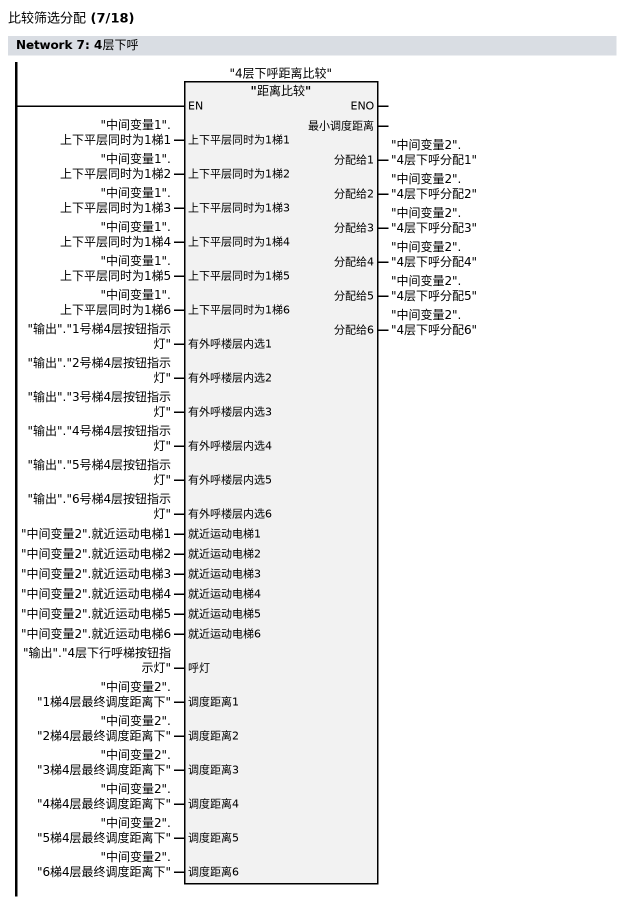
   RUNG wire#powerrail
      "4层下呼距离比较"(上下平层同时为1梯1 := "中间变量1".上下平层同时为1梯1, 上下平层同时为1梯2 := "中间变量1".上下平层同时为1梯2, 上下平层同时为1梯3 := "中间变量1".上下平层同时为1梯3, 上下平层同时为1梯4 := "中间变量1".上下平层同时为1梯4, 上下平层同时为1梯5 := "中间变量1".上下平层同时为1梯5, 上下平层同时为1梯6 := "中间变量1".上下平层同时为1梯6, 有外呼楼层内选1 := "输出"."1号梯4层按钮指示灯", 有外呼楼层内选2 := "输出"."2号梯4层按钮指示灯", 有外呼楼层内选3 := "输出"."3号梯4层按钮指示灯", 有外呼楼层内选4 := "输出"."4号梯4层按钮指示灯", 有外呼楼层内选5 := "输出"."5号梯4层按钮指示灯", 有外呼楼层内选6 := "输出"."6号梯4层按钮指示灯", 就近运动电梯1 := "中间变量2".就近运动电梯1, 就近运动电梯2 := "中间变量2".就近运动电梯2, 就近运动电梯3 := "中间变量2".就近运动电梯3, 就近运动电梯4 := "中间变量2".就近运动电梯4, 就近运动电梯5 := "中间变量2".就近运动电梯5, 就近运动电梯6 := "中间变量2".就近运动电梯6, 呼灯 := "输出"."4层下行呼梯按钮指示灯", 调度距离1 := "中间变量2"."1梯4层最终调度距离下", 调度距离2 := "中间变量2"."2梯4层最终调度距离下", 调度距离3 := "中间变量2"."3梯4层最终调度距离下", 调度距离4 := "中间变量2"."4梯4层最终调度距离下", 调度距离5 := "中间变量2"."5梯4层最终调度距离下", 调度距离6 := "中间变量2"."6梯4层最终调度距离下", 最小调度距离 =>, 分配给1 => "中间变量2"."4层下呼分配1", 分配给2 => "中间变量2"."4层下呼分配2", 分配给3 => "中间变量2"."4层下呼分配3", 分配给4 => "中间变量2"."4层下呼分配4", 分配给5 => "中间变量2"."4层下呼分配5", 分配给6 => "中间变量2"."4层下呼分配6")
   END_RUNG
   // the same network as SCL:
   "4层下呼距离比较"(上下平层同时为1梯1 := "中间变量1".上下平层同时为1梯1,   // "距离比较"
              上下平层同时为1梯2 := "中间变量1".上下平层同时为1梯2,
              上下平层同时为1梯3 := "中间变量1".上下平层同时为1梯3,
              上下平层同时为1梯4 := "中间变量1".上下平层同时为1梯4,
              上下平层同时为1梯5 := "中间变量1".上下平层同时为1梯5,
              上下平层同时为1梯6 := "中间变量1".上下平层同时为1梯6,
              有外呼楼层内选1 := "输出"."1号梯4层按钮指示灯",
              有外呼楼层内选2 := "输出"."2号梯4层按钮指示灯",
              有外呼楼层内选3 := "输出"."3号梯4层按钮指示灯",
              有外呼楼层内选4 := "输出"."4号梯4层按钮指示灯",
              有外呼楼层内选5 := "输出"."5号梯4层按钮指示灯",
              有外呼楼层内选6 := "输出"."6号梯4层按钮指示灯",
              就近运动电梯1 := "中间变量2".就近运动电梯1,
              就近运动电梯2 := "中间变量2".就近运动电梯2,
              就近运动电梯3 := "中间变量2".就近运动电梯3,
              就近运动电梯4 := "中间变量2".就近运动电梯4,
              就近运动电梯5 := "中间变量2".就近运动电梯5,
              就近运动电梯6 := "中间变量2".就近运动电梯6,
              呼灯 := "输出"."4层下行呼梯按钮指示灯",
              调度距离1 := "中间变量2"."1梯4层最终调度距离下",
              调度距离2 := "中间变量2"."2梯4层最终调度距离下",
              调度距离3 := "中间变量2"."3梯4层最终调度距离下",
              调度距离4 := "中间变量2"."4梯4层最终调度距离下",
              调度距离5 := "中间变量2"."5梯4层最终调度距离下",
              调度距离6 := "中间变量2"."6梯4层最终调度距离下",
              分配给1 => "中间变量2"."4层下呼分配1",
              分配给2 => "中间变量2"."4层下呼分配2",
              分配给3 => "中间变量2"."4层下呼分配3",
              分配给4 => "中间变量2"."4层下呼分配4",
              分配给5 => "中间变量2"."4层下呼分配5",
              分配给6 => "中间变量2"."4层下呼分配6");
END_REGION

REGION Network 8: 5层上呼
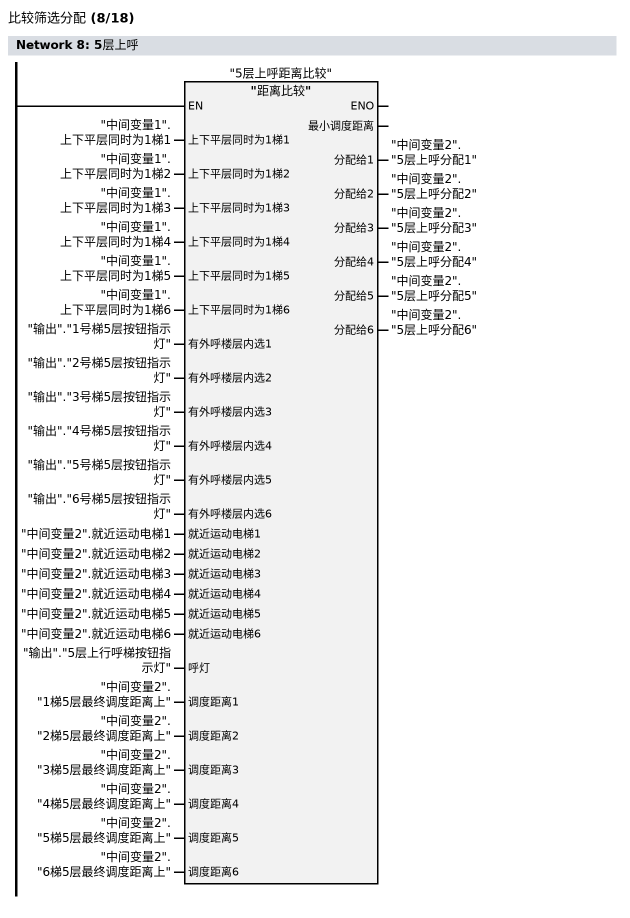
   RUNG wire#powerrail
      "5层上呼距离比较"(上下平层同时为1梯1 := "中间变量1".上下平层同时为1梯1, 上下平层同时为1梯2 := "中间变量1".上下平层同时为1梯2, 上下平层同时为1梯3 := "中间变量1".上下平层同时为1梯3, 上下平层同时为1梯4 := "中间变量1".上下平层同时为1梯4, 上下平层同时为1梯5 := "中间变量1".上下平层同时为1梯5, 上下平层同时为1梯6 := "中间变量1".上下平层同时为1梯6, 有外呼楼层内选1 := "输出"."1号梯5层按钮指示灯", 有外呼楼层内选2 := "输出"."2号梯5层按钮指示灯", 有外呼楼层内选3 := "输出"."3号梯5层按钮指示灯", 有外呼楼层内选4 := "输出"."4号梯5层按钮指示灯", 有外呼楼层内选5 := "输出"."5号梯5层按钮指示灯", 有外呼楼层内选6 := "输出"."6号梯5层按钮指示灯", 就近运动电梯1 := "中间变量2".就近运动电梯1, 就近运动电梯2 := "中间变量2".就近运动电梯2, 就近运动电梯3 := "中间变量2".就近运动电梯3, 就近运动电梯4 := "中间变量2".就近运动电梯4, 就近运动电梯5 := "中间变量2".就近运动电梯5, 就近运动电梯6 := "中间变量2".就近运动电梯6, 呼灯 := "输出"."5层上行呼梯按钮指示灯", 调度距离1 := "中间变量2"."1梯5层最终调度距离上", 调度距离2 := "中间变量2"."2梯5层最终调度距离上", 调度距离3 := "中间变量2"."3梯5层最终调度距离上", 调度距离4 := "中间变量2"."4梯5层最终调度距离上", 调度距离5 := "中间变量2"."5梯5层最终调度距离上", 调度距离6 := "中间变量2"."6梯5层最终调度距离上", 最小调度距离 =>, 分配给1 => "中间变量2"."5层上呼分配1", 分配给2 => "中间变量2"."5层上呼分配2", 分配给3 => "中间变量2"."5层上呼分配3", 分配给4 => "中间变量2"."5层上呼分配4", 分配给5 => "中间变量2"."5层上呼分配5", 分配给6 => "中间变量2"."5层上呼分配6")
   END_RUNG
   // the same network as SCL:
   "5层上呼距离比较"(上下平层同时为1梯1 := "中间变量1".上下平层同时为1梯1,   // "距离比较"
              上下平层同时为1梯2 := "中间变量1".上下平层同时为1梯2,
              上下平层同时为1梯3 := "中间变量1".上下平层同时为1梯3,
              上下平层同时为1梯4 := "中间变量1".上下平层同时为1梯4,
              上下平层同时为1梯5 := "中间变量1".上下平层同时为1梯5,
              上下平层同时为1梯6 := "中间变量1".上下平层同时为1梯6,
              有外呼楼层内选1 := "输出"."1号梯5层按钮指示灯",
              有外呼楼层内选2 := "输出"."2号梯5层按钮指示灯",
              有外呼楼层内选3 := "输出"."3号梯5层按钮指示灯",
              有外呼楼层内选4 := "输出"."4号梯5层按钮指示灯",
              有外呼楼层内选5 := "输出"."5号梯5层按钮指示灯",
              有外呼楼层内选6 := "输出"."6号梯5层按钮指示灯",
              就近运动电梯1 := "中间变量2".就近运动电梯1,
              就近运动电梯2 := "中间变量2".就近运动电梯2,
              就近运动电梯3 := "中间变量2".就近运动电梯3,
              就近运动电梯4 := "中间变量2".就近运动电梯4,
              就近运动电梯5 := "中间变量2".就近运动电梯5,
              就近运动电梯6 := "中间变量2".就近运动电梯6,
              呼灯 := "输出"."5层上行呼梯按钮指示灯",
              调度距离1 := "中间变量2"."1梯5层最终调度距离上",
              调度距离2 := "中间变量2"."2梯5层最终调度距离上",
              调度距离3 := "中间变量2"."3梯5层最终调度距离上",
              调度距离4 := "中间变量2"."4梯5层最终调度距离上",
              调度距离5 := "中间变量2"."5梯5层最终调度距离上",
              调度距离6 := "中间变量2"."6梯5层最终调度距离上",
              分配给1 => "中间变量2"."5层上呼分配1",
              分配给2 => "中间变量2"."5层上呼分配2",
              分配给3 => "中间变量2"."5层上呼分配3",
              分配给4 => "中间变量2"."5层上呼分配4",
              分配给5 => "中间变量2"."5层上呼分配5",
              分配给6 => "中间变量2"."5层上呼分配6");
END_REGION

REGION Network 9: 5层下呼
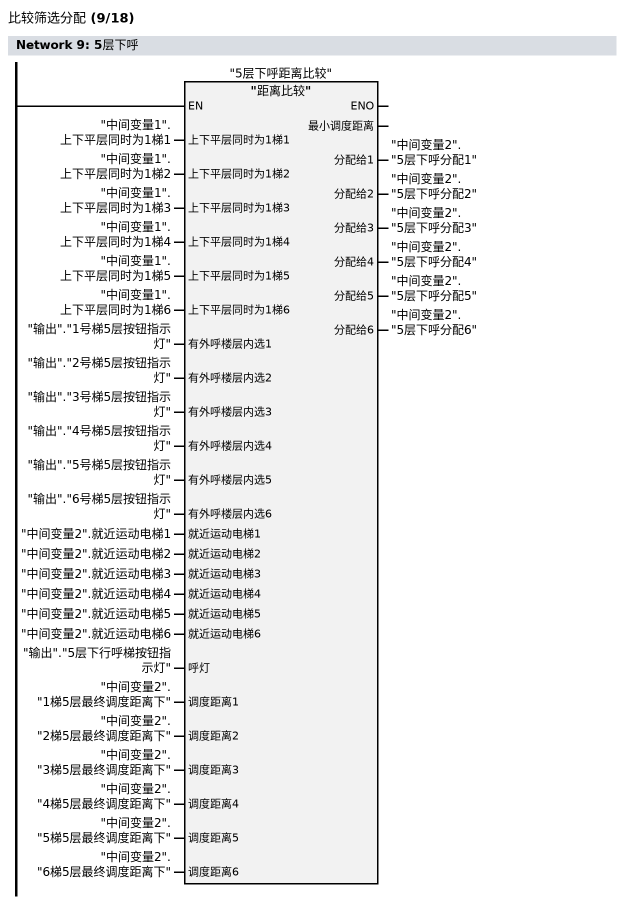
   RUNG wire#powerrail
      "5层下呼距离比较"(上下平层同时为1梯1 := "中间变量1".上下平层同时为1梯1, 上下平层同时为1梯2 := "中间变量1".上下平层同时为1梯2, 上下平层同时为1梯3 := "中间变量1".上下平层同时为1梯3, 上下平层同时为1梯4 := "中间变量1".上下平层同时为1梯4, 上下平层同时为1梯5 := "中间变量1".上下平层同时为1梯5, 上下平层同时为1梯6 := "中间变量1".上下平层同时为1梯6, 有外呼楼层内选1 := "输出"."1号梯5层按钮指示灯", 有外呼楼层内选2 := "输出"."2号梯5层按钮指示灯", 有外呼楼层内选3 := "输出"."3号梯5层按钮指示灯", 有外呼楼层内选4 := "输出"."4号梯5层按钮指示灯", 有外呼楼层内选5 := "输出"."5号梯5层按钮指示灯", 有外呼楼层内选6 := "输出"."6号梯5层按钮指示灯", 就近运动电梯1 := "中间变量2".就近运动电梯1, 就近运动电梯2 := "中间变量2".就近运动电梯2, 就近运动电梯3 := "中间变量2".就近运动电梯3, 就近运动电梯4 := "中间变量2".就近运动电梯4, 就近运动电梯5 := "中间变量2".就近运动电梯5, 就近运动电梯6 := "中间变量2".就近运动电梯6, 呼灯 := "输出"."5层下行呼梯按钮指示灯", 调度距离1 := "中间变量2"."1梯5层最终调度距离下", 调度距离2 := "中间变量2"."2梯5层最终调度距离下", 调度距离3 := "中间变量2"."3梯5层最终调度距离下", 调度距离4 := "中间变量2"."4梯5层最终调度距离下", 调度距离5 := "中间变量2"."5梯5层最终调度距离下", 调度距离6 := "中间变量2"."6梯5层最终调度距离下", 最小调度距离 =>, 分配给1 => "中间变量2"."5层下呼分配1", 分配给2 => "中间变量2"."5层下呼分配2", 分配给3 => "中间变量2"."5层下呼分配3", 分配给4 => "中间变量2"."5层下呼分配4", 分配给5 => "中间变量2"."5层下呼分配5", 分配给6 => "中间变量2"."5层下呼分配6")
   END_RUNG
   // the same network as SCL:
   "5层下呼距离比较"(上下平层同时为1梯1 := "中间变量1".上下平层同时为1梯1,   // "距离比较"
              上下平层同时为1梯2 := "中间变量1".上下平层同时为1梯2,
              上下平层同时为1梯3 := "中间变量1".上下平层同时为1梯3,
              上下平层同时为1梯4 := "中间变量1".上下平层同时为1梯4,
              上下平层同时为1梯5 := "中间变量1".上下平层同时为1梯5,
              上下平层同时为1梯6 := "中间变量1".上下平层同时为1梯6,
              有外呼楼层内选1 := "输出"."1号梯5层按钮指示灯",
              有外呼楼层内选2 := "输出"."2号梯5层按钮指示灯",
              有外呼楼层内选3 := "输出"."3号梯5层按钮指示灯",
              有外呼楼层内选4 := "输出"."4号梯5层按钮指示灯",
              有外呼楼层内选5 := "输出"."5号梯5层按钮指示灯",
              有外呼楼层内选6 := "输出"."6号梯5层按钮指示灯",
              就近运动电梯1 := "中间变量2".就近运动电梯1,
              就近运动电梯2 := "中间变量2".就近运动电梯2,
              就近运动电梯3 := "中间变量2".就近运动电梯3,
              就近运动电梯4 := "中间变量2".就近运动电梯4,
              就近运动电梯5 := "中间变量2".就近运动电梯5,
              就近运动电梯6 := "中间变量2".就近运动电梯6,
              呼灯 := "输出"."5层下行呼梯按钮指示灯",
              调度距离1 := "中间变量2"."1梯5层最终调度距离下",
              调度距离2 := "中间变量2"."2梯5层最终调度距离下",
              调度距离3 := "中间变量2"."3梯5层最终调度距离下",
              调度距离4 := "中间变量2"."4梯5层最终调度距离下",
              调度距离5 := "中间变量2"."5梯5层最终调度距离下",
              调度距离6 := "中间变量2"."6梯5层最终调度距离下",
              分配给1 => "中间变量2"."5层下呼分配1",
              分配给2 => "中间变量2"."5层下呼分配2",
              分配给3 => "中间变量2"."5层下呼分配3",
              分配给4 => "中间变量2"."5层下呼分配4",
              分配给5 => "中间变量2"."5层下呼分配5",
              分配给6 => "中间变量2"."5层下呼分配6");
END_REGION

REGION Network 10: 6层上呼
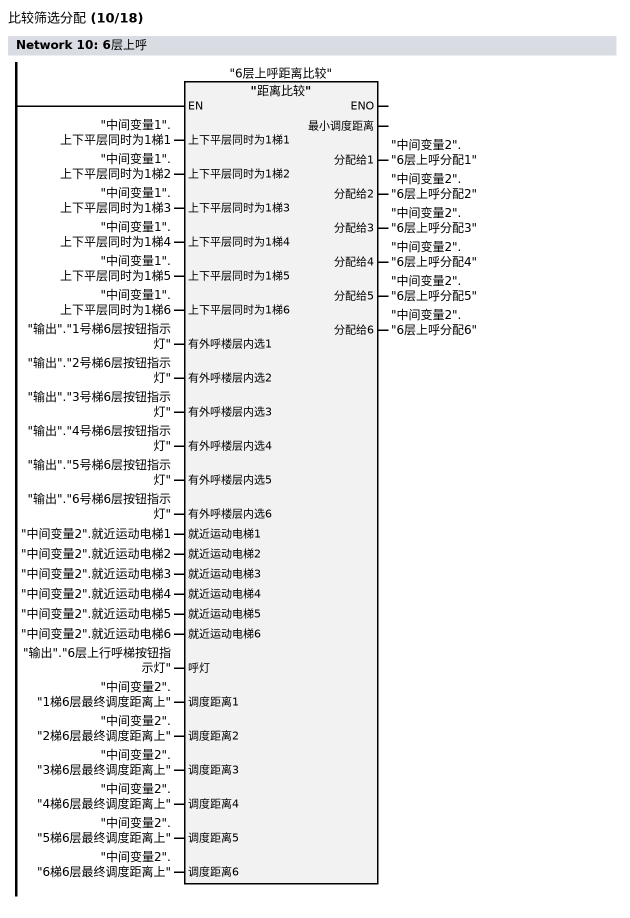
   RUNG wire#powerrail
      "6层上呼距离比较"(上下平层同时为1梯1 := "中间变量1".上下平层同时为1梯1, 上下平层同时为1梯2 := "中间变量1".上下平层同时为1梯2, 上下平层同时为1梯3 := "中间变量1".上下平层同时为1梯3, 上下平层同时为1梯4 := "中间变量1".上下平层同时为1梯4, 上下平层同时为1梯5 := "中间变量1".上下平层同时为1梯5, 上下平层同时为1梯6 := "中间变量1".上下平层同时为1梯6, 有外呼楼层内选1 := "输出"."1号梯6层按钮指示灯", 有外呼楼层内选2 := "输出"."2号梯6层按钮指示灯", 有外呼楼层内选3 := "输出"."3号梯6层按钮指示灯", 有外呼楼层内选4 := "输出"."4号梯6层按钮指示灯", 有外呼楼层内选5 := "输出"."5号梯6层按钮指示灯", 有外呼楼层内选6 := "输出"."6号梯6层按钮指示灯", 就近运动电梯1 := "中间变量2".就近运动电梯1, 就近运动电梯2 := "中间变量2".就近运动电梯2, 就近运动电梯3 := "中间变量2".就近运动电梯3, 就近运动电梯4 := "中间变量2".就近运动电梯4, 就近运动电梯5 := "中间变量2".就近运动电梯5, 就近运动电梯6 := "中间变量2".就近运动电梯6, 呼灯 := "输出"."6层上行呼梯按钮指示灯", 调度距离1 := "中间变量2"."1梯6层最终调度距离上", 调度距离2 := "中间变量2"."2梯6层最终调度距离上", 调度距离3 := "中间变量2"."3梯6层最终调度距离上", 调度距离4 := "中间变量2"."4梯6层最终调度距离上", 调度距离5 := "中间变量2"."5梯6层最终调度距离上", 调度距离6 := "中间变量2"."6梯6层最终调度距离上", 最小调度距离 =>, 分配给1 => "中间变量2"."6层上呼分配1", 分配给2 => "中间变量2"."6层上呼分配2", 分配给3 => "中间变量2"."6层上呼分配3", 分配给4 => "中间变量2"."6层上呼分配4", 分配给5 => "中间变量2"."6层上呼分配5", 分配给6 => "中间变量2"."6层上呼分配6")
   END_RUNG
   // the same network as SCL:
   "6层上呼距离比较"(上下平层同时为1梯1 := "中间变量1".上下平层同时为1梯1,   // "距离比较"
              上下平层同时为1梯2 := "中间变量1".上下平层同时为1梯2,
              上下平层同时为1梯3 := "中间变量1".上下平层同时为1梯3,
              上下平层同时为1梯4 := "中间变量1".上下平层同时为1梯4,
              上下平层同时为1梯5 := "中间变量1".上下平层同时为1梯5,
              上下平层同时为1梯6 := "中间变量1".上下平层同时为1梯6,
              有外呼楼层内选1 := "输出"."1号梯6层按钮指示灯",
              有外呼楼层内选2 := "输出"."2号梯6层按钮指示灯",
              有外呼楼层内选3 := "输出"."3号梯6层按钮指示灯",
              有外呼楼层内选4 := "输出"."4号梯6层按钮指示灯",
              有外呼楼层内选5 := "输出"."5号梯6层按钮指示灯",
              有外呼楼层内选6 := "输出"."6号梯6层按钮指示灯",
              就近运动电梯1 := "中间变量2".就近运动电梯1,
              就近运动电梯2 := "中间变量2".就近运动电梯2,
              就近运动电梯3 := "中间变量2".就近运动电梯3,
              就近运动电梯4 := "中间变量2".就近运动电梯4,
              就近运动电梯5 := "中间变量2".就近运动电梯5,
              就近运动电梯6 := "中间变量2".就近运动电梯6,
              呼灯 := "输出"."6层上行呼梯按钮指示灯",
              调度距离1 := "中间变量2"."1梯6层最终调度距离上",
              调度距离2 := "中间变量2"."2梯6层最终调度距离上",
              调度距离3 := "中间变量2"."3梯6层最终调度距离上",
              调度距离4 := "中间变量2"."4梯6层最终调度距离上",
              调度距离5 := "中间变量2"."5梯6层最终调度距离上",
              调度距离6 := "中间变量2"."6梯6层最终调度距离上",
              分配给1 => "中间变量2"."6层上呼分配1",
              分配给2 => "中间变量2"."6层上呼分配2",
              分配给3 => "中间变量2"."6层上呼分配3",
              分配给4 => "中间变量2"."6层上呼分配4",
              分配给5 => "中间变量2"."6层上呼分配5",
              分配给6 => "中间变量2"."6层上呼分配6");
END_REGION

REGION Network 11: 6层下呼
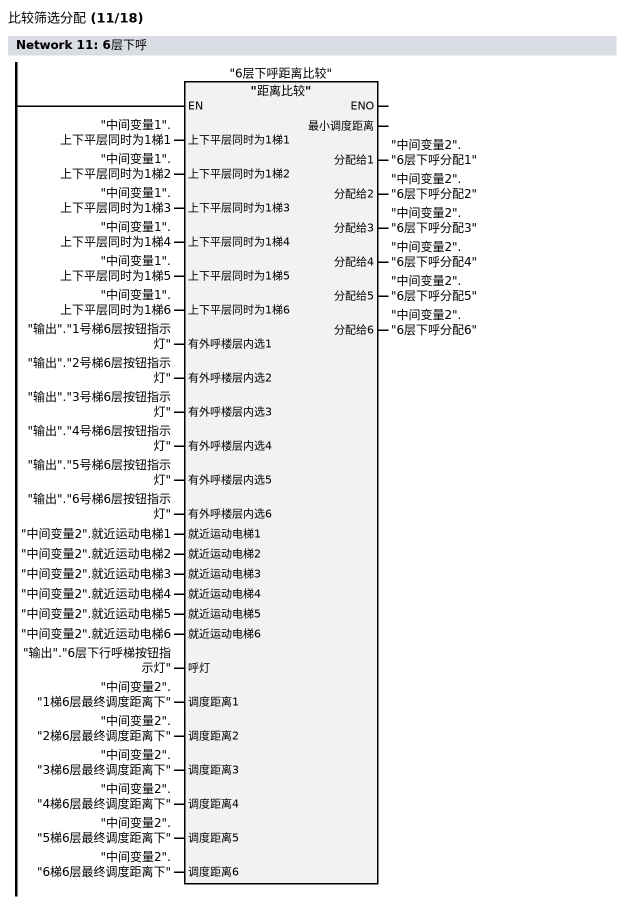
   RUNG wire#powerrail
      "6层下呼距离比较"(上下平层同时为1梯1 := "中间变量1".上下平层同时为1梯1, 上下平层同时为1梯2 := "中间变量1".上下平层同时为1梯2, 上下平层同时为1梯3 := "中间变量1".上下平层同时为1梯3, 上下平层同时为1梯4 := "中间变量1".上下平层同时为1梯4, 上下平层同时为1梯5 := "中间变量1".上下平层同时为1梯5, 上下平层同时为1梯6 := "中间变量1".上下平层同时为1梯6, 有外呼楼层内选1 := "输出"."1号梯6层按钮指示灯", 有外呼楼层内选2 := "输出"."2号梯6层按钮指示灯", 有外呼楼层内选3 := "输出"."3号梯6层按钮指示灯", 有外呼楼层内选4 := "输出"."4号梯6层按钮指示灯", 有外呼楼层内选5 := "输出"."5号梯6层按钮指示灯", 有外呼楼层内选6 := "输出"."6号梯6层按钮指示灯", 就近运动电梯1 := "中间变量2".就近运动电梯1, 就近运动电梯2 := "中间变量2".就近运动电梯2, 就近运动电梯3 := "中间变量2".就近运动电梯3, 就近运动电梯4 := "中间变量2".就近运动电梯4, 就近运动电梯5 := "中间变量2".就近运动电梯5, 就近运动电梯6 := "中间变量2".就近运动电梯6, 呼灯 := "输出"."6层下行呼梯按钮指示灯", 调度距离1 := "中间变量2"."1梯6层最终调度距离下", 调度距离2 := "中间变量2"."2梯6层最终调度距离下", 调度距离3 := "中间变量2"."3梯6层最终调度距离下", 调度距离4 := "中间变量2"."4梯6层最终调度距离下", 调度距离5 := "中间变量2"."5梯6层最终调度距离下", 调度距离6 := "中间变量2"."6梯6层最终调度距离下", 最小调度距离 =>, 分配给1 => "中间变量2"."6层下呼分配1", 分配给2 => "中间变量2"."6层下呼分配2", 分配给3 => "中间变量2"."6层下呼分配3", 分配给4 => "中间变量2"."6层下呼分配4", 分配给5 => "中间变量2"."6层下呼分配5", 分配给6 => "中间变量2"."6层下呼分配6")
   END_RUNG
   // the same network as SCL:
   "6层下呼距离比较"(上下平层同时为1梯1 := "中间变量1".上下平层同时为1梯1,   // "距离比较"
              上下平层同时为1梯2 := "中间变量1".上下平层同时为1梯2,
              上下平层同时为1梯3 := "中间变量1".上下平层同时为1梯3,
              上下平层同时为1梯4 := "中间变量1".上下平层同时为1梯4,
              上下平层同时为1梯5 := "中间变量1".上下平层同时为1梯5,
              上下平层同时为1梯6 := "中间变量1".上下平层同时为1梯6,
              有外呼楼层内选1 := "输出"."1号梯6层按钮指示灯",
              有外呼楼层内选2 := "输出"."2号梯6层按钮指示灯",
              有外呼楼层内选3 := "输出"."3号梯6层按钮指示灯",
              有外呼楼层内选4 := "输出"."4号梯6层按钮指示灯",
              有外呼楼层内选5 := "输出"."5号梯6层按钮指示灯",
              有外呼楼层内选6 := "输出"."6号梯6层按钮指示灯",
              就近运动电梯1 := "中间变量2".就近运动电梯1,
              就近运动电梯2 := "中间变量2".就近运动电梯2,
              就近运动电梯3 := "中间变量2".就近运动电梯3,
              就近运动电梯4 := "中间变量2".就近运动电梯4,
              就近运动电梯5 := "中间变量2".就近运动电梯5,
              就近运动电梯6 := "中间变量2".就近运动电梯6,
              呼灯 := "输出"."6层下行呼梯按钮指示灯",
              调度距离1 := "中间变量2"."1梯6层最终调度距离下",
              调度距离2 := "中间变量2"."2梯6层最终调度距离下",
              调度距离3 := "中间变量2"."3梯6层最终调度距离下",
              调度距离4 := "中间变量2"."4梯6层最终调度距离下",
              调度距离5 := "中间变量2"."5梯6层最终调度距离下",
              调度距离6 := "中间变量2"."6梯6层最终调度距离下",
              分配给1 => "中间变量2"."6层下呼分配1",
              分配给2 => "中间变量2"."6层下呼分配2",
              分配给3 => "中间变量2"."6层下呼分配3",
              分配给4 => "中间变量2"."6层下呼分配4",
              分配给5 => "中间变量2"."6层下呼分配5",
              分配给6 => "中间变量2"."6层下呼分配6");
END_REGION

REGION Network 12: 7层上呼
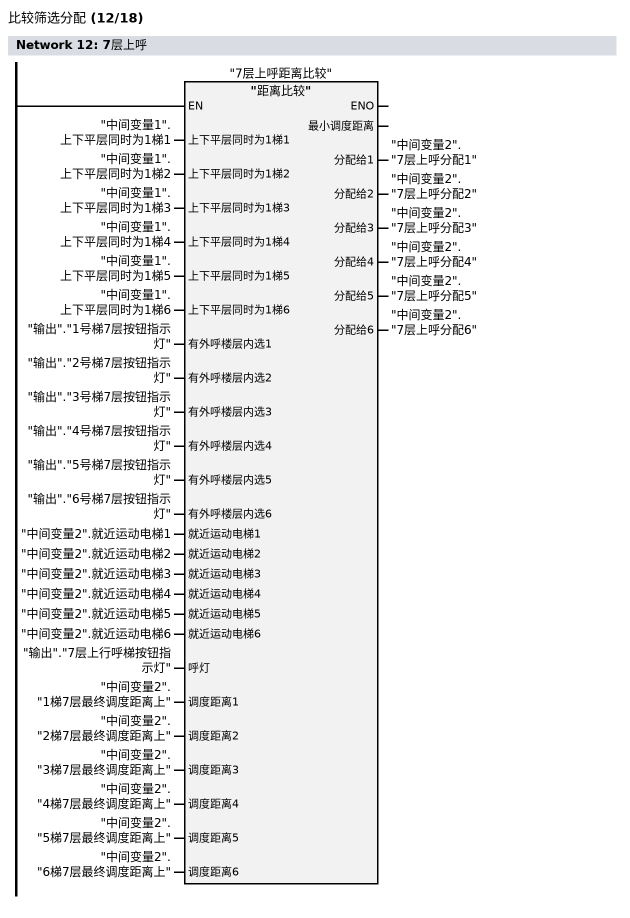
   RUNG wire#powerrail
      "7层上呼距离比较"(上下平层同时为1梯1 := "中间变量1".上下平层同时为1梯1, 上下平层同时为1梯2 := "中间变量1".上下平层同时为1梯2, 上下平层同时为1梯3 := "中间变量1".上下平层同时为1梯3, 上下平层同时为1梯4 := "中间变量1".上下平层同时为1梯4, 上下平层同时为1梯5 := "中间变量1".上下平层同时为1梯5, 上下平层同时为1梯6 := "中间变量1".上下平层同时为1梯6, 有外呼楼层内选1 := "输出"."1号梯7层按钮指示灯", 有外呼楼层内选2 := "输出"."2号梯7层按钮指示灯", 有外呼楼层内选3 := "输出"."3号梯7层按钮指示灯", 有外呼楼层内选4 := "输出"."4号梯7层按钮指示灯", 有外呼楼层内选5 := "输出"."5号梯7层按钮指示灯", 有外呼楼层内选6 := "输出"."6号梯7层按钮指示灯", 就近运动电梯1 := "中间变量2".就近运动电梯1, 就近运动电梯2 := "中间变量2".就近运动电梯2, 就近运动电梯3 := "中间变量2".就近运动电梯3, 就近运动电梯4 := "中间变量2".就近运动电梯4, 就近运动电梯5 := "中间变量2".就近运动电梯5, 就近运动电梯6 := "中间变量2".就近运动电梯6, 呼灯 := "输出"."7层上行呼梯按钮指示灯", 调度距离1 := "中间变量2"."1梯7层最终调度距离上", 调度距离2 := "中间变量2"."2梯7层最终调度距离上", 调度距离3 := "中间变量2"."3梯7层最终调度距离上", 调度距离4 := "中间变量2"."4梯7层最终调度距离上", 调度距离5 := "中间变量2"."5梯7层最终调度距离上", 调度距离6 := "中间变量2"."6梯7层最终调度距离上", 最小调度距离 =>, 分配给1 => "中间变量2"."7层上呼分配1", 分配给2 => "中间变量2"."7层上呼分配2", 分配给3 => "中间变量2"."7层上呼分配3", 分配给4 => "中间变量2"."7层上呼分配4", 分配给5 => "中间变量2"."7层上呼分配5", 分配给6 => "中间变量2"."7层上呼分配6")
   END_RUNG
   // the same network as SCL:
   "7层上呼距离比较"(上下平层同时为1梯1 := "中间变量1".上下平层同时为1梯1,   // "距离比较"
              上下平层同时为1梯2 := "中间变量1".上下平层同时为1梯2,
              上下平层同时为1梯3 := "中间变量1".上下平层同时为1梯3,
              上下平层同时为1梯4 := "中间变量1".上下平层同时为1梯4,
              上下平层同时为1梯5 := "中间变量1".上下平层同时为1梯5,
              上下平层同时为1梯6 := "中间变量1".上下平层同时为1梯6,
              有外呼楼层内选1 := "输出"."1号梯7层按钮指示灯",
              有外呼楼层内选2 := "输出"."2号梯7层按钮指示灯",
              有外呼楼层内选3 := "输出"."3号梯7层按钮指示灯",
              有外呼楼层内选4 := "输出"."4号梯7层按钮指示灯",
              有外呼楼层内选5 := "输出"."5号梯7层按钮指示灯",
              有外呼楼层内选6 := "输出"."6号梯7层按钮指示灯",
              就近运动电梯1 := "中间变量2".就近运动电梯1,
              就近运动电梯2 := "中间变量2".就近运动电梯2,
              就近运动电梯3 := "中间变量2".就近运动电梯3,
              就近运动电梯4 := "中间变量2".就近运动电梯4,
              就近运动电梯5 := "中间变量2".就近运动电梯5,
              就近运动电梯6 := "中间变量2".就近运动电梯6,
              呼灯 := "输出"."7层上行呼梯按钮指示灯",
              调度距离1 := "中间变量2"."1梯7层最终调度距离上",
              调度距离2 := "中间变量2"."2梯7层最终调度距离上",
              调度距离3 := "中间变量2"."3梯7层最终调度距离上",
              调度距离4 := "中间变量2"."4梯7层最终调度距离上",
              调度距离5 := "中间变量2"."5梯7层最终调度距离上",
              调度距离6 := "中间变量2"."6梯7层最终调度距离上",
              分配给1 => "中间变量2"."7层上呼分配1",
              分配给2 => "中间变量2"."7层上呼分配2",
              分配给3 => "中间变量2"."7层上呼分配3",
              分配给4 => "中间变量2"."7层上呼分配4",
              分配给5 => "中间变量2"."7层上呼分配5",
              分配给6 => "中间变量2"."7层上呼分配6");
END_REGION

REGION Network 13: 7层下呼
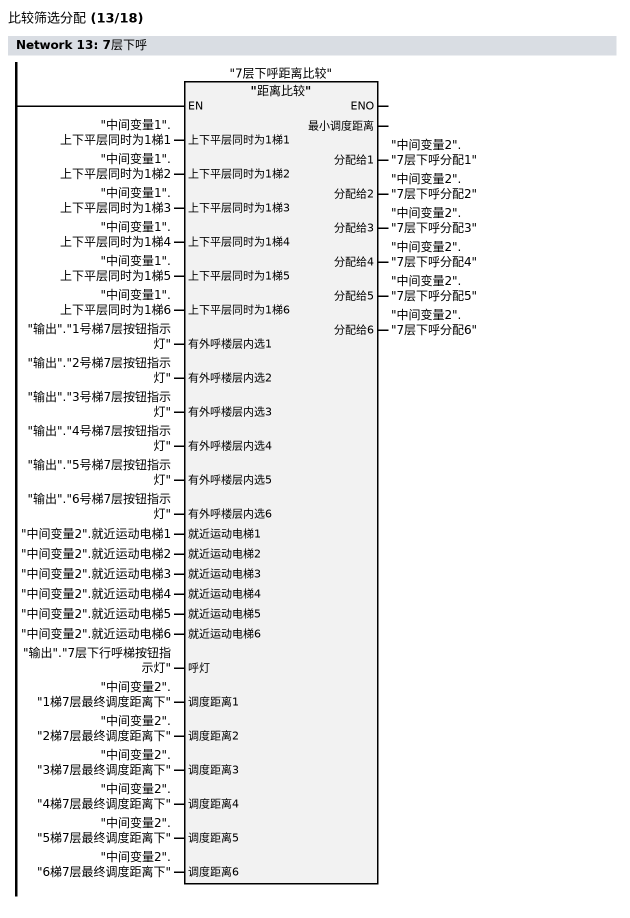
   RUNG wire#powerrail
      "7层下呼距离比较"(上下平层同时为1梯1 := "中间变量1".上下平层同时为1梯1, 上下平层同时为1梯2 := "中间变量1".上下平层同时为1梯2, 上下平层同时为1梯3 := "中间变量1".上下平层同时为1梯3, 上下平层同时为1梯4 := "中间变量1".上下平层同时为1梯4, 上下平层同时为1梯5 := "中间变量1".上下平层同时为1梯5, 上下平层同时为1梯6 := "中间变量1".上下平层同时为1梯6, 有外呼楼层内选1 := "输出"."1号梯7层按钮指示灯", 有外呼楼层内选2 := "输出"."2号梯7层按钮指示灯", 有外呼楼层内选3 := "输出"."3号梯7层按钮指示灯", 有外呼楼层内选4 := "输出"."4号梯7层按钮指示灯", 有外呼楼层内选5 := "输出"."5号梯7层按钮指示灯", 有外呼楼层内选6 := "输出"."6号梯7层按钮指示灯", 就近运动电梯1 := "中间变量2".就近运动电梯1, 就近运动电梯2 := "中间变量2".就近运动电梯2, 就近运动电梯3 := "中间变量2".就近运动电梯3, 就近运动电梯4 := "中间变量2".就近运动电梯4, 就近运动电梯5 := "中间变量2".就近运动电梯5, 就近运动电梯6 := "中间变量2".就近运动电梯6, 呼灯 := "输出"."7层下行呼梯按钮指示灯", 调度距离1 := "中间变量2"."1梯7层最终调度距离下", 调度距离2 := "中间变量2"."2梯7层最终调度距离下", 调度距离3 := "中间变量2"."3梯7层最终调度距离下", 调度距离4 := "中间变量2"."4梯7层最终调度距离下", 调度距离5 := "中间变量2"."5梯7层最终调度距离下", 调度距离6 := "中间变量2"."6梯7层最终调度距离下", 最小调度距离 =>, 分配给1 => "中间变量2"."7层下呼分配1", 分配给2 => "中间变量2"."7层下呼分配2", 分配给3 => "中间变量2"."7层下呼分配3", 分配给4 => "中间变量2"."7层下呼分配4", 分配给5 => "中间变量2"."7层下呼分配5", 分配给6 => "中间变量2"."7层下呼分配6")
   END_RUNG
   // the same network as SCL:
   "7层下呼距离比较"(上下平层同时为1梯1 := "中间变量1".上下平层同时为1梯1,   // "距离比较"
              上下平层同时为1梯2 := "中间变量1".上下平层同时为1梯2,
              上下平层同时为1梯3 := "中间变量1".上下平层同时为1梯3,
              上下平层同时为1梯4 := "中间变量1".上下平层同时为1梯4,
              上下平层同时为1梯5 := "中间变量1".上下平层同时为1梯5,
              上下平层同时为1梯6 := "中间变量1".上下平层同时为1梯6,
              有外呼楼层内选1 := "输出"."1号梯7层按钮指示灯",
              有外呼楼层内选2 := "输出"."2号梯7层按钮指示灯",
              有外呼楼层内选3 := "输出"."3号梯7层按钮指示灯",
              有外呼楼层内选4 := "输出"."4号梯7层按钮指示灯",
              有外呼楼层内选5 := "输出"."5号梯7层按钮指示灯",
              有外呼楼层内选6 := "输出"."6号梯7层按钮指示灯",
              就近运动电梯1 := "中间变量2".就近运动电梯1,
              就近运动电梯2 := "中间变量2".就近运动电梯2,
              就近运动电梯3 := "中间变量2".就近运动电梯3,
              就近运动电梯4 := "中间变量2".就近运动电梯4,
              就近运动电梯5 := "中间变量2".就近运动电梯5,
              就近运动电梯6 := "中间变量2".就近运动电梯6,
              呼灯 := "输出"."7层下行呼梯按钮指示灯",
              调度距离1 := "中间变量2"."1梯7层最终调度距离下",
              调度距离2 := "中间变量2"."2梯7层最终调度距离下",
              调度距离3 := "中间变量2"."3梯7层最终调度距离下",
              调度距离4 := "中间变量2"."4梯7层最终调度距离下",
              调度距离5 := "中间变量2"."5梯7层最终调度距离下",
              调度距离6 := "中间变量2"."6梯7层最终调度距离下",
              分配给1 => "中间变量2"."7层下呼分配1",
              分配给2 => "中间变量2"."7层下呼分配2",
              分配给3 => "中间变量2"."7层下呼分配3",
              分配给4 => "中间变量2"."7层下呼分配4",
              分配给5 => "中间变量2"."7层下呼分配5",
              分配给6 => "中间变量2"."7层下呼分配6");
END_REGION

REGION Network 14: 8层上呼
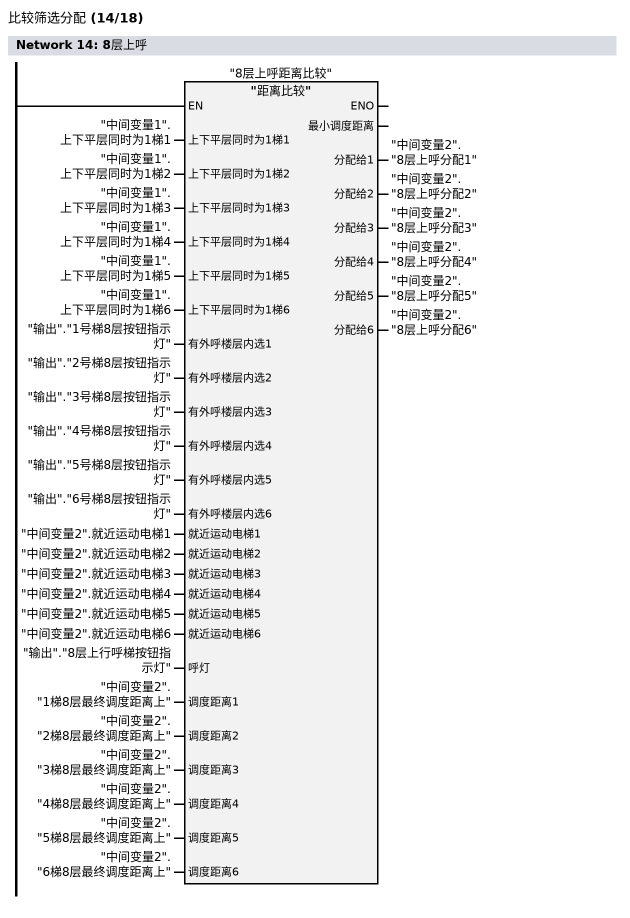
   RUNG wire#powerrail
      "8层上呼距离比较"(上下平层同时为1梯1 := "中间变量1".上下平层同时为1梯1, 上下平层同时为1梯2 := "中间变量1".上下平层同时为1梯2, 上下平层同时为1梯3 := "中间变量1".上下平层同时为1梯3, 上下平层同时为1梯4 := "中间变量1".上下平层同时为1梯4, 上下平层同时为1梯5 := "中间变量1".上下平层同时为1梯5, 上下平层同时为1梯6 := "中间变量1".上下平层同时为1梯6, 有外呼楼层内选1 := "输出"."1号梯8层按钮指示灯", 有外呼楼层内选2 := "输出"."2号梯8层按钮指示灯", 有外呼楼层内选3 := "输出"."3号梯8层按钮指示灯", 有外呼楼层内选4 := "输出"."4号梯8层按钮指示灯", 有外呼楼层内选5 := "输出"."5号梯8层按钮指示灯", 有外呼楼层内选6 := "输出"."6号梯8层按钮指示灯", 就近运动电梯1 := "中间变量2".就近运动电梯1, 就近运动电梯2 := "中间变量2".就近运动电梯2, 就近运动电梯3 := "中间变量2".就近运动电梯3, 就近运动电梯4 := "中间变量2".就近运动电梯4, 就近运动电梯5 := "中间变量2".就近运动电梯5, 就近运动电梯6 := "中间变量2".就近运动电梯6, 呼灯 := "输出"."8层上行呼梯按钮指示灯", 调度距离1 := "中间变量2"."1梯8层最终调度距离上", 调度距离2 := "中间变量2"."2梯8层最终调度距离上", 调度距离3 := "中间变量2"."3梯8层最终调度距离上", 调度距离4 := "中间变量2"."4梯8层最终调度距离上", 调度距离5 := "中间变量2"."5梯8层最终调度距离上", 调度距离6 := "中间变量2"."6梯8层最终调度距离上", 最小调度距离 =>, 分配给1 => "中间变量2"."8层上呼分配1", 分配给2 => "中间变量2"."8层上呼分配2", 分配给3 => "中间变量2"."8层上呼分配3", 分配给4 => "中间变量2"."8层上呼分配4", 分配给5 => "中间变量2"."8层上呼分配5", 分配给6 => "中间变量2"."8层上呼分配6")
   END_RUNG
   // the same network as SCL:
   "8层上呼距离比较"(上下平层同时为1梯1 := "中间变量1".上下平层同时为1梯1,   // "距离比较"
              上下平层同时为1梯2 := "中间变量1".上下平层同时为1梯2,
              上下平层同时为1梯3 := "中间变量1".上下平层同时为1梯3,
              上下平层同时为1梯4 := "中间变量1".上下平层同时为1梯4,
              上下平层同时为1梯5 := "中间变量1".上下平层同时为1梯5,
              上下平层同时为1梯6 := "中间变量1".上下平层同时为1梯6,
              有外呼楼层内选1 := "输出"."1号梯8层按钮指示灯",
              有外呼楼层内选2 := "输出"."2号梯8层按钮指示灯",
              有外呼楼层内选3 := "输出"."3号梯8层按钮指示灯",
              有外呼楼层内选4 := "输出"."4号梯8层按钮指示灯",
              有外呼楼层内选5 := "输出"."5号梯8层按钮指示灯",
              有外呼楼层内选6 := "输出"."6号梯8层按钮指示灯",
              就近运动电梯1 := "中间变量2".就近运动电梯1,
              就近运动电梯2 := "中间变量2".就近运动电梯2,
              就近运动电梯3 := "中间变量2".就近运动电梯3,
              就近运动电梯4 := "中间变量2".就近运动电梯4,
              就近运动电梯5 := "中间变量2".就近运动电梯5,
              就近运动电梯6 := "中间变量2".就近运动电梯6,
              呼灯 := "输出"."8层上行呼梯按钮指示灯",
              调度距离1 := "中间变量2"."1梯8层最终调度距离上",
              调度距离2 := "中间变量2"."2梯8层最终调度距离上",
              调度距离3 := "中间变量2"."3梯8层最终调度距离上",
              调度距离4 := "中间变量2"."4梯8层最终调度距离上",
              调度距离5 := "中间变量2"."5梯8层最终调度距离上",
              调度距离6 := "中间变量2"."6梯8层最终调度距离上",
              分配给1 => "中间变量2"."8层上呼分配1",
              分配给2 => "中间变量2"."8层上呼分配2",
              分配给3 => "中间变量2"."8层上呼分配3",
              分配给4 => "中间变量2"."8层上呼分配4",
              分配给5 => "中间变量2"."8层上呼分配5",
              分配给6 => "中间变量2"."8层上呼分配6");
END_REGION

REGION Network 15: 8层下呼
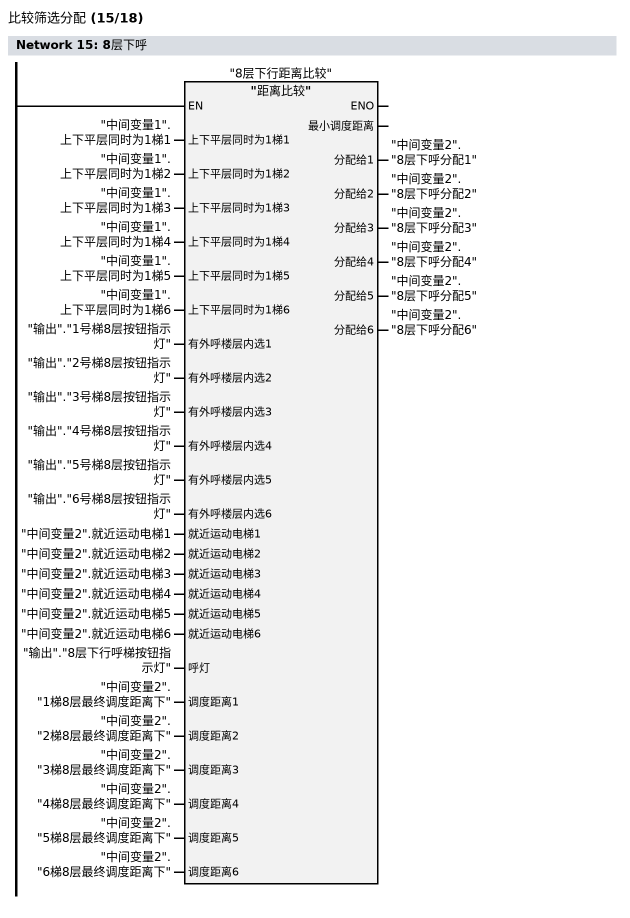
   RUNG wire#powerrail
      "8层下行距离比较"(上下平层同时为1梯1 := "中间变量1".上下平层同时为1梯1, 上下平层同时为1梯2 := "中间变量1".上下平层同时为1梯2, 上下平层同时为1梯3 := "中间变量1".上下平层同时为1梯3, 上下平层同时为1梯4 := "中间变量1".上下平层同时为1梯4, 上下平层同时为1梯5 := "中间变量1".上下平层同时为1梯5, 上下平层同时为1梯6 := "中间变量1".上下平层同时为1梯6, 有外呼楼层内选1 := "输出"."1号梯8层按钮指示灯", 有外呼楼层内选2 := "输出"."2号梯8层按钮指示灯", 有外呼楼层内选3 := "输出"."3号梯8层按钮指示灯", 有外呼楼层内选4 := "输出"."4号梯8层按钮指示灯", 有外呼楼层内选5 := "输出"."5号梯8层按钮指示灯", 有外呼楼层内选6 := "输出"."6号梯8层按钮指示灯", 就近运动电梯1 := "中间变量2".就近运动电梯1, 就近运动电梯2 := "中间变量2".就近运动电梯2, 就近运动电梯3 := "中间变量2".就近运动电梯3, 就近运动电梯4 := "中间变量2".就近运动电梯4, 就近运动电梯5 := "中间变量2".就近运动电梯5, 就近运动电梯6 := "中间变量2".就近运动电梯6, 呼灯 := "输出"."8层下行呼梯按钮指示灯", 调度距离1 := "中间变量2"."1梯8层最终调度距离下", 调度距离2 := "中间变量2"."2梯8层最终调度距离下", 调度距离3 := "中间变量2"."3梯8层最终调度距离下", 调度距离4 := "中间变量2"."4梯8层最终调度距离下", 调度距离5 := "中间变量2"."5梯8层最终调度距离下", 调度距离6 := "中间变量2"."6梯8层最终调度距离下", 最小调度距离 =>, 分配给1 => "中间变量2"."8层下呼分配1", 分配给2 => "中间变量2"."8层下呼分配2", 分配给3 => "中间变量2"."8层下呼分配3", 分配给4 => "中间变量2"."8层下呼分配4", 分配给5 => "中间变量2"."8层下呼分配5", 分配给6 => "中间变量2"."8层下呼分配6")
   END_RUNG
   // the same network as SCL:
   "8层下行距离比较"(上下平层同时为1梯1 := "中间变量1".上下平层同时为1梯1,   // "距离比较"
              上下平层同时为1梯2 := "中间变量1".上下平层同时为1梯2,
              上下平层同时为1梯3 := "中间变量1".上下平层同时为1梯3,
              上下平层同时为1梯4 := "中间变量1".上下平层同时为1梯4,
              上下平层同时为1梯5 := "中间变量1".上下平层同时为1梯5,
              上下平层同时为1梯6 := "中间变量1".上下平层同时为1梯6,
              有外呼楼层内选1 := "输出"."1号梯8层按钮指示灯",
              有外呼楼层内选2 := "输出"."2号梯8层按钮指示灯",
              有外呼楼层内选3 := "输出"."3号梯8层按钮指示灯",
              有外呼楼层内选4 := "输出"."4号梯8层按钮指示灯",
              有外呼楼层内选5 := "输出"."5号梯8层按钮指示灯",
              有外呼楼层内选6 := "输出"."6号梯8层按钮指示灯",
              就近运动电梯1 := "中间变量2".就近运动电梯1,
              就近运动电梯2 := "中间变量2".就近运动电梯2,
              就近运动电梯3 := "中间变量2".就近运动电梯3,
              就近运动电梯4 := "中间变量2".就近运动电梯4,
              就近运动电梯5 := "中间变量2".就近运动电梯5,
              就近运动电梯6 := "中间变量2".就近运动电梯6,
              呼灯 := "输出"."8层下行呼梯按钮指示灯",
              调度距离1 := "中间变量2"."1梯8层最终调度距离下",
              调度距离2 := "中间变量2"."2梯8层最终调度距离下",
              调度距离3 := "中间变量2"."3梯8层最终调度距离下",
              调度距离4 := "中间变量2"."4梯8层最终调度距离下",
              调度距离5 := "中间变量2"."5梯8层最终调度距离下",
              调度距离6 := "中间变量2"."6梯8层最终调度距离下",
              分配给1 => "中间变量2"."8层下呼分配1",
              分配给2 => "中间变量2"."8层下呼分配2",
              分配给3 => "中间变量2"."8层下呼分配3",
              分配给4 => "中间变量2"."8层下呼分配4",
              分配给5 => "中间变量2"."8层下呼分配5",
              分配给6 => "中间变量2"."8层下呼分配6");
END_REGION

REGION Network 16: 9层上呼
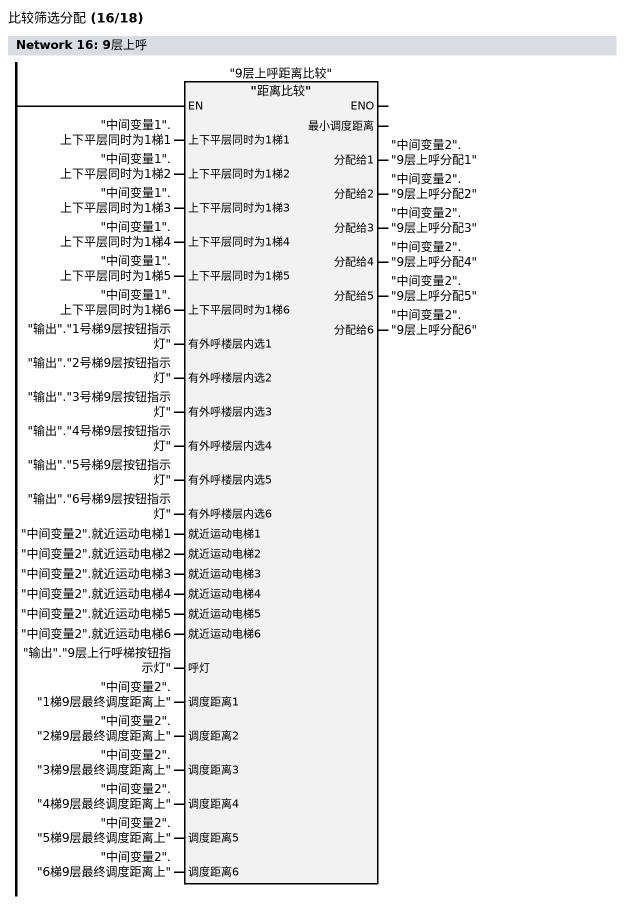
   RUNG wire#powerrail
      "9层上呼距离比较"(上下平层同时为1梯1 := "中间变量1".上下平层同时为1梯1, 上下平层同时为1梯2 := "中间变量1".上下平层同时为1梯2, 上下平层同时为1梯3 := "中间变量1".上下平层同时为1梯3, 上下平层同时为1梯4 := "中间变量1".上下平层同时为1梯4, 上下平层同时为1梯5 := "中间变量1".上下平层同时为1梯5, 上下平层同时为1梯6 := "中间变量1".上下平层同时为1梯6, 有外呼楼层内选1 := "输出"."1号梯9层按钮指示灯", 有外呼楼层内选2 := "输出"."2号梯9层按钮指示灯", 有外呼楼层内选3 := "输出"."3号梯9层按钮指示灯", 有外呼楼层内选4 := "输出"."4号梯9层按钮指示灯", 有外呼楼层内选5 := "输出"."5号梯9层按钮指示灯", 有外呼楼层内选6 := "输出"."6号梯9层按钮指示灯", 就近运动电梯1 := "中间变量2".就近运动电梯1, 就近运动电梯2 := "中间变量2".就近运动电梯2, 就近运动电梯3 := "中间变量2".就近运动电梯3, 就近运动电梯4 := "中间变量2".就近运动电梯4, 就近运动电梯5 := "中间变量2".就近运动电梯5, 就近运动电梯6 := "中间变量2".就近运动电梯6, 呼灯 := "输出"."9层上行呼梯按钮指示灯", 调度距离1 := "中间变量2"."1梯9层最终调度距离上", 调度距离2 := "中间变量2"."2梯9层最终调度距离上", 调度距离3 := "中间变量2"."3梯9层最终调度距离上", 调度距离4 := "中间变量2"."4梯9层最终调度距离上", 调度距离5 := "中间变量2"."5梯9层最终调度距离上", 调度距离6 := "中间变量2"."6梯9层最终调度距离上", 最小调度距离 =>, 分配给1 => "中间变量2"."9层上呼分配1", 分配给2 => "中间变量2"."9层上呼分配2", 分配给3 => "中间变量2"."9层上呼分配3", 分配给4 => "中间变量2"."9层上呼分配4", 分配给5 => "中间变量2"."9层上呼分配5", 分配给6 => "中间变量2"."9层上呼分配6")
   END_RUNG
   // the same network as SCL:
   "9层上呼距离比较"(上下平层同时为1梯1 := "中间变量1".上下平层同时为1梯1,   // "距离比较"
              上下平层同时为1梯2 := "中间变量1".上下平层同时为1梯2,
              上下平层同时为1梯3 := "中间变量1".上下平层同时为1梯3,
              上下平层同时为1梯4 := "中间变量1".上下平层同时为1梯4,
              上下平层同时为1梯5 := "中间变量1".上下平层同时为1梯5,
              上下平层同时为1梯6 := "中间变量1".上下平层同时为1梯6,
              有外呼楼层内选1 := "输出"."1号梯9层按钮指示灯",
              有外呼楼层内选2 := "输出"."2号梯9层按钮指示灯",
              有外呼楼层内选3 := "输出"."3号梯9层按钮指示灯",
              有外呼楼层内选4 := "输出"."4号梯9层按钮指示灯",
              有外呼楼层内选5 := "输出"."5号梯9层按钮指示灯",
              有外呼楼层内选6 := "输出"."6号梯9层按钮指示灯",
              就近运动电梯1 := "中间变量2".就近运动电梯1,
              就近运动电梯2 := "中间变量2".就近运动电梯2,
              就近运动电梯3 := "中间变量2".就近运动电梯3,
              就近运动电梯4 := "中间变量2".就近运动电梯4,
              就近运动电梯5 := "中间变量2".就近运动电梯5,
              就近运动电梯6 := "中间变量2".就近运动电梯6,
              呼灯 := "输出"."9层上行呼梯按钮指示灯",
              调度距离1 := "中间变量2"."1梯9层最终调度距离上",
              调度距离2 := "中间变量2"."2梯9层最终调度距离上",
              调度距离3 := "中间变量2"."3梯9层最终调度距离上",
              调度距离4 := "中间变量2"."4梯9层最终调度距离上",
              调度距离5 := "中间变量2"."5梯9层最终调度距离上",
              调度距离6 := "中间变量2"."6梯9层最终调度距离上",
              分配给1 => "中间变量2"."9层上呼分配1",
              分配给2 => "中间变量2"."9层上呼分配2",
              分配给3 => "中间变量2"."9层上呼分配3",
              分配给4 => "中间变量2"."9层上呼分配4",
              分配给5 => "中间变量2"."9层上呼分配5",
              分配给6 => "中间变量2"."9层上呼分配6");
END_REGION

REGION Network 17: 9层下呼
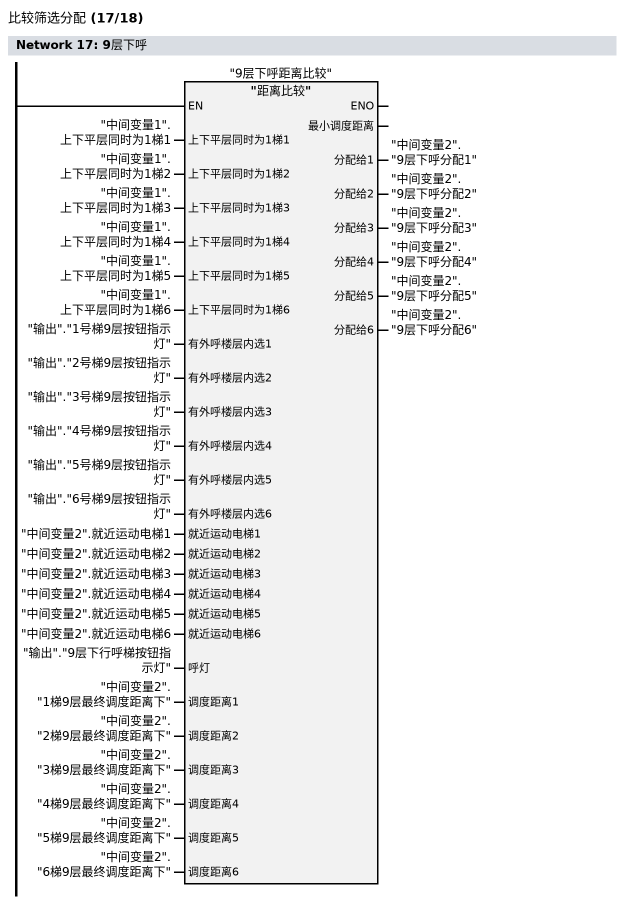
   RUNG wire#powerrail
      "9层下呼距离比较"(上下平层同时为1梯1 := "中间变量1".上下平层同时为1梯1, 上下平层同时为1梯2 := "中间变量1".上下平层同时为1梯2, 上下平层同时为1梯3 := "中间变量1".上下平层同时为1梯3, 上下平层同时为1梯4 := "中间变量1".上下平层同时为1梯4, 上下平层同时为1梯5 := "中间变量1".上下平层同时为1梯5, 上下平层同时为1梯6 := "中间变量1".上下平层同时为1梯6, 有外呼楼层内选1 := "输出"."1号梯9层按钮指示灯", 有外呼楼层内选2 := "输出"."2号梯9层按钮指示灯", 有外呼楼层内选3 := "输出"."3号梯9层按钮指示灯", 有外呼楼层内选4 := "输出"."4号梯9层按钮指示灯", 有外呼楼层内选5 := "输出"."5号梯9层按钮指示灯", 有外呼楼层内选6 := "输出"."6号梯9层按钮指示灯", 就近运动电梯1 := "中间变量2".就近运动电梯1, 就近运动电梯2 := "中间变量2".就近运动电梯2, 就近运动电梯3 := "中间变量2".就近运动电梯3, 就近运动电梯4 := "中间变量2".就近运动电梯4, 就近运动电梯5 := "中间变量2".就近运动电梯5, 就近运动电梯6 := "中间变量2".就近运动电梯6, 呼灯 := "输出"."9层下行呼梯按钮指示灯", 调度距离1 := "中间变量2"."1梯9层最终调度距离下", 调度距离2 := "中间变量2"."2梯9层最终调度距离下", 调度距离3 := "中间变量2"."3梯9层最终调度距离下", 调度距离4 := "中间变量2"."4梯9层最终调度距离下", 调度距离5 := "中间变量2"."5梯9层最终调度距离下", 调度距离6 := "中间变量2"."6梯9层最终调度距离下", 最小调度距离 =>, 分配给1 => "中间变量2"."9层下呼分配1", 分配给2 => "中间变量2"."9层下呼分配2", 分配给3 => "中间变量2"."9层下呼分配3", 分配给4 => "中间变量2"."9层下呼分配4", 分配给5 => "中间变量2"."9层下呼分配5", 分配给6 => "中间变量2"."9层下呼分配6")
   END_RUNG
   // the same network as SCL:
   "9层下呼距离比较"(上下平层同时为1梯1 := "中间变量1".上下平层同时为1梯1,   // "距离比较"
              上下平层同时为1梯2 := "中间变量1".上下平层同时为1梯2,
              上下平层同时为1梯3 := "中间变量1".上下平层同时为1梯3,
              上下平层同时为1梯4 := "中间变量1".上下平层同时为1梯4,
              上下平层同时为1梯5 := "中间变量1".上下平层同时为1梯5,
              上下平层同时为1梯6 := "中间变量1".上下平层同时为1梯6,
              有外呼楼层内选1 := "输出"."1号梯9层按钮指示灯",
              有外呼楼层内选2 := "输出"."2号梯9层按钮指示灯",
              有外呼楼层内选3 := "输出"."3号梯9层按钮指示灯",
              有外呼楼层内选4 := "输出"."4号梯9层按钮指示灯",
              有外呼楼层内选5 := "输出"."5号梯9层按钮指示灯",
              有外呼楼层内选6 := "输出"."6号梯9层按钮指示灯",
              就近运动电梯1 := "中间变量2".就近运动电梯1,
              就近运动电梯2 := "中间变量2".就近运动电梯2,
              就近运动电梯3 := "中间变量2".就近运动电梯3,
              就近运动电梯4 := "中间变量2".就近运动电梯4,
              就近运动电梯5 := "中间变量2".就近运动电梯5,
              就近运动电梯6 := "中间变量2".就近运动电梯6,
              呼灯 := "输出"."9层下行呼梯按钮指示灯",
              调度距离1 := "中间变量2"."1梯9层最终调度距离下",
              调度距离2 := "中间变量2"."2梯9层最终调度距离下",
              调度距离3 := "中间变量2"."3梯9层最终调度距离下",
              调度距离4 := "中间变量2"."4梯9层最终调度距离下",
              调度距离5 := "中间变量2"."5梯9层最终调度距离下",
              调度距离6 := "中间变量2"."6梯9层最终调度距离下",
              分配给1 => "中间变量2"."9层下呼分配1",
              分配给2 => "中间变量2"."9层下呼分配2",
              分配给3 => "中间变量2"."9层下呼分配3",
              分配给4 => "中间变量2"."9层下呼分配4",
              分配给5 => "中间变量2"."9层下呼分配5",
              分配给6 => "中间变量2"."9层下呼分配6");
END_REGION

REGION Network 18: 10层下呼
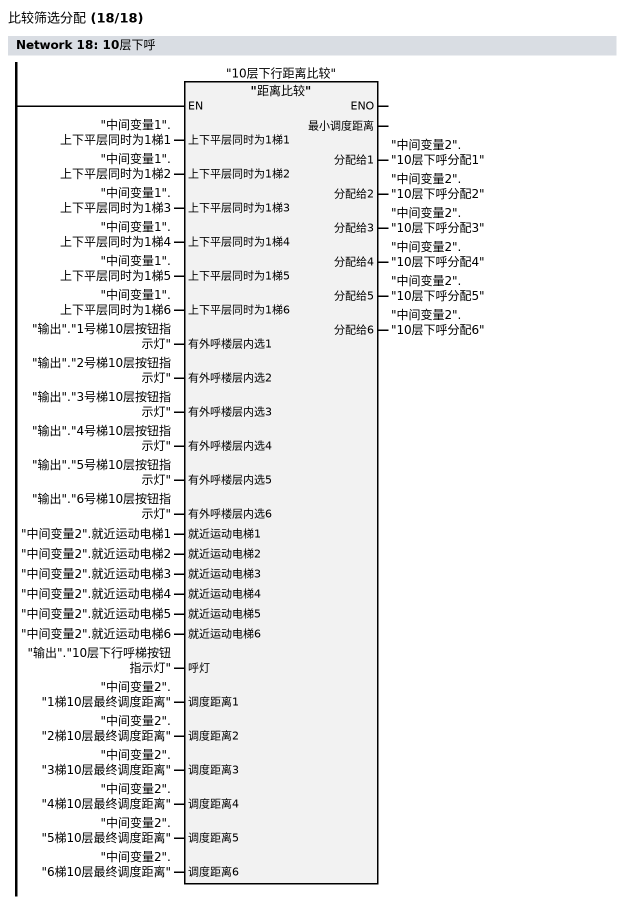
   RUNG wire#powerrail
      "10层下行距离比较"(上下平层同时为1梯1 := "中间变量1".上下平层同时为1梯1, 上下平层同时为1梯2 := "中间变量1".上下平层同时为1梯2, 上下平层同时为1梯3 := "中间变量1".上下平层同时为1梯3, 上下平层同时为1梯4 := "中间变量1".上下平层同时为1梯4, 上下平层同时为1梯5 := "中间变量1".上下平层同时为1梯5, 上下平层同时为1梯6 := "中间变量1".上下平层同时为1梯6, 有外呼楼层内选1 := "输出"."1号梯10层按钮指示灯", 有外呼楼层内选2 := "输出"."2号梯10层按钮指示灯", 有外呼楼层内选3 := "输出"."3号梯10层按钮指示灯", 有外呼楼层内选4 := "输出"."4号梯10层按钮指示灯", 有外呼楼层内选5 := "输出"."5号梯10层按钮指示灯", 有外呼楼层内选6 := "输出"."6号梯10层按钮指示灯", 就近运动电梯1 := "中间变量2".就近运动电梯1, 就近运动电梯2 := "中间变量2".就近运动电梯2, 就近运动电梯3 := "中间变量2".就近运动电梯3, 就近运动电梯4 := "中间变量2".就近运动电梯4, 就近运动电梯5 := "中间变量2".就近运动电梯5, 就近运动电梯6 := "中间变量2".就近运动电梯6, 呼灯 := "输出"."10层下行呼梯按钮指示灯", 调度距离1 := "中间变量2"."1梯10层最终调度距离", 调度距离2 := "中间变量2"."2梯10层最终调度距离", 调度距离3 := "中间变量2"."3梯10层最终调度距离", 调度距离4 := "中间变量2"."4梯10层最终调度距离", 调度距离5 := "中间变量2"."5梯10层最终调度距离", 调度距离6 := "中间变量2"."6梯10层最终调度距离", 最小调度距离 =>, 分配给1 => "中间变量2"."10层下呼分配1", 分配给2 => "中间变量2"."10层下呼分配2", 分配给3 => "中间变量2"."10层下呼分配3", 分配给4 => "中间变量2"."10层下呼分配4", 分配给5 => "中间变量2"."10层下呼分配5", 分配给6 => "中间变量2"."10层下呼分配6")
   END_RUNG
   // the same network as SCL:
   "10层下行距离比较"(上下平层同时为1梯1 := "中间变量1".上下平层同时为1梯1,   // "距离比较"
               上下平层同时为1梯2 := "中间变量1".上下平层同时为1梯2,
               上下平层同时为1梯3 := "中间变量1".上下平层同时为1梯3,
               上下平层同时为1梯4 := "中间变量1".上下平层同时为1梯4,
               上下平层同时为1梯5 := "中间变量1".上下平层同时为1梯5,
               上下平层同时为1梯6 := "中间变量1".上下平层同时为1梯6,
               有外呼楼层内选1 := "输出"."1号梯10层按钮指示灯",
               有外呼楼层内选2 := "输出"."2号梯10层按钮指示灯",
               有外呼楼层内选3 := "输出"."3号梯10层按钮指示灯",
               有外呼楼层内选4 := "输出"."4号梯10层按钮指示灯",
               有外呼楼层内选5 := "输出"."5号梯10层按钮指示灯",
               有外呼楼层内选6 := "输出"."6号梯10层按钮指示灯",
               就近运动电梯1 := "中间变量2".就近运动电梯1,
               就近运动电梯2 := "中间变量2".就近运动电梯2,
               就近运动电梯3 := "中间变量2".就近运动电梯3,
               就近运动电梯4 := "中间变量2".就近运动电梯4,
               就近运动电梯5 := "中间变量2".就近运动电梯5,
               就近运动电梯6 := "中间变量2".就近运动电梯6,
               呼灯 := "输出"."10层下行呼梯按钮指示灯",
               调度距离1 := "中间变量2"."1梯10层最终调度距离",
               调度距离2 := "中间变量2"."2梯10层最终调度距离",
               调度距离3 := "中间变量2"."3梯10层最终调度距离",
               调度距离4 := "中间变量2"."4梯10层最终调度距离",
               调度距离5 := "中间变量2"."5梯10层最终调度距离",
               调度距离6 := "中间变量2"."6梯10层最终调度距离",
               分配给1 => "中间变量2"."10层下呼分配1",
               分配给2 => "中间变量2"."10层下呼分配2",
               分配给3 => "中间变量2"."10层下呼分配3",
               分配给4 => "中间变量2"."10层下呼分配4",
               分配给5 => "中间变量2"."10层下呼分配5",
               分配给6 => "中间变量2"."10层下呼分配6");
END_REGION
END_FUNCTION

FUNCTION "电梯初始化" : Void   // FC2, LAD
{ S7_Optimized_Access := 'TRUE' }
VERSION : 0.1
BEGIN

REGION Network 1: 1号梯初始化
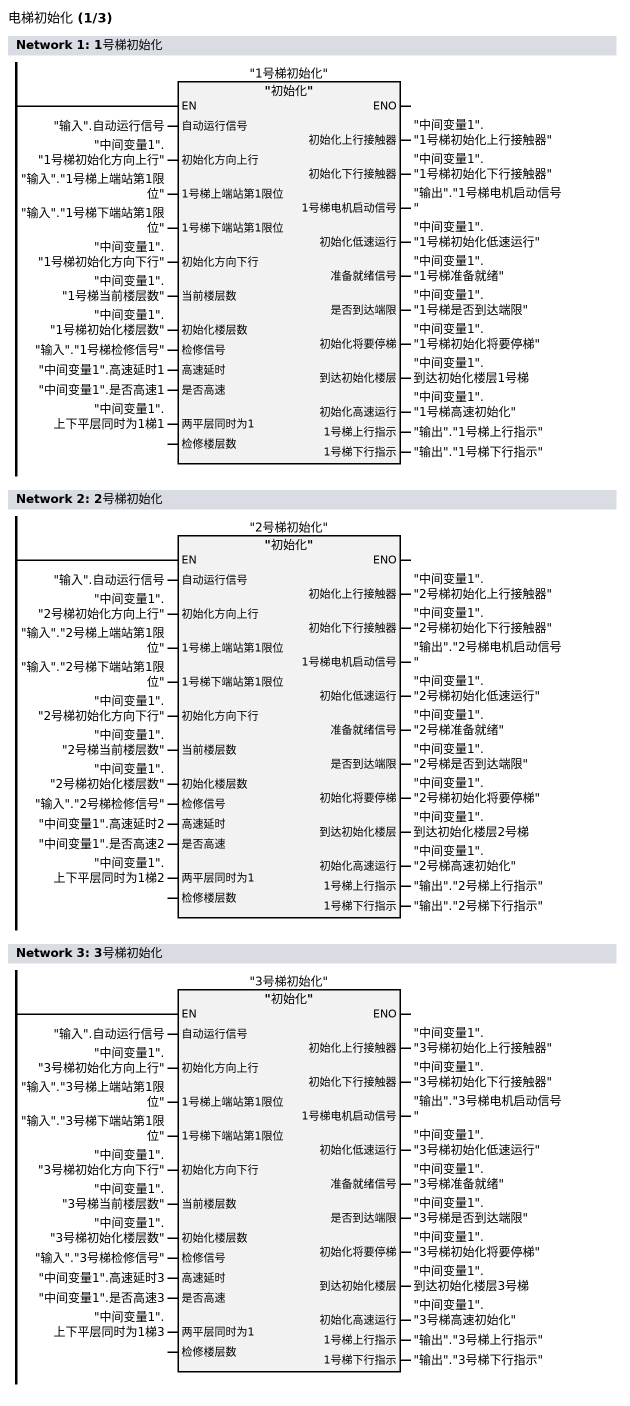
   RUNG wire#powerrail
      "1号梯初始化"(自动运行信号 := "输入".自动运行信号, 初始化方向上行 := "中间变量1"."1号梯初始化方向上行", "1号梯上端站第1限位" := "输入"."1号梯上端站第1限位", "1号梯下端站第1限位" := "输入"."1号梯下端站第1限位", 初始化方向下行 := "中间变量1"."1号梯初始化方向下行", 当前楼层数 := "中间变量1"."1号梯当前楼层数", 初始化楼层数 := "中间变量1"."1号梯初始化楼层数", 检修信号 := "输入"."1号梯检修信号", 高速延时 := "中间变量1".高速延时1, 是否高速 := "中间变量1".是否高速1, 两平层同时为1 := "中间变量1".上下平层同时为1梯1, 检修楼层数 :=, 初始化上行接触器 => "中间变量1"."1号梯初始化上行接触器", 初始化下行接触器 => "中间变量1"."1号梯初始化下行接触器", "1号梯电机启动信号" => "输出"."1号梯电机启动信号", 初始化低速运行 => "中间变量1"."1号梯初始化低速运行", 准备就绪信号 => "中间变量1"."1号梯准备就绪", 是否到达端限 => "中间变量1"."1号梯是否到达端限", 初始化将要停梯 => "中间变量1"."1号梯初始化将要停梯", 到达初始化楼层 => "中间变量1".到达初始化楼层1号梯, 初始化高速运行 => "中间变量1"."1号梯高速初始化", "1号梯上行指示" => "输出"."1号梯上行指示", "1号梯下行指示" => "输出"."1号梯下行指示")
   END_RUNG
   // the same network as SCL:
   "1号梯初始化"(自动运行信号 := "输入".自动运行信号,   // "初始化"
            初始化方向上行 := "中间变量1"."1号梯初始化方向上行",
            "1号梯上端站第1限位" := "输入"."1号梯上端站第1限位",
            "1号梯下端站第1限位" := "输入"."1号梯下端站第1限位",
            初始化方向下行 := "中间变量1"."1号梯初始化方向下行",
            当前楼层数 := "中间变量1"."1号梯当前楼层数",
            初始化楼层数 := "中间变量1"."1号梯初始化楼层数",
            检修信号 := "输入"."1号梯检修信号",
            高速延时 := "中间变量1".高速延时1,
            是否高速 := "中间变量1".是否高速1,
            两平层同时为1 := "中间变量1".上下平层同时为1梯1,
            初始化上行接触器 => "中间变量1"."1号梯初始化上行接触器",
            初始化下行接触器 => "中间变量1"."1号梯初始化下行接触器",
            "1号梯电机启动信号" => "输出"."1号梯电机启动信号",
            初始化低速运行 => "中间变量1"."1号梯初始化低速运行",
            准备就绪信号 => "中间变量1"."1号梯准备就绪",
            是否到达端限 => "中间变量1"."1号梯是否到达端限",
            初始化将要停梯 => "中间变量1"."1号梯初始化将要停梯",
            到达初始化楼层 => "中间变量1".到达初始化楼层1号梯,
            初始化高速运行 => "中间变量1"."1号梯高速初始化",
            "1号梯上行指示" => "输出"."1号梯上行指示",
            "1号梯下行指示" => "输出"."1号梯下行指示");
END_REGION

REGION Network 2: 2号梯初始化
   RUNG wire#powerrail
      "2号梯初始化"(自动运行信号 := "输入".自动运行信号, 初始化方向上行 := "中间变量1"."2号梯初始化方向上行", "1号梯上端站第1限位" := "输入"."2号梯上端站第1限位", "1号梯下端站第1限位" := "输入"."2号梯下端站第1限位", 初始化方向下行 := "中间变量1"."2号梯初始化方向下行", 当前楼层数 := "中间变量1"."2号梯当前楼层数", 初始化楼层数 := "中间变量1"."2号梯初始化楼层数", 检修信号 := "输入"."2号梯检修信号", 高速延时 := "中间变量1".高速延时2, 是否高速 := "中间变量1".是否高速2, 两平层同时为1 := "中间变量1".上下平层同时为1梯2, 检修楼层数 :=, 初始化上行接触器 => "中间变量1"."2号梯初始化上行接触器", 初始化下行接触器 => "中间变量1"."2号梯初始化下行接触器", "1号梯电机启动信号" => "输出"."2号梯电机启动信号", 初始化低速运行 => "中间变量1"."2号梯初始化低速运行", 准备就绪信号 => "中间变量1"."2号梯准备就绪", 是否到达端限 => "中间变量1"."2号梯是否到达端限", 初始化将要停梯 => "中间变量1"."2号梯初始化将要停梯", 到达初始化楼层 => "中间变量1".到达初始化楼层2号梯, 初始化高速运行 => "中间变量1"."2号梯高速初始化", "1号梯上行指示" => "输出"."2号梯上行指示", "1号梯下行指示" => "输出"."2号梯下行指示")
   END_RUNG
   // the same network as SCL:
   "2号梯初始化"(自动运行信号 := "输入".自动运行信号,   // "初始化"
            初始化方向上行 := "中间变量1"."2号梯初始化方向上行",
            "1号梯上端站第1限位" := "输入"."2号梯上端站第1限位",
            "1号梯下端站第1限位" := "输入"."2号梯下端站第1限位",
            初始化方向下行 := "中间变量1"."2号梯初始化方向下行",
            当前楼层数 := "中间变量1"."2号梯当前楼层数",
            初始化楼层数 := "中间变量1"."2号梯初始化楼层数",
            检修信号 := "输入"."2号梯检修信号",
            高速延时 := "中间变量1".高速延时2,
            是否高速 := "中间变量1".是否高速2,
            两平层同时为1 := "中间变量1".上下平层同时为1梯2,
            初始化上行接触器 => "中间变量1"."2号梯初始化上行接触器",
            初始化下行接触器 => "中间变量1"."2号梯初始化下行接触器",
            "1号梯电机启动信号" => "输出"."2号梯电机启动信号",
            初始化低速运行 => "中间变量1"."2号梯初始化低速运行",
            准备就绪信号 => "中间变量1"."2号梯准备就绪",
            是否到达端限 => "中间变量1"."2号梯是否到达端限",
            初始化将要停梯 => "中间变量1"."2号梯初始化将要停梯",
            到达初始化楼层 => "中间变量1".到达初始化楼层2号梯,
            初始化高速运行 => "中间变量1"."2号梯高速初始化",
            "1号梯上行指示" => "输出"."2号梯上行指示",
            "1号梯下行指示" => "输出"."2号梯下行指示");
END_REGION

REGION Network 3: 3号梯初始化
   RUNG wire#powerrail
      "3号梯初始化"(自动运行信号 := "输入".自动运行信号, 初始化方向上行 := "中间变量1"."3号梯初始化方向上行", "1号梯上端站第1限位" := "输入"."3号梯上端站第1限位", "1号梯下端站第1限位" := "输入"."3号梯下端站第1限位", 初始化方向下行 := "中间变量1"."3号梯初始化方向下行", 当前楼层数 := "中间变量1"."3号梯当前楼层数", 初始化楼层数 := "中间变量1"."3号梯初始化楼层数", 检修信号 := "输入"."3号梯检修信号", 高速延时 := "中间变量1".高速延时3, 是否高速 := "中间变量1".是否高速3, 两平层同时为1 := "中间变量1".上下平层同时为1梯3, 检修楼层数 :=, 初始化上行接触器 => "中间变量1"."3号梯初始化上行接触器", 初始化下行接触器 => "中间变量1"."3号梯初始化下行接触器", "1号梯电机启动信号" => "输出"."3号梯电机启动信号", 初始化低速运行 => "中间变量1"."3号梯初始化低速运行", 准备就绪信号 => "中间变量1"."3号梯准备就绪", 是否到达端限 => "中间变量1"."3号梯是否到达端限", 初始化将要停梯 => "中间变量1"."3号梯初始化将要停梯", 到达初始化楼层 => "中间变量1".到达初始化楼层3号梯, 初始化高速运行 => "中间变量1"."3号梯高速初始化", "1号梯上行指示" => "输出"."3号梯上行指示", "1号梯下行指示" => "输出"."3号梯下行指示")
   END_RUNG
   // the same network as SCL:
   "3号梯初始化"(自动运行信号 := "输入".自动运行信号,   // "初始化"
            初始化方向上行 := "中间变量1"."3号梯初始化方向上行",
            "1号梯上端站第1限位" := "输入"."3号梯上端站第1限位",
            "1号梯下端站第1限位" := "输入"."3号梯下端站第1限位",
            初始化方向下行 := "中间变量1"."3号梯初始化方向下行",
            当前楼层数 := "中间变量1"."3号梯当前楼层数",
            初始化楼层数 := "中间变量1"."3号梯初始化楼层数",
            检修信号 := "输入"."3号梯检修信号",
            高速延时 := "中间变量1".高速延时3,
            是否高速 := "中间变量1".是否高速3,
            两平层同时为1 := "中间变量1".上下平层同时为1梯3,
            初始化上行接触器 => "中间变量1"."3号梯初始化上行接触器",
            初始化下行接触器 => "中间变量1"."3号梯初始化下行接触器",
            "1号梯电机启动信号" => "输出"."3号梯电机启动信号",
            初始化低速运行 => "中间变量1"."3号梯初始化低速运行",
            准备就绪信号 => "中间变量1"."3号梯准备就绪",
            是否到达端限 => "中间变量1"."3号梯是否到达端限",
            初始化将要停梯 => "中间变量1"."3号梯初始化将要停梯",
            到达初始化楼层 => "中间变量1".到达初始化楼层3号梯,
            初始化高速运行 => "中间变量1"."3号梯高速初始化",
            "1号梯上行指示" => "输出"."3号梯上行指示",
            "1号梯下行指示" => "输出"."3号梯下行指示");
END_REGION

REGION Network 4: 4号梯初始化
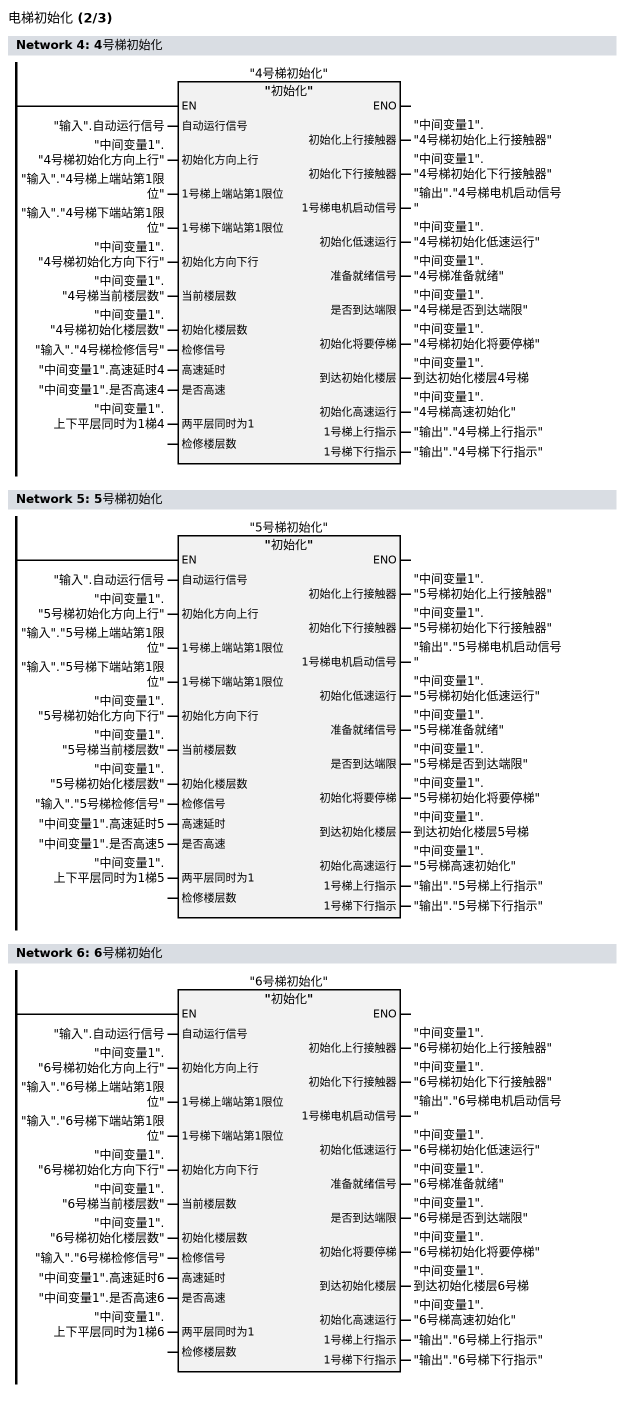
   RUNG wire#powerrail
      "4号梯初始化"(自动运行信号 := "输入".自动运行信号, 初始化方向上行 := "中间变量1"."4号梯初始化方向上行", "1号梯上端站第1限位" := "输入"."4号梯上端站第1限位", "1号梯下端站第1限位" := "输入"."4号梯下端站第1限位", 初始化方向下行 := "中间变量1"."4号梯初始化方向下行", 当前楼层数 := "中间变量1"."4号梯当前楼层数", 初始化楼层数 := "中间变量1"."4号梯初始化楼层数", 检修信号 := "输入"."4号梯检修信号", 高速延时 := "中间变量1".高速延时4, 是否高速 := "中间变量1".是否高速4, 两平层同时为1 := "中间变量1".上下平层同时为1梯4, 检修楼层数 :=, 初始化上行接触器 => "中间变量1"."4号梯初始化上行接触器", 初始化下行接触器 => "中间变量1"."4号梯初始化下行接触器", "1号梯电机启动信号" => "输出"."4号梯电机启动信号", 初始化低速运行 => "中间变量1"."4号梯初始化低速运行", 准备就绪信号 => "中间变量1"."4号梯准备就绪", 是否到达端限 => "中间变量1"."4号梯是否到达端限", 初始化将要停梯 => "中间变量1"."4号梯初始化将要停梯", 到达初始化楼层 => "中间变量1".到达初始化楼层4号梯, 初始化高速运行 => "中间变量1"."4号梯高速初始化", "1号梯上行指示" => "输出"."4号梯上行指示", "1号梯下行指示" => "输出"."4号梯下行指示")
   END_RUNG
   // the same network as SCL:
   "4号梯初始化"(自动运行信号 := "输入".自动运行信号,   // "初始化"
            初始化方向上行 := "中间变量1"."4号梯初始化方向上行",
            "1号梯上端站第1限位" := "输入"."4号梯上端站第1限位",
            "1号梯下端站第1限位" := "输入"."4号梯下端站第1限位",
            初始化方向下行 := "中间变量1"."4号梯初始化方向下行",
            当前楼层数 := "中间变量1"."4号梯当前楼层数",
            初始化楼层数 := "中间变量1"."4号梯初始化楼层数",
            检修信号 := "输入"."4号梯检修信号",
            高速延时 := "中间变量1".高速延时4,
            是否高速 := "中间变量1".是否高速4,
            两平层同时为1 := "中间变量1".上下平层同时为1梯4,
            初始化上行接触器 => "中间变量1"."4号梯初始化上行接触器",
            初始化下行接触器 => "中间变量1"."4号梯初始化下行接触器",
            "1号梯电机启动信号" => "输出"."4号梯电机启动信号",
            初始化低速运行 => "中间变量1"."4号梯初始化低速运行",
            准备就绪信号 => "中间变量1"."4号梯准备就绪",
            是否到达端限 => "中间变量1"."4号梯是否到达端限",
            初始化将要停梯 => "中间变量1"."4号梯初始化将要停梯",
            到达初始化楼层 => "中间变量1".到达初始化楼层4号梯,
            初始化高速运行 => "中间变量1"."4号梯高速初始化",
            "1号梯上行指示" => "输出"."4号梯上行指示",
            "1号梯下行指示" => "输出"."4号梯下行指示");
END_REGION

REGION Network 5: 5号梯初始化
   RUNG wire#powerrail
      "5号梯初始化"(自动运行信号 := "输入".自动运行信号, 初始化方向上行 := "中间变量1"."5号梯初始化方向上行", "1号梯上端站第1限位" := "输入"."5号梯上端站第1限位", "1号梯下端站第1限位" := "输入"."5号梯下端站第1限位", 初始化方向下行 := "中间变量1"."5号梯初始化方向下行", 当前楼层数 := "中间变量1"."5号梯当前楼层数", 初始化楼层数 := "中间变量1"."5号梯初始化楼层数", 检修信号 := "输入"."5号梯检修信号", 高速延时 := "中间变量1".高速延时5, 是否高速 := "中间变量1".是否高速5, 两平层同时为1 := "中间变量1".上下平层同时为1梯5, 检修楼层数 :=, 初始化上行接触器 => "中间变量1"."5号梯初始化上行接触器", 初始化下行接触器 => "中间变量1"."5号梯初始化下行接触器", "1号梯电机启动信号" => "输出"."5号梯电机启动信号", 初始化低速运行 => "中间变量1"."5号梯初始化低速运行", 准备就绪信号 => "中间变量1"."5号梯准备就绪", 是否到达端限 => "中间变量1"."5号梯是否到达端限", 初始化将要停梯 => "中间变量1"."5号梯初始化将要停梯", 到达初始化楼层 => "中间变量1".到达初始化楼层5号梯, 初始化高速运行 => "中间变量1"."5号梯高速初始化", "1号梯上行指示" => "输出"."5号梯上行指示", "1号梯下行指示" => "输出"."5号梯下行指示")
   END_RUNG
   // the same network as SCL:
   "5号梯初始化"(自动运行信号 := "输入".自动运行信号,   // "初始化"
            初始化方向上行 := "中间变量1"."5号梯初始化方向上行",
            "1号梯上端站第1限位" := "输入"."5号梯上端站第1限位",
            "1号梯下端站第1限位" := "输入"."5号梯下端站第1限位",
            初始化方向下行 := "中间变量1"."5号梯初始化方向下行",
            当前楼层数 := "中间变量1"."5号梯当前楼层数",
            初始化楼层数 := "中间变量1"."5号梯初始化楼层数",
            检修信号 := "输入"."5号梯检修信号",
            高速延时 := "中间变量1".高速延时5,
            是否高速 := "中间变量1".是否高速5,
            两平层同时为1 := "中间变量1".上下平层同时为1梯5,
            初始化上行接触器 => "中间变量1"."5号梯初始化上行接触器",
            初始化下行接触器 => "中间变量1"."5号梯初始化下行接触器",
            "1号梯电机启动信号" => "输出"."5号梯电机启动信号",
            初始化低速运行 => "中间变量1"."5号梯初始化低速运行",
            准备就绪信号 => "中间变量1"."5号梯准备就绪",
            是否到达端限 => "中间变量1"."5号梯是否到达端限",
            初始化将要停梯 => "中间变量1"."5号梯初始化将要停梯",
            到达初始化楼层 => "中间变量1".到达初始化楼层5号梯,
            初始化高速运行 => "中间变量1"."5号梯高速初始化",
            "1号梯上行指示" => "输出"."5号梯上行指示",
            "1号梯下行指示" => "输出"."5号梯下行指示");
END_REGION

REGION Network 6: 6号梯初始化
   RUNG wire#powerrail
      "6号梯初始化"(自动运行信号 := "输入".自动运行信号, 初始化方向上行 := "中间变量1"."6号梯初始化方向上行", "1号梯上端站第1限位" := "输入"."6号梯上端站第1限位", "1号梯下端站第1限位" := "输入"."6号梯下端站第1限位", 初始化方向下行 := "中间变量1"."6号梯初始化方向下行", 当前楼层数 := "中间变量1"."6号梯当前楼层数", 初始化楼层数 := "中间变量1"."6号梯初始化楼层数", 检修信号 := "输入"."6号梯检修信号", 高速延时 := "中间变量1".高速延时6, 是否高速 := "中间变量1".是否高速6, 两平层同时为1 := "中间变量1".上下平层同时为1梯6, 检修楼层数 :=, 初始化上行接触器 => "中间变量1"."6号梯初始化上行接触器", 初始化下行接触器 => "中间变量1"."6号梯初始化下行接触器", "1号梯电机启动信号" => "输出"."6号梯电机启动信号", 初始化低速运行 => "中间变量1"."6号梯初始化低速运行", 准备就绪信号 => "中间变量1"."6号梯准备就绪", 是否到达端限 => "中间变量1"."6号梯是否到达端限", 初始化将要停梯 => "中间变量1"."6号梯初始化将要停梯", 到达初始化楼层 => "中间变量1".到达初始化楼层6号梯, 初始化高速运行 => "中间变量1"."6号梯高速初始化", "1号梯上行指示" => "输出"."6号梯上行指示", "1号梯下行指示" => "输出"."6号梯下行指示")
   END_RUNG
   // the same network as SCL:
   "6号梯初始化"(自动运行信号 := "输入".自动运行信号,   // "初始化"
            初始化方向上行 := "中间变量1"."6号梯初始化方向上行",
            "1号梯上端站第1限位" := "输入"."6号梯上端站第1限位",
            "1号梯下端站第1限位" := "输入"."6号梯下端站第1限位",
            初始化方向下行 := "中间变量1"."6号梯初始化方向下行",
            当前楼层数 := "中间变量1"."6号梯当前楼层数",
            初始化楼层数 := "中间变量1"."6号梯初始化楼层数",
            检修信号 := "输入"."6号梯检修信号",
            高速延时 := "中间变量1".高速延时6,
            是否高速 := "中间变量1".是否高速6,
            两平层同时为1 := "中间变量1".上下平层同时为1梯6,
            初始化上行接触器 => "中间变量1"."6号梯初始化上行接触器",
            初始化下行接触器 => "中间变量1"."6号梯初始化下行接触器",
            "1号梯电机启动信号" => "输出"."6号梯电机启动信号",
            初始化低速运行 => "中间变量1"."6号梯初始化低速运行",
            准备就绪信号 => "中间变量1"."6号梯准备就绪",
            是否到达端限 => "中间变量1"."6号梯是否到达端限",
            初始化将要停梯 => "中间变量1"."6号梯初始化将要停梯",
            到达初始化楼层 => "中间变量1".到达初始化楼层6号梯,
            初始化高速运行 => "中间变量1"."6号梯高速初始化",
            "1号梯上行指示" => "输出"."6号梯上行指示",
            "1号梯下行指示" => "输出"."6号梯下行指示");
END_REGION

REGION Network 7: 准备就绪输出
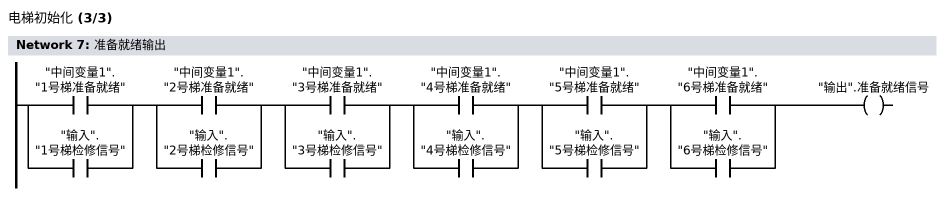
   RUNG wire#powerrail
      Contact( "中间变量1"."1号梯准备就绪" )
      wire#w1
      Contact( "中间变量1"."2号梯准备就绪" )
      wire#w2
      Contact( "中间变量1"."3号梯准备就绪" )
      wire#w3
      Contact( "中间变量1"."4号梯准备就绪" )
      wire#w4
      Contact( "中间变量1"."5号梯准备就绪" )
      wire#w5
      Contact( "中间变量1"."6号梯准备就绪" )
      wire#w6
      Coil( "输出".准备就绪信号 )
   END_RUNG
   RUNG wire#powerrail
      Contact( "输入"."1号梯检修信号" )
   END_RUNG wire#w1
   RUNG wire#w1
      Contact( "输入"."2号梯检修信号" )
   END_RUNG wire#w2
   RUNG wire#w2
      Contact( "输入"."3号梯检修信号" )
   END_RUNG wire#w3
   RUNG wire#w3
      Contact( "输入"."4号梯检修信号" )
   END_RUNG wire#w4
   RUNG wire#w4
      Contact( "输入"."5号梯检修信号" )
   END_RUNG wire#w5
   RUNG wire#w5
      Contact( "输入"."6号梯检修信号" )
   END_RUNG wire#w6
   // the same network as SCL:
   "输出".准备就绪信号 := ("中间变量1"."1号梯准备就绪" OR "输入"."1号梯检修信号") AND ("中间变量1"."2号梯准备就绪" OR "输入"."2号梯检修信号") AND ("中间变量1"."3号梯准备就绪" OR "输入"."3号梯检修信号") AND ("中间变量1"."4号梯准备就绪" OR "输入"."4号梯检修信号") AND ("中间变量1"."5号梯准备就绪" OR "输入"."5号梯检修信号") AND ("中间变量1"."6号梯准备就绪" OR "输入"."6号梯检修信号");
END_REGION
END_FUNCTION

FUNCTION "电梯高低速转换" : Void   // FC3, LAD
{ S7_Optimized_Access := 'TRUE' }
VERSION : 0.1
BEGIN

REGION Network 1: 1号梯
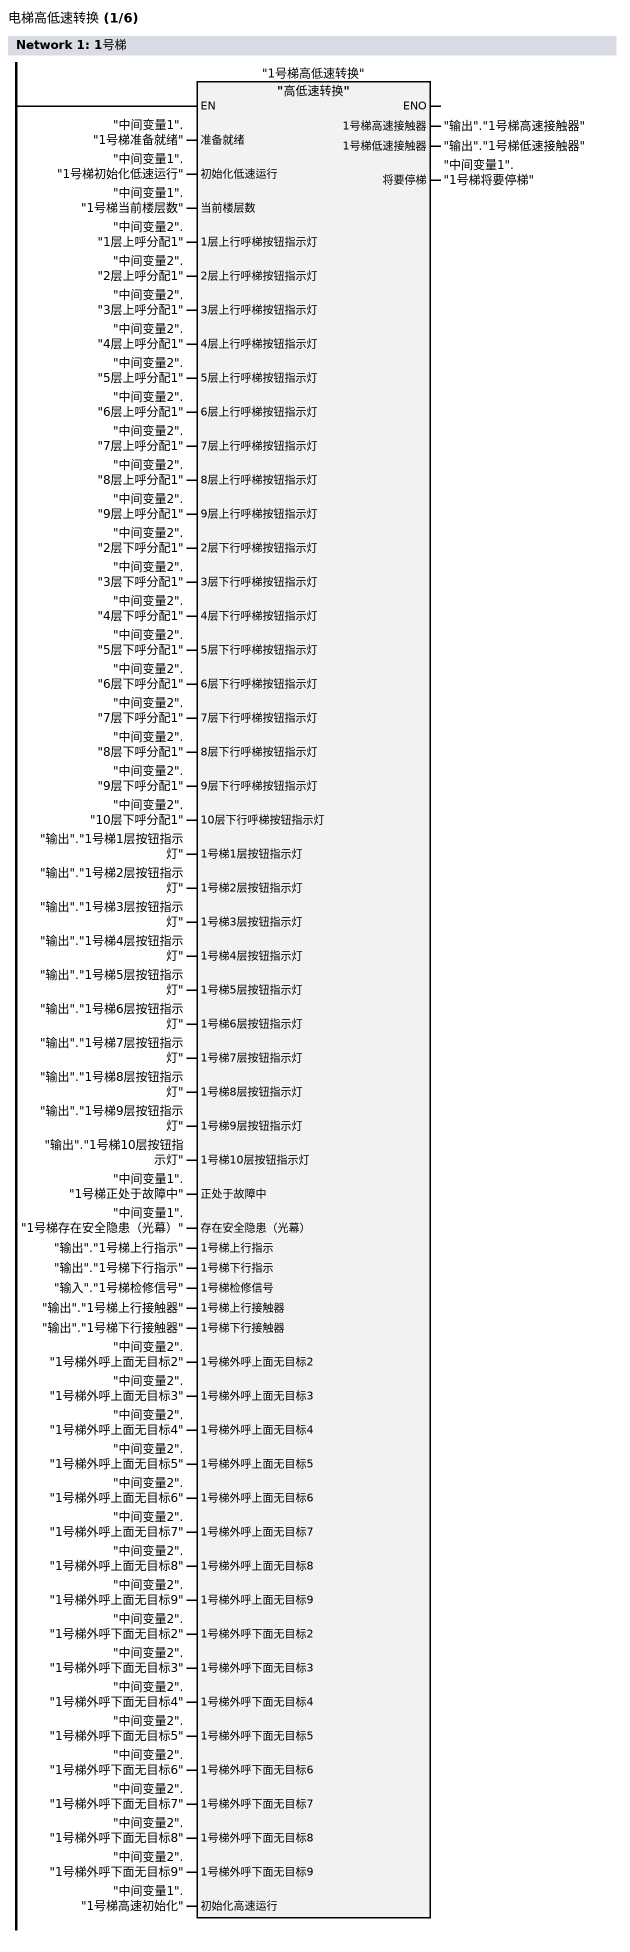
   RUNG wire#powerrail
      "1号梯高低速转换"(准备就绪 := "中间变量1"."1号梯准备就绪", 初始化低速运行 := "中间变量1"."1号梯初始化低速运行", 当前楼层数 := "中间变量1"."1号梯当前楼层数", "1层上行呼梯按钮指示灯" := "中间变量2"."1层上呼分配1", "2层上行呼梯按钮指示灯" := "中间变量2"."2层上呼分配1", "3层上行呼梯按钮指示灯" := "中间变量2"."3层上呼分配1", "4层上行呼梯按钮指示灯" := "中间变量2"."4层上呼分配1", "5层上行呼梯按钮指示灯" := "中间变量2"."5层上呼分配1", "6层上行呼梯按钮指示灯" := "中间变量2"."6层上呼分配1", "7层上行呼梯按钮指示灯" := "中间变量2"."7层上呼分配1", "8层上行呼梯按钮指示灯" := "中间变量2"."8层上呼分配1", "9层上行呼梯按钮指示灯" := "中间变量2"."9层上呼分配1", "2层下行呼梯按钮指示灯" := "中间变量2"."2层下呼分配1", "3层下行呼梯按钮指示灯" := "中间变量2"."3层下呼分配1", "4层下行呼梯按钮指示灯" := "中间变量2"."4层下呼分配1", "5层下行呼梯按钮指示灯" := "中间变量2"."5层下呼分配1", "6层下行呼梯按钮指示灯" := "中间变量2"."6层下呼分配1", "7层下行呼梯按钮指示灯" := "中间变量2"."7层下呼分配1", "8层下行呼梯按钮指示灯" := "中间变量2"."8层下呼分配1", "9层下行呼梯按钮指示灯" := "中间变量2"."9层下呼分配1", "10层下行呼梯按钮指示灯" := "中间变量2"."10层下呼分配1", "1号梯1层按钮指示灯" := "输出"."1号梯1层按钮指示灯", "1号梯2层按钮指示灯" := "输出"."1号梯2层按钮指示灯", "1号梯3层按钮指示灯" := "输出"."1号梯3层按钮指示灯", "1号梯4层按钮指示灯" := "输出"."1号梯4层按钮指示灯", "1号梯5层按钮指示灯" := "输出"."1号梯5层按钮指示灯", "1号梯6层按钮指示灯" := "输出"."1号梯6层按钮指示灯", "1号梯7层按钮指示灯" := "输出"."1号梯7层按钮指示灯", "1号梯8层按钮指示灯" := "输出"."1号梯8层按钮指示灯", "1号梯9层按钮指示灯" := "输出"."1号梯9层按钮指示灯", "1号梯10层按钮指示灯" := "输出"."1号梯10层按钮指示灯", 正处于故障中 := "中间变量1"."1号梯正处于故障中", "存在安全隐患（光幕）" := "中间变量1"."1号梯存在安全隐患（光幕）", "1号梯上行指示" := "输出"."1号梯上行指示", "1号梯下行指示" := "输出"."1号梯下行指示", "1号梯检修信号" := "输入"."1号梯检修信号", "1号梯上行接触器" := "输出"."1号梯上行接触器", "1号梯下行接触器" := "输出"."1号梯下行接触器", "1号梯外呼上面无目标2" := "中间变量2"."1号梯外呼上面无目标2", "1号梯外呼上面无目标3" := "中间变量2"."1号梯外呼上面无目标3", "1号梯外呼上面无目标4" := "中间变量2"."1号梯外呼上面无目标4", "1号梯外呼上面无目标5" := "中间变量2"."1号梯外呼上面无目标5", "1号梯外呼上面无目标6" := "中间变量2"."1号梯外呼上面无目标6", "1号梯外呼上面无目标7" := "中间变量2"."1号梯外呼上面无目标7", "1号梯外呼上面无目标8" := "中间变量2"."1号梯外呼上面无目标8", "1号梯外呼上面无目标9" := "中间变量2"."1号梯外呼上面无目标9", "1号梯外呼下面无目标2" := "中间变量2"."1号梯外呼下面无目标2", "1号梯外呼下面无目标3" := "中间变量2"."1号梯外呼下面无目标3", "1号梯外呼下面无目标4" := "中间变量2"."1号梯外呼下面无目标4", "1号梯外呼下面无目标5" := "中间变量2"."1号梯外呼下面无目标5", "1号梯外呼下面无目标6" := "中间变量2"."1号梯外呼下面无目标6", "1号梯外呼下面无目标7" := "中间变量2"."1号梯外呼下面无目标7", "1号梯外呼下面无目标8" := "中间变量2"."1号梯外呼下面无目标8", "1号梯外呼下面无目标9" := "中间变量2"."1号梯外呼下面无目标9", 初始化高速运行 := "中间变量1"."1号梯高速初始化", "1号梯高速接触器" => "输出"."1号梯高速接触器", "1号梯低速接触器" => "输出"."1号梯低速接触器", 将要停梯 => "中间变量1"."1号梯将要停梯")
   END_RUNG
   // the same network as SCL:
   "1号梯高低速转换"(准备就绪 := "中间变量1"."1号梯准备就绪",   // "高低速转换"
              初始化低速运行 := "中间变量1"."1号梯初始化低速运行",
              当前楼层数 := "中间变量1"."1号梯当前楼层数",
              "1层上行呼梯按钮指示灯" := "中间变量2"."1层上呼分配1",
              "2层上行呼梯按钮指示灯" := "中间变量2"."2层上呼分配1",
              "3层上行呼梯按钮指示灯" := "中间变量2"."3层上呼分配1",
              "4层上行呼梯按钮指示灯" := "中间变量2"."4层上呼分配1",
              "5层上行呼梯按钮指示灯" := "中间变量2"."5层上呼分配1",
              "6层上行呼梯按钮指示灯" := "中间变量2"."6层上呼分配1",
              "7层上行呼梯按钮指示灯" := "中间变量2"."7层上呼分配1",
              "8层上行呼梯按钮指示灯" := "中间变量2"."8层上呼分配1",
              "9层上行呼梯按钮指示灯" := "中间变量2"."9层上呼分配1",
              "2层下行呼梯按钮指示灯" := "中间变量2"."2层下呼分配1",
              "3层下行呼梯按钮指示灯" := "中间变量2"."3层下呼分配1",
              "4层下行呼梯按钮指示灯" := "中间变量2"."4层下呼分配1",
              "5层下行呼梯按钮指示灯" := "中间变量2"."5层下呼分配1",
              "6层下行呼梯按钮指示灯" := "中间变量2"."6层下呼分配1",
              "7层下行呼梯按钮指示灯" := "中间变量2"."7层下呼分配1",
              "8层下行呼梯按钮指示灯" := "中间变量2"."8层下呼分配1",
              "9层下行呼梯按钮指示灯" := "中间变量2"."9层下呼分配1",
              "10层下行呼梯按钮指示灯" := "中间变量2"."10层下呼分配1",
              "1号梯1层按钮指示灯" := "输出"."1号梯1层按钮指示灯",
              "1号梯2层按钮指示灯" := "输出"."1号梯2层按钮指示灯",
              "1号梯3层按钮指示灯" := "输出"."1号梯3层按钮指示灯",
              "1号梯4层按钮指示灯" := "输出"."1号梯4层按钮指示灯",
              "1号梯5层按钮指示灯" := "输出"."1号梯5层按钮指示灯",
              "1号梯6层按钮指示灯" := "输出"."1号梯6层按钮指示灯",
              "1号梯7层按钮指示灯" := "输出"."1号梯7层按钮指示灯",
              "1号梯8层按钮指示灯" := "输出"."1号梯8层按钮指示灯",
              "1号梯9层按钮指示灯" := "输出"."1号梯9层按钮指示灯",
              "1号梯10层按钮指示灯" := "输出"."1号梯10层按钮指示灯",
              正处于故障中 := "中间变量1"."1号梯正处于故障中",
              "存在安全隐患（光幕）" := "中间变量1"."1号梯存在安全隐患（光幕）",
              "1号梯上行指示" := "输出"."1号梯上行指示",
              "1号梯下行指示" := "输出"."1号梯下行指示",
              "1号梯检修信号" := "输入"."1号梯检修信号",
              "1号梯上行接触器" := "输出"."1号梯上行接触器",
              "1号梯下行接触器" := "输出"."1号梯下行接触器",
              "1号梯外呼上面无目标2" := "中间变量2"."1号梯外呼上面无目标2",
              "1号梯外呼上面无目标3" := "中间变量2"."1号梯外呼上面无目标3",
              "1号梯外呼上面无目标4" := "中间变量2"."1号梯外呼上面无目标4",
              "1号梯外呼上面无目标5" := "中间变量2"."1号梯外呼上面无目标5",
              "1号梯外呼上面无目标6" := "中间变量2"."1号梯外呼上面无目标6",
              "1号梯外呼上面无目标7" := "中间变量2"."1号梯外呼上面无目标7",
              "1号梯外呼上面无目标8" := "中间变量2"."1号梯外呼上面无目标8",
              "1号梯外呼上面无目标9" := "中间变量2"."1号梯外呼上面无目标9",
              "1号梯外呼下面无目标2" := "中间变量2"."1号梯外呼下面无目标2",
              "1号梯外呼下面无目标3" := "中间变量2"."1号梯外呼下面无目标3",
              "1号梯外呼下面无目标4" := "中间变量2"."1号梯外呼下面无目标4",
              "1号梯外呼下面无目标5" := "中间变量2"."1号梯外呼下面无目标5",
              "1号梯外呼下面无目标6" := "中间变量2"."1号梯外呼下面无目标6",
              "1号梯外呼下面无目标7" := "中间变量2"."1号梯外呼下面无目标7",
              "1号梯外呼下面无目标8" := "中间变量2"."1号梯外呼下面无目标8",
              "1号梯外呼下面无目标9" := "中间变量2"."1号梯外呼下面无目标9",
              初始化高速运行 := "中间变量1"."1号梯高速初始化",
              "1号梯高速接触器" => "输出"."1号梯高速接触器",
              "1号梯低速接触器" => "输出"."1号梯低速接触器",
              将要停梯 => "中间变量1"."1号梯将要停梯");
END_REGION

REGION Network 2: 2号梯
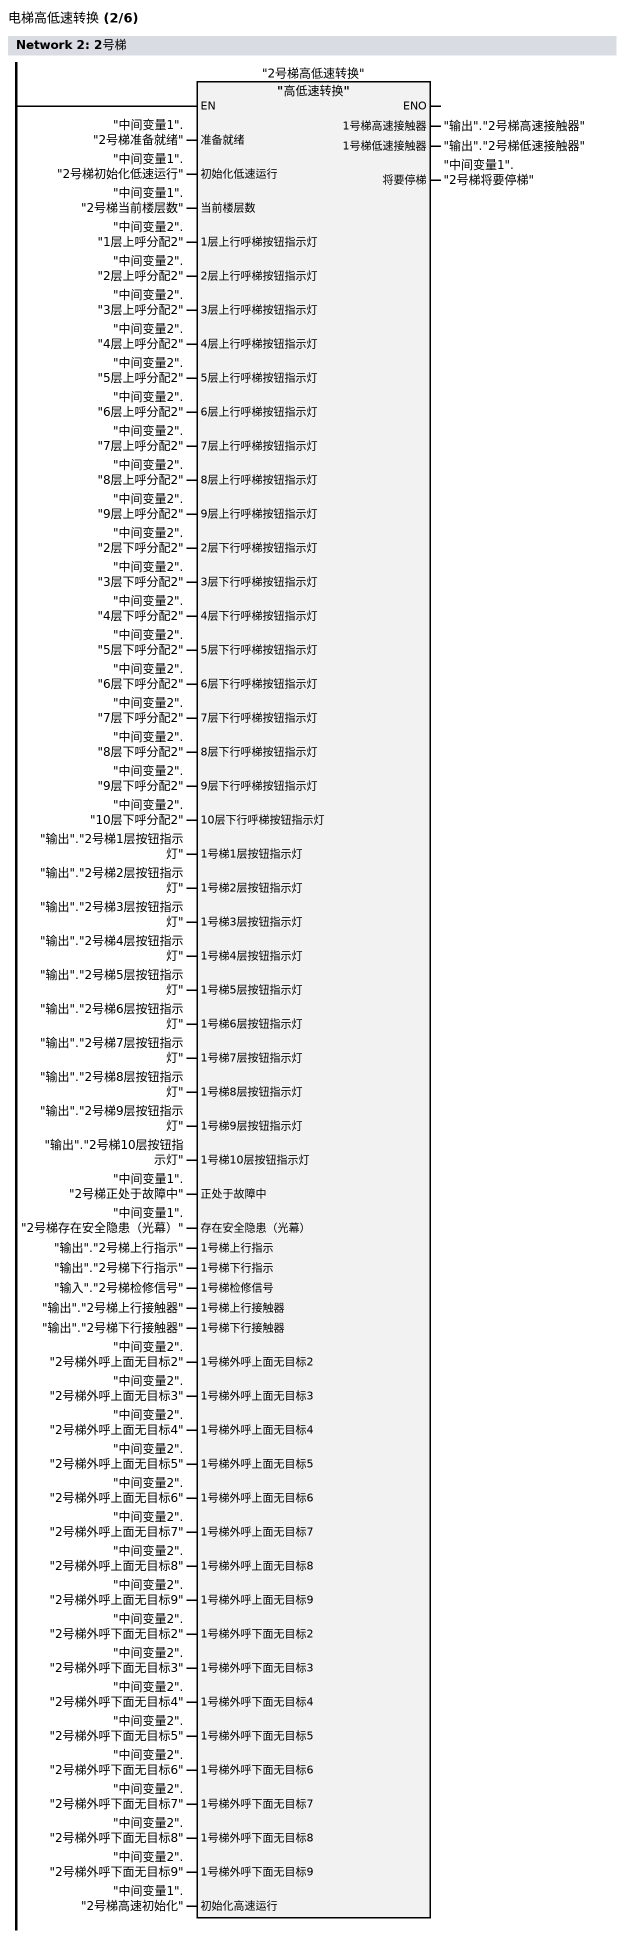
   RUNG wire#powerrail
      "2号梯高低速转换"(准备就绪 := "中间变量1"."2号梯准备就绪", 初始化低速运行 := "中间变量1"."2号梯初始化低速运行", 当前楼层数 := "中间变量1"."2号梯当前楼层数", "1层上行呼梯按钮指示灯" := "中间变量2"."1层上呼分配2", "2层上行呼梯按钮指示灯" := "中间变量2"."2层上呼分配2", "3层上行呼梯按钮指示灯" := "中间变量2"."3层上呼分配2", "4层上行呼梯按钮指示灯" := "中间变量2"."4层上呼分配2", "5层上行呼梯按钮指示灯" := "中间变量2"."5层上呼分配2", "6层上行呼梯按钮指示灯" := "中间变量2"."6层上呼分配2", "7层上行呼梯按钮指示灯" := "中间变量2"."7层上呼分配2", "8层上行呼梯按钮指示灯" := "中间变量2"."8层上呼分配2", "9层上行呼梯按钮指示灯" := "中间变量2"."9层上呼分配2", "2层下行呼梯按钮指示灯" := "中间变量2"."2层下呼分配2", "3层下行呼梯按钮指示灯" := "中间变量2"."3层下呼分配2", "4层下行呼梯按钮指示灯" := "中间变量2"."4层下呼分配2", "5层下行呼梯按钮指示灯" := "中间变量2"."5层下呼分配2", "6层下行呼梯按钮指示灯" := "中间变量2"."6层下呼分配2", "7层下行呼梯按钮指示灯" := "中间变量2"."7层下呼分配2", "8层下行呼梯按钮指示灯" := "中间变量2"."8层下呼分配2", "9层下行呼梯按钮指示灯" := "中间变量2"."9层下呼分配2", "10层下行呼梯按钮指示灯" := "中间变量2"."10层下呼分配2", "1号梯1层按钮指示灯" := "输出"."2号梯1层按钮指示灯", "1号梯2层按钮指示灯" := "输出"."2号梯2层按钮指示灯", "1号梯3层按钮指示灯" := "输出"."2号梯3层按钮指示灯", "1号梯4层按钮指示灯" := "输出"."2号梯4层按钮指示灯", "1号梯5层按钮指示灯" := "输出"."2号梯5层按钮指示灯", "1号梯6层按钮指示灯" := "输出"."2号梯6层按钮指示灯", "1号梯7层按钮指示灯" := "输出"."2号梯7层按钮指示灯", "1号梯8层按钮指示灯" := "输出"."2号梯8层按钮指示灯", "1号梯9层按钮指示灯" := "输出"."2号梯9层按钮指示灯", "1号梯10层按钮指示灯" := "输出"."2号梯10层按钮指示灯", 正处于故障中 := "中间变量1"."2号梯正处于故障中", "存在安全隐患（光幕）" := "中间变量1"."2号梯存在安全隐患（光幕）", "1号梯上行指示" := "输出"."2号梯上行指示", "1号梯下行指示" := "输出"."2号梯下行指示", "1号梯检修信号" := "输入"."2号梯检修信号", "1号梯上行接触器" := "输出"."2号梯上行接触器", "1号梯下行接触器" := "输出"."2号梯下行接触器", "1号梯外呼上面无目标2" := "中间变量2"."2号梯外呼上面无目标2", "1号梯外呼上面无目标3" := "中间变量2"."2号梯外呼上面无目标3", "1号梯外呼上面无目标4" := "中间变量2"."2号梯外呼上面无目标4", "1号梯外呼上面无目标5" := "中间变量2"."2号梯外呼上面无目标5", "1号梯外呼上面无目标6" := "中间变量2"."2号梯外呼上面无目标6", "1号梯外呼上面无目标7" := "中间变量2"."2号梯外呼上面无目标7", "1号梯外呼上面无目标8" := "中间变量2"."2号梯外呼上面无目标8", "1号梯外呼上面无目标9" := "中间变量2"."2号梯外呼上面无目标9", "1号梯外呼下面无目标2" := "中间变量2"."2号梯外呼下面无目标2", "1号梯外呼下面无目标3" := "中间变量2"."2号梯外呼下面无目标3", "1号梯外呼下面无目标4" := "中间变量2"."2号梯外呼下面无目标4", "1号梯外呼下面无目标5" := "中间变量2"."2号梯外呼下面无目标5", "1号梯外呼下面无目标6" := "中间变量2"."2号梯外呼下面无目标6", "1号梯外呼下面无目标7" := "中间变量2"."2号梯外呼下面无目标7", "1号梯外呼下面无目标8" := "中间变量2"."2号梯外呼下面无目标8", "1号梯外呼下面无目标9" := "中间变量2"."2号梯外呼下面无目标9", 初始化高速运行 := "中间变量1"."2号梯高速初始化", "1号梯高速接触器" => "输出"."2号梯高速接触器", "1号梯低速接触器" => "输出"."2号梯低速接触器", 将要停梯 => "中间变量1"."2号梯将要停梯")
   END_RUNG
   // the same network as SCL:
   "2号梯高低速转换"(准备就绪 := "中间变量1"."2号梯准备就绪",   // "高低速转换"
              初始化低速运行 := "中间变量1"."2号梯初始化低速运行",
              当前楼层数 := "中间变量1"."2号梯当前楼层数",
              "1层上行呼梯按钮指示灯" := "中间变量2"."1层上呼分配2",
              "2层上行呼梯按钮指示灯" := "中间变量2"."2层上呼分配2",
              "3层上行呼梯按钮指示灯" := "中间变量2"."3层上呼分配2",
              "4层上行呼梯按钮指示灯" := "中间变量2"."4层上呼分配2",
              "5层上行呼梯按钮指示灯" := "中间变量2"."5层上呼分配2",
              "6层上行呼梯按钮指示灯" := "中间变量2"."6层上呼分配2",
              "7层上行呼梯按钮指示灯" := "中间变量2"."7层上呼分配2",
              "8层上行呼梯按钮指示灯" := "中间变量2"."8层上呼分配2",
              "9层上行呼梯按钮指示灯" := "中间变量2"."9层上呼分配2",
              "2层下行呼梯按钮指示灯" := "中间变量2"."2层下呼分配2",
              "3层下行呼梯按钮指示灯" := "中间变量2"."3层下呼分配2",
              "4层下行呼梯按钮指示灯" := "中间变量2"."4层下呼分配2",
              "5层下行呼梯按钮指示灯" := "中间变量2"."5层下呼分配2",
              "6层下行呼梯按钮指示灯" := "中间变量2"."6层下呼分配2",
              "7层下行呼梯按钮指示灯" := "中间变量2"."7层下呼分配2",
              "8层下行呼梯按钮指示灯" := "中间变量2"."8层下呼分配2",
              "9层下行呼梯按钮指示灯" := "中间变量2"."9层下呼分配2",
              "10层下行呼梯按钮指示灯" := "中间变量2"."10层下呼分配2",
              "1号梯1层按钮指示灯" := "输出"."2号梯1层按钮指示灯",
              "1号梯2层按钮指示灯" := "输出"."2号梯2层按钮指示灯",
              "1号梯3层按钮指示灯" := "输出"."2号梯3层按钮指示灯",
              "1号梯4层按钮指示灯" := "输出"."2号梯4层按钮指示灯",
              "1号梯5层按钮指示灯" := "输出"."2号梯5层按钮指示灯",
              "1号梯6层按钮指示灯" := "输出"."2号梯6层按钮指示灯",
              "1号梯7层按钮指示灯" := "输出"."2号梯7层按钮指示灯",
              "1号梯8层按钮指示灯" := "输出"."2号梯8层按钮指示灯",
              "1号梯9层按钮指示灯" := "输出"."2号梯9层按钮指示灯",
              "1号梯10层按钮指示灯" := "输出"."2号梯10层按钮指示灯",
              正处于故障中 := "中间变量1"."2号梯正处于故障中",
              "存在安全隐患（光幕）" := "中间变量1"."2号梯存在安全隐患（光幕）",
              "1号梯上行指示" := "输出"."2号梯上行指示",
              "1号梯下行指示" := "输出"."2号梯下行指示",
              "1号梯检修信号" := "输入"."2号梯检修信号",
              "1号梯上行接触器" := "输出"."2号梯上行接触器",
              "1号梯下行接触器" := "输出"."2号梯下行接触器",
              "1号梯外呼上面无目标2" := "中间变量2"."2号梯外呼上面无目标2",
              "1号梯外呼上面无目标3" := "中间变量2"."2号梯外呼上面无目标3",
              "1号梯外呼上面无目标4" := "中间变量2"."2号梯外呼上面无目标4",
              "1号梯外呼上面无目标5" := "中间变量2"."2号梯外呼上面无目标5",
              "1号梯外呼上面无目标6" := "中间变量2"."2号梯外呼上面无目标6",
              "1号梯外呼上面无目标7" := "中间变量2"."2号梯外呼上面无目标7",
              "1号梯外呼上面无目标8" := "中间变量2"."2号梯外呼上面无目标8",
              "1号梯外呼上面无目标9" := "中间变量2"."2号梯外呼上面无目标9",
              "1号梯外呼下面无目标2" := "中间变量2"."2号梯外呼下面无目标2",
              "1号梯外呼下面无目标3" := "中间变量2"."2号梯外呼下面无目标3",
              "1号梯外呼下面无目标4" := "中间变量2"."2号梯外呼下面无目标4",
              "1号梯外呼下面无目标5" := "中间变量2"."2号梯外呼下面无目标5",
              "1号梯外呼下面无目标6" := "中间变量2"."2号梯外呼下面无目标6",
              "1号梯外呼下面无目标7" := "中间变量2"."2号梯外呼下面无目标7",
              "1号梯外呼下面无目标8" := "中间变量2"."2号梯外呼下面无目标8",
              "1号梯外呼下面无目标9" := "中间变量2"."2号梯外呼下面无目标9",
              初始化高速运行 := "中间变量1"."2号梯高速初始化",
              "1号梯高速接触器" => "输出"."2号梯高速接触器",
              "1号梯低速接触器" => "输出"."2号梯低速接触器",
              将要停梯 => "中间变量1"."2号梯将要停梯");
END_REGION

REGION Network 3: 3号梯
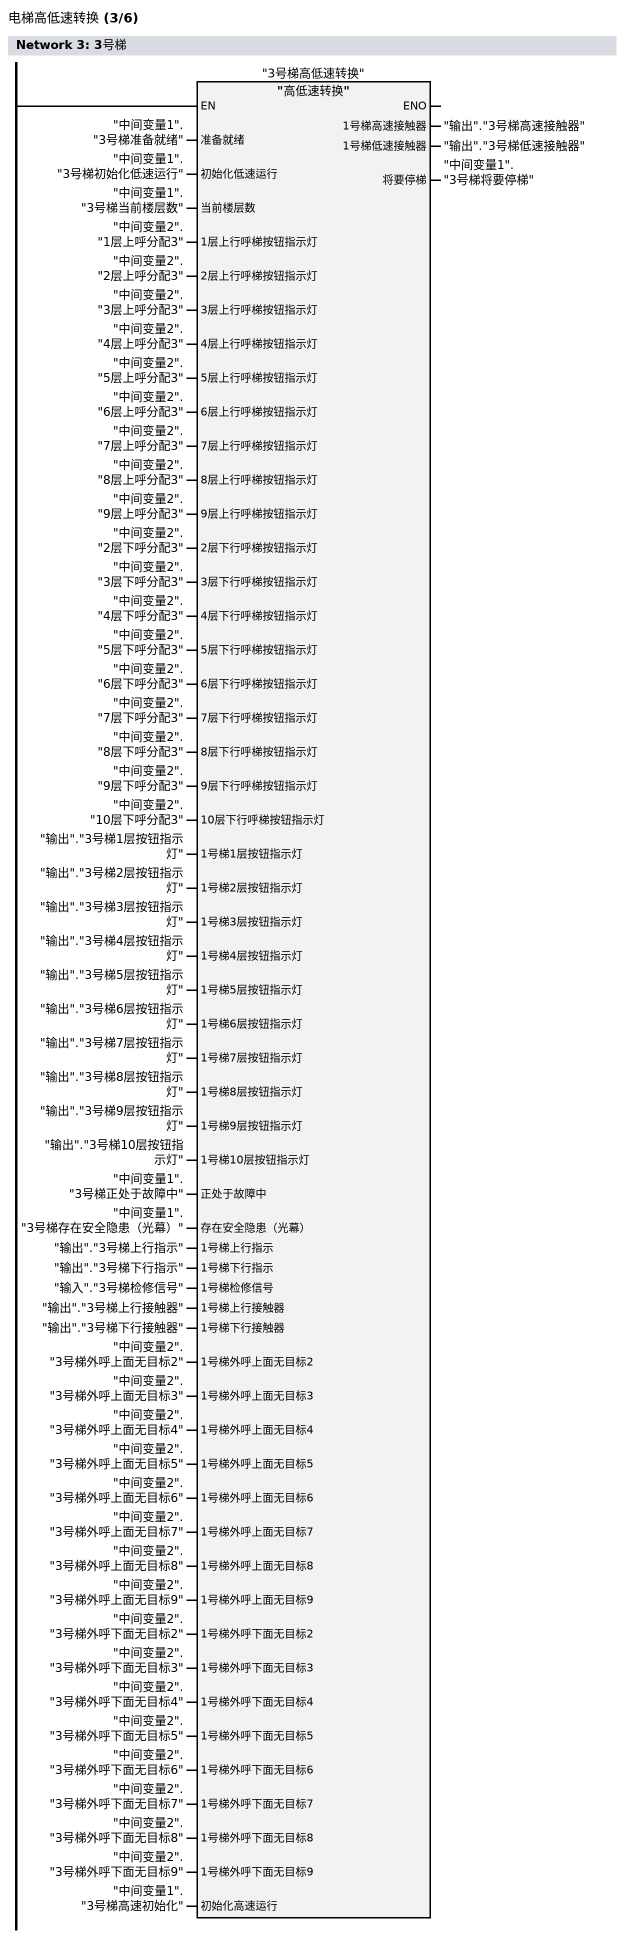
   RUNG wire#powerrail
      "3号梯高低速转换"(准备就绪 := "中间变量1"."3号梯准备就绪", 初始化低速运行 := "中间变量1"."3号梯初始化低速运行", 当前楼层数 := "中间变量1"."3号梯当前楼层数", "1层上行呼梯按钮指示灯" := "中间变量2"."1层上呼分配3", "2层上行呼梯按钮指示灯" := "中间变量2"."2层上呼分配3", "3层上行呼梯按钮指示灯" := "中间变量2"."3层上呼分配3", "4层上行呼梯按钮指示灯" := "中间变量2"."4层上呼分配3", "5层上行呼梯按钮指示灯" := "中间变量2"."5层上呼分配3", "6层上行呼梯按钮指示灯" := "中间变量2"."6层上呼分配3", "7层上行呼梯按钮指示灯" := "中间变量2"."7层上呼分配3", "8层上行呼梯按钮指示灯" := "中间变量2"."8层上呼分配3", "9层上行呼梯按钮指示灯" := "中间变量2"."9层上呼分配3", "2层下行呼梯按钮指示灯" := "中间变量2"."2层下呼分配3", "3层下行呼梯按钮指示灯" := "中间变量2"."3层下呼分配3", "4层下行呼梯按钮指示灯" := "中间变量2"."4层下呼分配3", "5层下行呼梯按钮指示灯" := "中间变量2"."5层下呼分配3", "6层下行呼梯按钮指示灯" := "中间变量2"."6层下呼分配3", "7层下行呼梯按钮指示灯" := "中间变量2"."7层下呼分配3", "8层下行呼梯按钮指示灯" := "中间变量2"."8层下呼分配3", "9层下行呼梯按钮指示灯" := "中间变量2"."9层下呼分配3", "10层下行呼梯按钮指示灯" := "中间变量2"."10层下呼分配3", "1号梯1层按钮指示灯" := "输出"."3号梯1层按钮指示灯", "1号梯2层按钮指示灯" := "输出"."3号梯2层按钮指示灯", "1号梯3层按钮指示灯" := "输出"."3号梯3层按钮指示灯", "1号梯4层按钮指示灯" := "输出"."3号梯4层按钮指示灯", "1号梯5层按钮指示灯" := "输出"."3号梯5层按钮指示灯", "1号梯6层按钮指示灯" := "输出"."3号梯6层按钮指示灯", "1号梯7层按钮指示灯" := "输出"."3号梯7层按钮指示灯", "1号梯8层按钮指示灯" := "输出"."3号梯8层按钮指示灯", "1号梯9层按钮指示灯" := "输出"."3号梯9层按钮指示灯", "1号梯10层按钮指示灯" := "输出"."3号梯10层按钮指示灯", 正处于故障中 := "中间变量1"."3号梯正处于故障中", "存在安全隐患（光幕）" := "中间变量1"."3号梯存在安全隐患（光幕）", "1号梯上行指示" := "输出"."3号梯上行指示", "1号梯下行指示" := "输出"."3号梯下行指示", "1号梯检修信号" := "输入"."3号梯检修信号", "1号梯上行接触器" := "输出"."3号梯上行接触器", "1号梯下行接触器" := "输出"."3号梯下行接触器", "1号梯外呼上面无目标2" := "中间变量2"."3号梯外呼上面无目标2", "1号梯外呼上面无目标3" := "中间变量2"."3号梯外呼上面无目标3", "1号梯外呼上面无目标4" := "中间变量2"."3号梯外呼上面无目标4", "1号梯外呼上面无目标5" := "中间变量2"."3号梯外呼上面无目标5", "1号梯外呼上面无目标6" := "中间变量2"."3号梯外呼上面无目标6", "1号梯外呼上面无目标7" := "中间变量2"."3号梯外呼上面无目标7", "1号梯外呼上面无目标8" := "中间变量2"."3号梯外呼上面无目标8", "1号梯外呼上面无目标9" := "中间变量2"."3号梯外呼上面无目标9", "1号梯外呼下面无目标2" := "中间变量2"."3号梯外呼下面无目标2", "1号梯外呼下面无目标3" := "中间变量2"."3号梯外呼下面无目标3", "1号梯外呼下面无目标4" := "中间变量2"."3号梯外呼下面无目标4", "1号梯外呼下面无目标5" := "中间变量2"."3号梯外呼下面无目标5", "1号梯外呼下面无目标6" := "中间变量2"."3号梯外呼下面无目标6", "1号梯外呼下面无目标7" := "中间变量2"."3号梯外呼下面无目标7", "1号梯外呼下面无目标8" := "中间变量2"."3号梯外呼下面无目标8", "1号梯外呼下面无目标9" := "中间变量2"."3号梯外呼下面无目标9", 初始化高速运行 := "中间变量1"."3号梯高速初始化", "1号梯高速接触器" => "输出"."3号梯高速接触器", "1号梯低速接触器" => "输出"."3号梯低速接触器", 将要停梯 => "中间变量1"."3号梯将要停梯")
   END_RUNG
   // the same network as SCL:
   "3号梯高低速转换"(准备就绪 := "中间变量1"."3号梯准备就绪",   // "高低速转换"
              初始化低速运行 := "中间变量1"."3号梯初始化低速运行",
              当前楼层数 := "中间变量1"."3号梯当前楼层数",
              "1层上行呼梯按钮指示灯" := "中间变量2"."1层上呼分配3",
              "2层上行呼梯按钮指示灯" := "中间变量2"."2层上呼分配3",
              "3层上行呼梯按钮指示灯" := "中间变量2"."3层上呼分配3",
              "4层上行呼梯按钮指示灯" := "中间变量2"."4层上呼分配3",
              "5层上行呼梯按钮指示灯" := "中间变量2"."5层上呼分配3",
              "6层上行呼梯按钮指示灯" := "中间变量2"."6层上呼分配3",
              "7层上行呼梯按钮指示灯" := "中间变量2"."7层上呼分配3",
              "8层上行呼梯按钮指示灯" := "中间变量2"."8层上呼分配3",
              "9层上行呼梯按钮指示灯" := "中间变量2"."9层上呼分配3",
              "2层下行呼梯按钮指示灯" := "中间变量2"."2层下呼分配3",
              "3层下行呼梯按钮指示灯" := "中间变量2"."3层下呼分配3",
              "4层下行呼梯按钮指示灯" := "中间变量2"."4层下呼分配3",
              "5层下行呼梯按钮指示灯" := "中间变量2"."5层下呼分配3",
              "6层下行呼梯按钮指示灯" := "中间变量2"."6层下呼分配3",
              "7层下行呼梯按钮指示灯" := "中间变量2"."7层下呼分配3",
              "8层下行呼梯按钮指示灯" := "中间变量2"."8层下呼分配3",
              "9层下行呼梯按钮指示灯" := "中间变量2"."9层下呼分配3",
              "10层下行呼梯按钮指示灯" := "中间变量2"."10层下呼分配3",
              "1号梯1层按钮指示灯" := "输出"."3号梯1层按钮指示灯",
              "1号梯2层按钮指示灯" := "输出"."3号梯2层按钮指示灯",
              "1号梯3层按钮指示灯" := "输出"."3号梯3层按钮指示灯",
              "1号梯4层按钮指示灯" := "输出"."3号梯4层按钮指示灯",
              "1号梯5层按钮指示灯" := "输出"."3号梯5层按钮指示灯",
              "1号梯6层按钮指示灯" := "输出"."3号梯6层按钮指示灯",
              "1号梯7层按钮指示灯" := "输出"."3号梯7层按钮指示灯",
              "1号梯8层按钮指示灯" := "输出"."3号梯8层按钮指示灯",
              "1号梯9层按钮指示灯" := "输出"."3号梯9层按钮指示灯",
              "1号梯10层按钮指示灯" := "输出"."3号梯10层按钮指示灯",
              正处于故障中 := "中间变量1"."3号梯正处于故障中",
              "存在安全隐患（光幕）" := "中间变量1"."3号梯存在安全隐患（光幕）",
              "1号梯上行指示" := "输出"."3号梯上行指示",
              "1号梯下行指示" := "输出"."3号梯下行指示",
              "1号梯检修信号" := "输入"."3号梯检修信号",
              "1号梯上行接触器" := "输出"."3号梯上行接触器",
              "1号梯下行接触器" := "输出"."3号梯下行接触器",
              "1号梯外呼上面无目标2" := "中间变量2"."3号梯外呼上面无目标2",
              "1号梯外呼上面无目标3" := "中间变量2"."3号梯外呼上面无目标3",
              "1号梯外呼上面无目标4" := "中间变量2"."3号梯外呼上面无目标4",
              "1号梯外呼上面无目标5" := "中间变量2"."3号梯外呼上面无目标5",
              "1号梯外呼上面无目标6" := "中间变量2"."3号梯外呼上面无目标6",
              "1号梯外呼上面无目标7" := "中间变量2"."3号梯外呼上面无目标7",
              "1号梯外呼上面无目标8" := "中间变量2"."3号梯外呼上面无目标8",
              "1号梯外呼上面无目标9" := "中间变量2"."3号梯外呼上面无目标9",
              "1号梯外呼下面无目标2" := "中间变量2"."3号梯外呼下面无目标2",
              "1号梯外呼下面无目标3" := "中间变量2"."3号梯外呼下面无目标3",
              "1号梯外呼下面无目标4" := "中间变量2"."3号梯外呼下面无目标4",
              "1号梯外呼下面无目标5" := "中间变量2"."3号梯外呼下面无目标5",
              "1号梯外呼下面无目标6" := "中间变量2"."3号梯外呼下面无目标6",
              "1号梯外呼下面无目标7" := "中间变量2"."3号梯外呼下面无目标7",
              "1号梯外呼下面无目标8" := "中间变量2"."3号梯外呼下面无目标8",
              "1号梯外呼下面无目标9" := "中间变量2"."3号梯外呼下面无目标9",
              初始化高速运行 := "中间变量1"."3号梯高速初始化",
              "1号梯高速接触器" => "输出"."3号梯高速接触器",
              "1号梯低速接触器" => "输出"."3号梯低速接触器",
              将要停梯 => "中间变量1"."3号梯将要停梯");
END_REGION

REGION Network 4: 4号梯
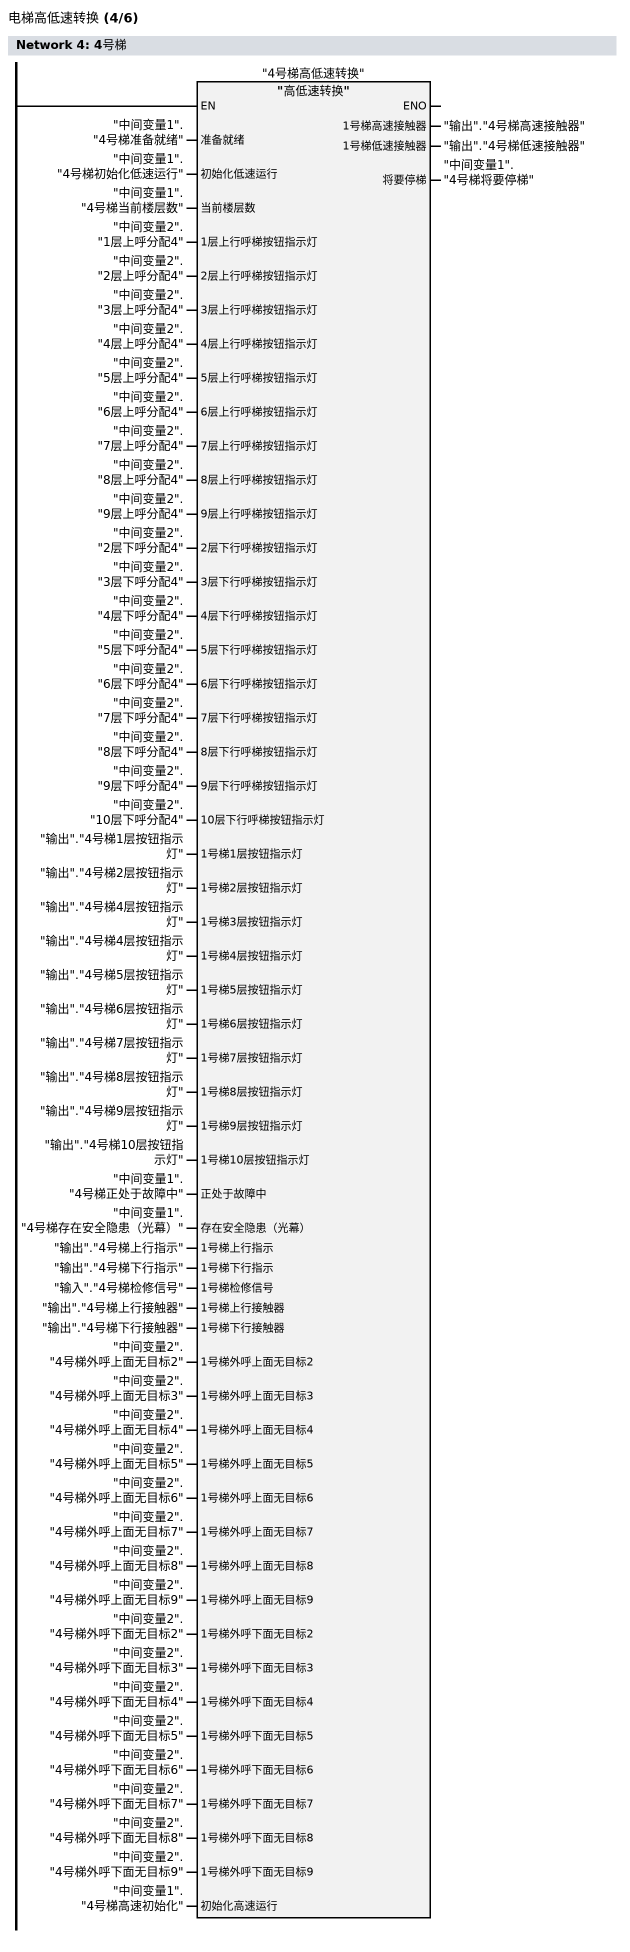
   RUNG wire#powerrail
      "4号梯高低速转换"(准备就绪 := "中间变量1"."4号梯准备就绪", 初始化低速运行 := "中间变量1"."4号梯初始化低速运行", 当前楼层数 := "中间变量1"."4号梯当前楼层数", "1层上行呼梯按钮指示灯" := "中间变量2"."1层上呼分配4", "2层上行呼梯按钮指示灯" := "中间变量2"."2层上呼分配4", "3层上行呼梯按钮指示灯" := "中间变量2"."3层上呼分配4", "4层上行呼梯按钮指示灯" := "中间变量2"."4层上呼分配4", "5层上行呼梯按钮指示灯" := "中间变量2"."5层上呼分配4", "6层上行呼梯按钮指示灯" := "中间变量2"."6层上呼分配4", "7层上行呼梯按钮指示灯" := "中间变量2"."7层上呼分配4", "8层上行呼梯按钮指示灯" := "中间变量2"."8层上呼分配4", "9层上行呼梯按钮指示灯" := "中间变量2"."9层上呼分配4", "2层下行呼梯按钮指示灯" := "中间变量2"."2层下呼分配4", "3层下行呼梯按钮指示灯" := "中间变量2"."3层下呼分配4", "4层下行呼梯按钮指示灯" := "中间变量2"."4层下呼分配4", "5层下行呼梯按钮指示灯" := "中间变量2"."5层下呼分配4", "6层下行呼梯按钮指示灯" := "中间变量2"."6层下呼分配4", "7层下行呼梯按钮指示灯" := "中间变量2"."7层下呼分配4", "8层下行呼梯按钮指示灯" := "中间变量2"."8层下呼分配4", "9层下行呼梯按钮指示灯" := "中间变量2"."9层下呼分配4", "10层下行呼梯按钮指示灯" := "中间变量2"."10层下呼分配4", "1号梯1层按钮指示灯" := "输出"."4号梯1层按钮指示灯", "1号梯2层按钮指示灯" := "输出"."4号梯2层按钮指示灯", "1号梯3层按钮指示灯" := "输出"."4号梯4层按钮指示灯", "1号梯4层按钮指示灯" := "输出"."4号梯4层按钮指示灯", "1号梯5层按钮指示灯" := "输出"."4号梯5层按钮指示灯", "1号梯6层按钮指示灯" := "输出"."4号梯6层按钮指示灯", "1号梯7层按钮指示灯" := "输出"."4号梯7层按钮指示灯", "1号梯8层按钮指示灯" := "输出"."4号梯8层按钮指示灯", "1号梯9层按钮指示灯" := "输出"."4号梯9层按钮指示灯", "1号梯10层按钮指示灯" := "输出"."4号梯10层按钮指示灯", 正处于故障中 := "中间变量1"."4号梯正处于故障中", "存在安全隐患（光幕）" := "中间变量1"."4号梯存在安全隐患（光幕）", "1号梯上行指示" := "输出"."4号梯上行指示", "1号梯下行指示" := "输出"."4号梯下行指示", "1号梯检修信号" := "输入"."4号梯检修信号", "1号梯上行接触器" := "输出"."4号梯上行接触器", "1号梯下行接触器" := "输出"."4号梯下行接触器", "1号梯外呼上面无目标2" := "中间变量2"."4号梯外呼上面无目标2", "1号梯外呼上面无目标3" := "中间变量2"."4号梯外呼上面无目标3", "1号梯外呼上面无目标4" := "中间变量2"."4号梯外呼上面无目标4", "1号梯外呼上面无目标5" := "中间变量2"."4号梯外呼上面无目标5", "1号梯外呼上面无目标6" := "中间变量2"."4号梯外呼上面无目标6", "1号梯外呼上面无目标7" := "中间变量2"."4号梯外呼上面无目标7", "1号梯外呼上面无目标8" := "中间变量2"."4号梯外呼上面无目标8", "1号梯外呼上面无目标9" := "中间变量2"."4号梯外呼上面无目标9", "1号梯外呼下面无目标2" := "中间变量2"."4号梯外呼下面无目标2", "1号梯外呼下面无目标3" := "中间变量2"."4号梯外呼下面无目标3", "1号梯外呼下面无目标4" := "中间变量2"."4号梯外呼下面无目标4", "1号梯外呼下面无目标5" := "中间变量2"."4号梯外呼下面无目标5", "1号梯外呼下面无目标6" := "中间变量2"."4号梯外呼下面无目标6", "1号梯外呼下面无目标7" := "中间变量2"."4号梯外呼下面无目标7", "1号梯外呼下面无目标8" := "中间变量2"."4号梯外呼下面无目标8", "1号梯外呼下面无目标9" := "中间变量2"."4号梯外呼下面无目标9", 初始化高速运行 := "中间变量1"."4号梯高速初始化", "1号梯高速接触器" => "输出"."4号梯高速接触器", "1号梯低速接触器" => "输出"."4号梯低速接触器", 将要停梯 => "中间变量1"."4号梯将要停梯")
   END_RUNG
   // the same network as SCL:
   "4号梯高低速转换"(准备就绪 := "中间变量1"."4号梯准备就绪",   // "高低速转换"
              初始化低速运行 := "中间变量1"."4号梯初始化低速运行",
              当前楼层数 := "中间变量1"."4号梯当前楼层数",
              "1层上行呼梯按钮指示灯" := "中间变量2"."1层上呼分配4",
              "2层上行呼梯按钮指示灯" := "中间变量2"."2层上呼分配4",
              "3层上行呼梯按钮指示灯" := "中间变量2"."3层上呼分配4",
              "4层上行呼梯按钮指示灯" := "中间变量2"."4层上呼分配4",
              "5层上行呼梯按钮指示灯" := "中间变量2"."5层上呼分配4",
              "6层上行呼梯按钮指示灯" := "中间变量2"."6层上呼分配4",
              "7层上行呼梯按钮指示灯" := "中间变量2"."7层上呼分配4",
              "8层上行呼梯按钮指示灯" := "中间变量2"."8层上呼分配4",
              "9层上行呼梯按钮指示灯" := "中间变量2"."9层上呼分配4",
              "2层下行呼梯按钮指示灯" := "中间变量2"."2层下呼分配4",
              "3层下行呼梯按钮指示灯" := "中间变量2"."3层下呼分配4",
              "4层下行呼梯按钮指示灯" := "中间变量2"."4层下呼分配4",
              "5层下行呼梯按钮指示灯" := "中间变量2"."5层下呼分配4",
              "6层下行呼梯按钮指示灯" := "中间变量2"."6层下呼分配4",
              "7层下行呼梯按钮指示灯" := "中间变量2"."7层下呼分配4",
              "8层下行呼梯按钮指示灯" := "中间变量2"."8层下呼分配4",
              "9层下行呼梯按钮指示灯" := "中间变量2"."9层下呼分配4",
              "10层下行呼梯按钮指示灯" := "中间变量2"."10层下呼分配4",
              "1号梯1层按钮指示灯" := "输出"."4号梯1层按钮指示灯",
              "1号梯2层按钮指示灯" := "输出"."4号梯2层按钮指示灯",
              "1号梯3层按钮指示灯" := "输出"."4号梯4层按钮指示灯",
              "1号梯4层按钮指示灯" := "输出"."4号梯4层按钮指示灯",
              "1号梯5层按钮指示灯" := "输出"."4号梯5层按钮指示灯",
              "1号梯6层按钮指示灯" := "输出"."4号梯6层按钮指示灯",
              "1号梯7层按钮指示灯" := "输出"."4号梯7层按钮指示灯",
              "1号梯8层按钮指示灯" := "输出"."4号梯8层按钮指示灯",
              "1号梯9层按钮指示灯" := "输出"."4号梯9层按钮指示灯",
              "1号梯10层按钮指示灯" := "输出"."4号梯10层按钮指示灯",
              正处于故障中 := "中间变量1"."4号梯正处于故障中",
              "存在安全隐患（光幕）" := "中间变量1"."4号梯存在安全隐患（光幕）",
              "1号梯上行指示" := "输出"."4号梯上行指示",
              "1号梯下行指示" := "输出"."4号梯下行指示",
              "1号梯检修信号" := "输入"."4号梯检修信号",
              "1号梯上行接触器" := "输出"."4号梯上行接触器",
              "1号梯下行接触器" := "输出"."4号梯下行接触器",
              "1号梯外呼上面无目标2" := "中间变量2"."4号梯外呼上面无目标2",
              "1号梯外呼上面无目标3" := "中间变量2"."4号梯外呼上面无目标3",
              "1号梯外呼上面无目标4" := "中间变量2"."4号梯外呼上面无目标4",
              "1号梯外呼上面无目标5" := "中间变量2"."4号梯外呼上面无目标5",
              "1号梯外呼上面无目标6" := "中间变量2"."4号梯外呼上面无目标6",
              "1号梯外呼上面无目标7" := "中间变量2"."4号梯外呼上面无目标7",
              "1号梯外呼上面无目标8" := "中间变量2"."4号梯外呼上面无目标8",
              "1号梯外呼上面无目标9" := "中间变量2"."4号梯外呼上面无目标9",
              "1号梯外呼下面无目标2" := "中间变量2"."4号梯外呼下面无目标2",
              "1号梯外呼下面无目标3" := "中间变量2"."4号梯外呼下面无目标3",
              "1号梯外呼下面无目标4" := "中间变量2"."4号梯外呼下面无目标4",
              "1号梯外呼下面无目标5" := "中间变量2"."4号梯外呼下面无目标5",
              "1号梯外呼下面无目标6" := "中间变量2"."4号梯外呼下面无目标6",
              "1号梯外呼下面无目标7" := "中间变量2"."4号梯外呼下面无目标7",
              "1号梯外呼下面无目标8" := "中间变量2"."4号梯外呼下面无目标8",
              "1号梯外呼下面无目标9" := "中间变量2"."4号梯外呼下面无目标9",
              初始化高速运行 := "中间变量1"."4号梯高速初始化",
              "1号梯高速接触器" => "输出"."4号梯高速接触器",
              "1号梯低速接触器" => "输出"."4号梯低速接触器",
              将要停梯 => "中间变量1"."4号梯将要停梯");
END_REGION

REGION Network 5: 5号梯
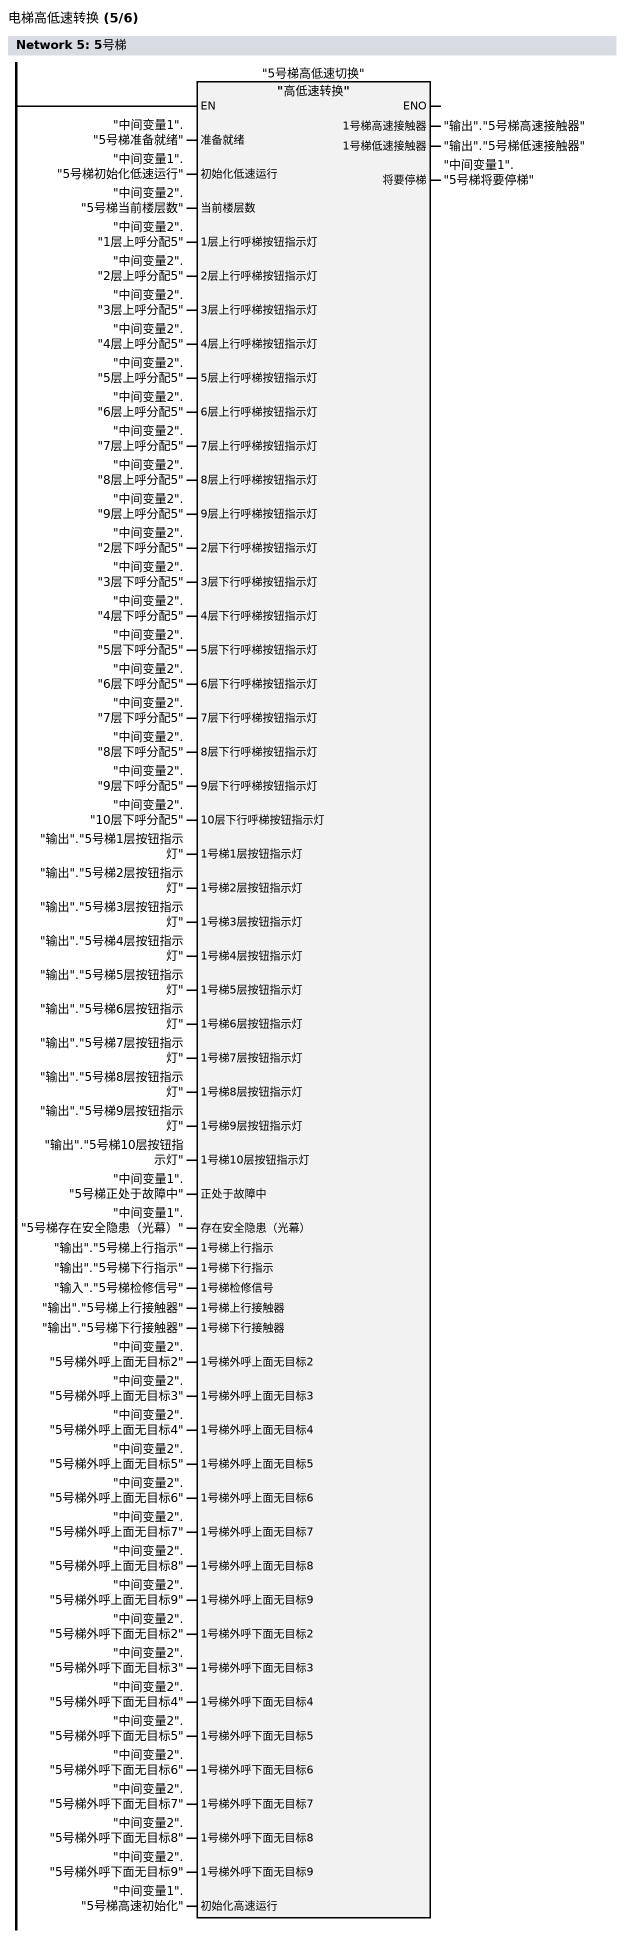
   RUNG wire#powerrail
      "5号梯高低速切换"(准备就绪 := "中间变量1"."5号梯准备就绪", 初始化低速运行 := "中间变量1"."5号梯初始化低速运行", 当前楼层数 := "中间变量2"."5号梯当前楼层数", "1层上行呼梯按钮指示灯" := "中间变量2"."1层上呼分配5", "2层上行呼梯按钮指示灯" := "中间变量2"."2层上呼分配5", "3层上行呼梯按钮指示灯" := "中间变量2"."3层上呼分配5", "4层上行呼梯按钮指示灯" := "中间变量2"."4层上呼分配5", "5层上行呼梯按钮指示灯" := "中间变量2"."5层上呼分配5", "6层上行呼梯按钮指示灯" := "中间变量2"."6层上呼分配5", "7层上行呼梯按钮指示灯" := "中间变量2"."7层上呼分配5", "8层上行呼梯按钮指示灯" := "中间变量2"."8层上呼分配5", "9层上行呼梯按钮指示灯" := "中间变量2"."9层上呼分配5", "2层下行呼梯按钮指示灯" := "中间变量2"."2层下呼分配5", "3层下行呼梯按钮指示灯" := "中间变量2"."3层下呼分配5", "4层下行呼梯按钮指示灯" := "中间变量2"."4层下呼分配5", "5层下行呼梯按钮指示灯" := "中间变量2"."5层下呼分配5", "6层下行呼梯按钮指示灯" := "中间变量2"."6层下呼分配5", "7层下行呼梯按钮指示灯" := "中间变量2"."7层下呼分配5", "8层下行呼梯按钮指示灯" := "中间变量2"."8层下呼分配5", "9层下行呼梯按钮指示灯" := "中间变量2"."9层下呼分配5", "10层下行呼梯按钮指示灯" := "中间变量2"."10层下呼分配5", "1号梯1层按钮指示灯" := "输出"."5号梯1层按钮指示灯", "1号梯2层按钮指示灯" := "输出"."5号梯2层按钮指示灯", "1号梯3层按钮指示灯" := "输出"."5号梯3层按钮指示灯", "1号梯4层按钮指示灯" := "输出"."5号梯4层按钮指示灯", "1号梯5层按钮指示灯" := "输出"."5号梯5层按钮指示灯", "1号梯6层按钮指示灯" := "输出"."5号梯6层按钮指示灯", "1号梯7层按钮指示灯" := "输出"."5号梯7层按钮指示灯", "1号梯8层按钮指示灯" := "输出"."5号梯8层按钮指示灯", "1号梯9层按钮指示灯" := "输出"."5号梯9层按钮指示灯", "1号梯10层按钮指示灯" := "输出"."5号梯10层按钮指示灯", 正处于故障中 := "中间变量1"."5号梯正处于故障中", "存在安全隐患（光幕）" := "中间变量1"."5号梯存在安全隐患（光幕）", "1号梯上行指示" := "输出"."5号梯上行指示", "1号梯下行指示" := "输出"."5号梯下行指示", "1号梯检修信号" := "输入"."5号梯检修信号", "1号梯上行接触器" := "输出"."5号梯上行接触器", "1号梯下行接触器" := "输出"."5号梯下行接触器", "1号梯外呼上面无目标2" := "中间变量2"."5号梯外呼上面无目标2", "1号梯外呼上面无目标3" := "中间变量2"."5号梯外呼上面无目标3", "1号梯外呼上面无目标4" := "中间变量2"."5号梯外呼上面无目标4", "1号梯外呼上面无目标5" := "中间变量2"."5号梯外呼上面无目标5", "1号梯外呼上面无目标6" := "中间变量2"."5号梯外呼上面无目标6", "1号梯外呼上面无目标7" := "中间变量2"."5号梯外呼上面无目标7", "1号梯外呼上面无目标8" := "中间变量2"."5号梯外呼上面无目标8", "1号梯外呼上面无目标9" := "中间变量2"."5号梯外呼上面无目标9", "1号梯外呼下面无目标2" := "中间变量2"."5号梯外呼下面无目标2", "1号梯外呼下面无目标3" := "中间变量2"."5号梯外呼下面无目标3", "1号梯外呼下面无目标4" := "中间变量2"."5号梯外呼下面无目标4", "1号梯外呼下面无目标5" := "中间变量2"."5号梯外呼下面无目标5", "1号梯外呼下面无目标6" := "中间变量2"."5号梯外呼下面无目标6", "1号梯外呼下面无目标7" := "中间变量2"."5号梯外呼下面无目标7", "1号梯外呼下面无目标8" := "中间变量2"."5号梯外呼下面无目标8", "1号梯外呼下面无目标9" := "中间变量2"."5号梯外呼下面无目标9", 初始化高速运行 := "中间变量1"."5号梯高速初始化", "1号梯高速接触器" => "输出"."5号梯高速接触器", "1号梯低速接触器" => "输出"."5号梯低速接触器", 将要停梯 => "中间变量1"."5号梯将要停梯")
   END_RUNG
   // the same network as SCL:
   "5号梯高低速切换"(准备就绪 := "中间变量1"."5号梯准备就绪",   // "高低速转换"
              初始化低速运行 := "中间变量1"."5号梯初始化低速运行",
              当前楼层数 := "中间变量2"."5号梯当前楼层数",
              "1层上行呼梯按钮指示灯" := "中间变量2"."1层上呼分配5",
              "2层上行呼梯按钮指示灯" := "中间变量2"."2层上呼分配5",
              "3层上行呼梯按钮指示灯" := "中间变量2"."3层上呼分配5",
              "4层上行呼梯按钮指示灯" := "中间变量2"."4层上呼分配5",
              "5层上行呼梯按钮指示灯" := "中间变量2"."5层上呼分配5",
              "6层上行呼梯按钮指示灯" := "中间变量2"."6层上呼分配5",
              "7层上行呼梯按钮指示灯" := "中间变量2"."7层上呼分配5",
              "8层上行呼梯按钮指示灯" := "中间变量2"."8层上呼分配5",
              "9层上行呼梯按钮指示灯" := "中间变量2"."9层上呼分配5",
              "2层下行呼梯按钮指示灯" := "中间变量2"."2层下呼分配5",
              "3层下行呼梯按钮指示灯" := "中间变量2"."3层下呼分配5",
              "4层下行呼梯按钮指示灯" := "中间变量2"."4层下呼分配5",
              "5层下行呼梯按钮指示灯" := "中间变量2"."5层下呼分配5",
              "6层下行呼梯按钮指示灯" := "中间变量2"."6层下呼分配5",
              "7层下行呼梯按钮指示灯" := "中间变量2"."7层下呼分配5",
              "8层下行呼梯按钮指示灯" := "中间变量2"."8层下呼分配5",
              "9层下行呼梯按钮指示灯" := "中间变量2"."9层下呼分配5",
              "10层下行呼梯按钮指示灯" := "中间变量2"."10层下呼分配5",
              "1号梯1层按钮指示灯" := "输出"."5号梯1层按钮指示灯",
              "1号梯2层按钮指示灯" := "输出"."5号梯2层按钮指示灯",
              "1号梯3层按钮指示灯" := "输出"."5号梯3层按钮指示灯",
              "1号梯4层按钮指示灯" := "输出"."5号梯4层按钮指示灯",
              "1号梯5层按钮指示灯" := "输出"."5号梯5层按钮指示灯",
              "1号梯6层按钮指示灯" := "输出"."5号梯6层按钮指示灯",
              "1号梯7层按钮指示灯" := "输出"."5号梯7层按钮指示灯",
              "1号梯8层按钮指示灯" := "输出"."5号梯8层按钮指示灯",
              "1号梯9层按钮指示灯" := "输出"."5号梯9层按钮指示灯",
              "1号梯10层按钮指示灯" := "输出"."5号梯10层按钮指示灯",
              正处于故障中 := "中间变量1"."5号梯正处于故障中",
              "存在安全隐患（光幕）" := "中间变量1"."5号梯存在安全隐患（光幕）",
              "1号梯上行指示" := "输出"."5号梯上行指示",
              "1号梯下行指示" := "输出"."5号梯下行指示",
              "1号梯检修信号" := "输入"."5号梯检修信号",
              "1号梯上行接触器" := "输出"."5号梯上行接触器",
              "1号梯下行接触器" := "输出"."5号梯下行接触器",
              "1号梯外呼上面无目标2" := "中间变量2"."5号梯外呼上面无目标2",
              "1号梯外呼上面无目标3" := "中间变量2"."5号梯外呼上面无目标3",
              "1号梯外呼上面无目标4" := "中间变量2"."5号梯外呼上面无目标4",
              "1号梯外呼上面无目标5" := "中间变量2"."5号梯外呼上面无目标5",
              "1号梯外呼上面无目标6" := "中间变量2"."5号梯外呼上面无目标6",
              "1号梯外呼上面无目标7" := "中间变量2"."5号梯外呼上面无目标7",
              "1号梯外呼上面无目标8" := "中间变量2"."5号梯外呼上面无目标8",
              "1号梯外呼上面无目标9" := "中间变量2"."5号梯外呼上面无目标9",
              "1号梯外呼下面无目标2" := "中间变量2"."5号梯外呼下面无目标2",
              "1号梯外呼下面无目标3" := "中间变量2"."5号梯外呼下面无目标3",
              "1号梯外呼下面无目标4" := "中间变量2"."5号梯外呼下面无目标4",
              "1号梯外呼下面无目标5" := "中间变量2"."5号梯外呼下面无目标5",
              "1号梯外呼下面无目标6" := "中间变量2"."5号梯外呼下面无目标6",
              "1号梯外呼下面无目标7" := "中间变量2"."5号梯外呼下面无目标7",
              "1号梯外呼下面无目标8" := "中间变量2"."5号梯外呼下面无目标8",
              "1号梯外呼下面无目标9" := "中间变量2"."5号梯外呼下面无目标9",
              初始化高速运行 := "中间变量1"."5号梯高速初始化",
              "1号梯高速接触器" => "输出"."5号梯高速接触器",
              "1号梯低速接触器" => "输出"."5号梯低速接触器",
              将要停梯 => "中间变量1"."5号梯将要停梯");
END_REGION

REGION Network 6: 6号梯
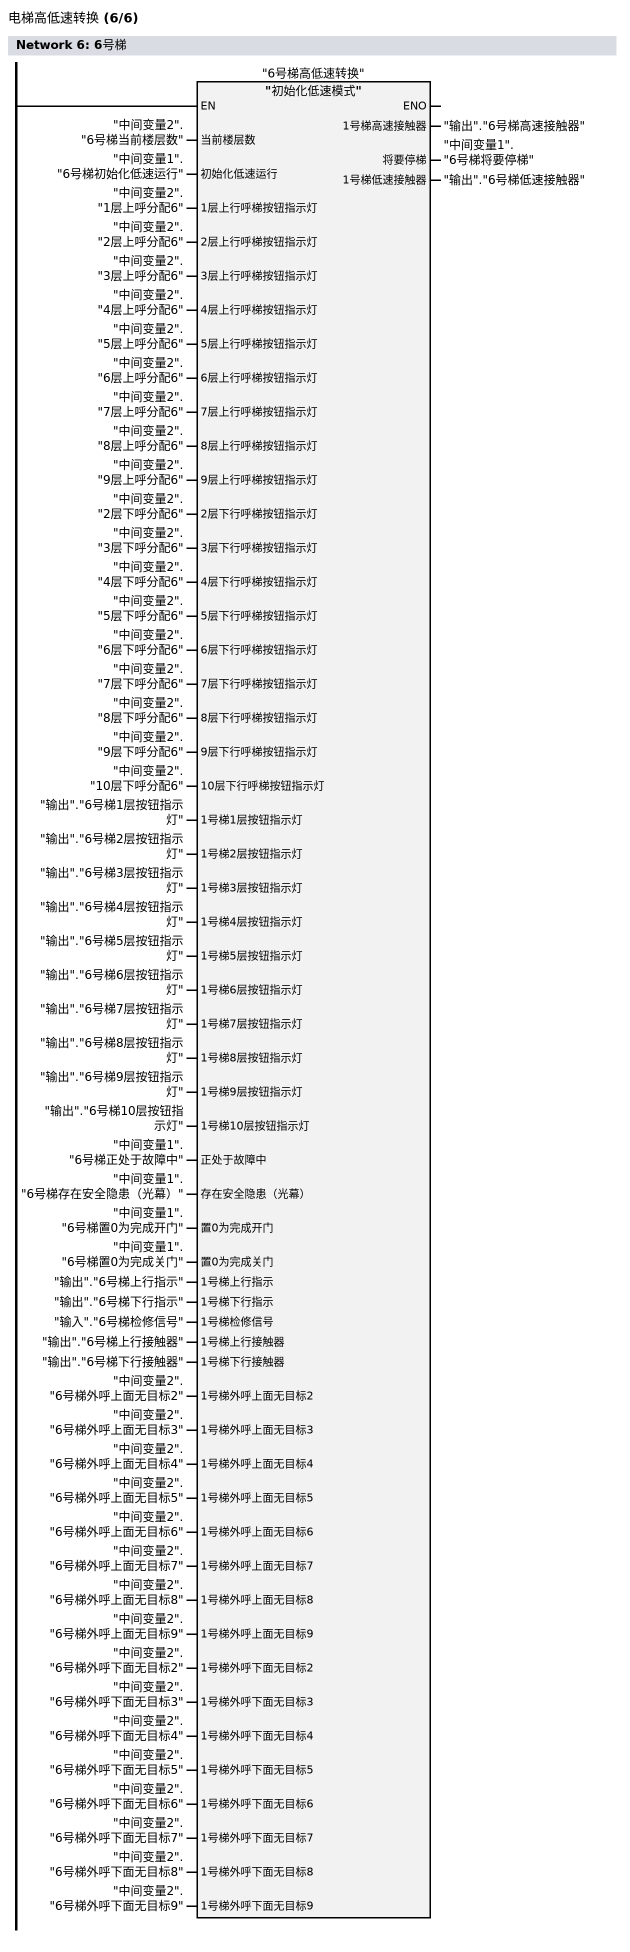
   RUNG wire#powerrail
      "6号梯高低速转换"(当前楼层数 := "中间变量2"."6号梯当前楼层数", 初始化低速运行 := "中间变量1"."6号梯初始化低速运行", "1层上行呼梯按钮指示灯" := "中间变量2"."1层上呼分配6", "2层上行呼梯按钮指示灯" := "中间变量2"."2层上呼分配6", "3层上行呼梯按钮指示灯" := "中间变量2"."3层上呼分配6", "4层上行呼梯按钮指示灯" := "中间变量2"."4层上呼分配6", "5层上行呼梯按钮指示灯" := "中间变量2"."5层上呼分配6", "6层上行呼梯按钮指示灯" := "中间变量2"."6层上呼分配6", "7层上行呼梯按钮指示灯" := "中间变量2"."7层上呼分配6", "8层上行呼梯按钮指示灯" := "中间变量2"."8层上呼分配6", "9层上行呼梯按钮指示灯" := "中间变量2"."9层上呼分配6", "2层下行呼梯按钮指示灯" := "中间变量2"."2层下呼分配6", "3层下行呼梯按钮指示灯" := "中间变量2"."3层下呼分配6", "4层下行呼梯按钮指示灯" := "中间变量2"."4层下呼分配6", "5层下行呼梯按钮指示灯" := "中间变量2"."5层下呼分配6", "6层下行呼梯按钮指示灯" := "中间变量2"."6层下呼分配6", "7层下行呼梯按钮指示灯" := "中间变量2"."7层下呼分配6", "8层下行呼梯按钮指示灯" := "中间变量2"."8层下呼分配6", "9层下行呼梯按钮指示灯" := "中间变量2"."9层下呼分配6", "10层下行呼梯按钮指示灯" := "中间变量2"."10层下呼分配6", "1号梯1层按钮指示灯" := "输出"."6号梯1层按钮指示灯", "1号梯2层按钮指示灯" := "输出"."6号梯2层按钮指示灯", "1号梯3层按钮指示灯" := "输出"."6号梯3层按钮指示灯", "1号梯4层按钮指示灯" := "输出"."6号梯4层按钮指示灯", "1号梯5层按钮指示灯" := "输出"."6号梯5层按钮指示灯", "1号梯6层按钮指示灯" := "输出"."6号梯6层按钮指示灯", "1号梯7层按钮指示灯" := "输出"."6号梯7层按钮指示灯", "1号梯8层按钮指示灯" := "输出"."6号梯8层按钮指示灯", "1号梯9层按钮指示灯" := "输出"."6号梯9层按钮指示灯", "1号梯10层按钮指示灯" := "输出"."6号梯10层按钮指示灯", 正处于故障中 := "中间变量1"."6号梯正处于故障中", "存在安全隐患（光幕）" := "中间变量1"."6号梯存在安全隐患（光幕）", 置0为完成开门 := "中间变量1"."6号梯置0为完成开门", 置0为完成关门 := "中间变量1"."6号梯置0为完成关门", "1号梯上行指示" := "输出"."6号梯上行指示", "1号梯下行指示" := "输出"."6号梯下行指示", "1号梯检修信号" := "输入"."6号梯检修信号", "1号梯上行接触器" := "输出"."6号梯上行接触器", "1号梯下行接触器" := "输出"."6号梯下行接触器", "1号梯外呼上面无目标2" := "中间变量2"."6号梯外呼上面无目标2", "1号梯外呼上面无目标3" := "中间变量2"."6号梯外呼上面无目标3", "1号梯外呼上面无目标4" := "中间变量2"."6号梯外呼上面无目标4", "1号梯外呼上面无目标5" := "中间变量2"."6号梯外呼上面无目标5", "1号梯外呼上面无目标6" := "中间变量2"."6号梯外呼上面无目标6", "1号梯外呼上面无目标7" := "中间变量2"."6号梯外呼上面无目标7", "1号梯外呼上面无目标8" := "中间变量2"."6号梯外呼上面无目标8", "1号梯外呼上面无目标9" := "中间变量2"."6号梯外呼上面无目标9", "1号梯外呼下面无目标2" := "中间变量2"."6号梯外呼下面无目标2", "1号梯外呼下面无目标3" := "中间变量2"."6号梯外呼下面无目标3", "1号梯外呼下面无目标4" := "中间变量2"."6号梯外呼下面无目标4", "1号梯外呼下面无目标5" := "中间变量2"."6号梯外呼下面无目标5", "1号梯外呼下面无目标6" := "中间变量2"."6号梯外呼下面无目标6", "1号梯外呼下面无目标7" := "中间变量2"."6号梯外呼下面无目标7", "1号梯外呼下面无目标8" := "中间变量2"."6号梯外呼下面无目标8", "1号梯外呼下面无目标9" := "中间变量2"."6号梯外呼下面无目标9", "1号梯高速接触器" => "输出"."6号梯高速接触器", 将要停梯 => "中间变量1"."6号梯将要停梯", "1号梯低速接触器" => "输出"."6号梯低速接触器")
   END_RUNG
   // the same network as SCL:
   "6号梯高低速转换"(当前楼层数 := "中间变量2"."6号梯当前楼层数",   // "初始化低速模式"
              初始化低速运行 := "中间变量1"."6号梯初始化低速运行",
              "1层上行呼梯按钮指示灯" := "中间变量2"."1层上呼分配6",
              "2层上行呼梯按钮指示灯" := "中间变量2"."2层上呼分配6",
              "3层上行呼梯按钮指示灯" := "中间变量2"."3层上呼分配6",
              "4层上行呼梯按钮指示灯" := "中间变量2"."4层上呼分配6",
              "5层上行呼梯按钮指示灯" := "中间变量2"."5层上呼分配6",
              "6层上行呼梯按钮指示灯" := "中间变量2"."6层上呼分配6",
              "7层上行呼梯按钮指示灯" := "中间变量2"."7层上呼分配6",
              "8层上行呼梯按钮指示灯" := "中间变量2"."8层上呼分配6",
              "9层上行呼梯按钮指示灯" := "中间变量2"."9层上呼分配6",
              "2层下行呼梯按钮指示灯" := "中间变量2"."2层下呼分配6",
              "3层下行呼梯按钮指示灯" := "中间变量2"."3层下呼分配6",
              "4层下行呼梯按钮指示灯" := "中间变量2"."4层下呼分配6",
              "5层下行呼梯按钮指示灯" := "中间变量2"."5层下呼分配6",
              "6层下行呼梯按钮指示灯" := "中间变量2"."6层下呼分配6",
              "7层下行呼梯按钮指示灯" := "中间变量2"."7层下呼分配6",
              "8层下行呼梯按钮指示灯" := "中间变量2"."8层下呼分配6",
              "9层下行呼梯按钮指示灯" := "中间变量2"."9层下呼分配6",
              "10层下行呼梯按钮指示灯" := "中间变量2"."10层下呼分配6",
              "1号梯1层按钮指示灯" := "输出"."6号梯1层按钮指示灯",
              "1号梯2层按钮指示灯" := "输出"."6号梯2层按钮指示灯",
              "1号梯3层按钮指示灯" := "输出"."6号梯3层按钮指示灯",
              "1号梯4层按钮指示灯" := "输出"."6号梯4层按钮指示灯",
              "1号梯5层按钮指示灯" := "输出"."6号梯5层按钮指示灯",
              "1号梯6层按钮指示灯" := "输出"."6号梯6层按钮指示灯",
              "1号梯7层按钮指示灯" := "输出"."6号梯7层按钮指示灯",
              "1号梯8层按钮指示灯" := "输出"."6号梯8层按钮指示灯",
              "1号梯9层按钮指示灯" := "输出"."6号梯9层按钮指示灯",
              "1号梯10层按钮指示灯" := "输出"."6号梯10层按钮指示灯",
              正处于故障中 := "中间变量1"."6号梯正处于故障中",
              "存在安全隐患（光幕）" := "中间变量1"."6号梯存在安全隐患（光幕）",
              置0为完成开门 := "中间变量1"."6号梯置0为完成开门",
              置0为完成关门 := "中间变量1"."6号梯置0为完成关门",
              "1号梯上行指示" := "输出"."6号梯上行指示",
              "1号梯下行指示" := "输出"."6号梯下行指示",
              "1号梯检修信号" := "输入"."6号梯检修信号",
              "1号梯上行接触器" := "输出"."6号梯上行接触器",
              "1号梯下行接触器" := "输出"."6号梯下行接触器",
              "1号梯外呼上面无目标2" := "中间变量2"."6号梯外呼上面无目标2",
              "1号梯外呼上面无目标3" := "中间变量2"."6号梯外呼上面无目标3",
              "1号梯外呼上面无目标4" := "中间变量2"."6号梯外呼上面无目标4",
              "1号梯外呼上面无目标5" := "中间变量2"."6号梯外呼上面无目标5",
              "1号梯外呼上面无目标6" := "中间变量2"."6号梯外呼上面无目标6",
              "1号梯外呼上面无目标7" := "中间变量2"."6号梯外呼上面无目标7",
              "1号梯外呼上面无目标8" := "中间变量2"."6号梯外呼上面无目标8",
              "1号梯外呼上面无目标9" := "中间变量2"."6号梯外呼上面无目标9",
              "1号梯外呼下面无目标2" := "中间变量2"."6号梯外呼下面无目标2",
              "1号梯外呼下面无目标3" := "中间变量2"."6号梯外呼下面无目标3",
              "1号梯外呼下面无目标4" := "中间变量2"."6号梯外呼下面无目标4",
              "1号梯外呼下面无目标5" := "中间变量2"."6号梯外呼下面无目标5",
              "1号梯外呼下面无目标6" := "中间变量2"."6号梯外呼下面无目标6",
              "1号梯外呼下面无目标7" := "中间变量2"."6号梯外呼下面无目标7",
              "1号梯外呼下面无目标8" := "中间变量2"."6号梯外呼下面无目标8",
              "1号梯外呼下面无目标9" := "中间变量2"."6号梯外呼下面无目标9",
              "1号梯高速接触器" => "输出"."6号梯高速接触器",
              将要停梯 => "中间变量1"."6号梯将要停梯",
              "1号梯低速接触器" => "输出"."6号梯低速接触器");
END_REGION
END_FUNCTION

FUNCTION "电梯运行与制动" : Void   // FC4, LAD
{ S7_Optimized_Access := 'TRUE' }
VERSION : 0.1
BEGIN

REGION Network 1: 1号梯
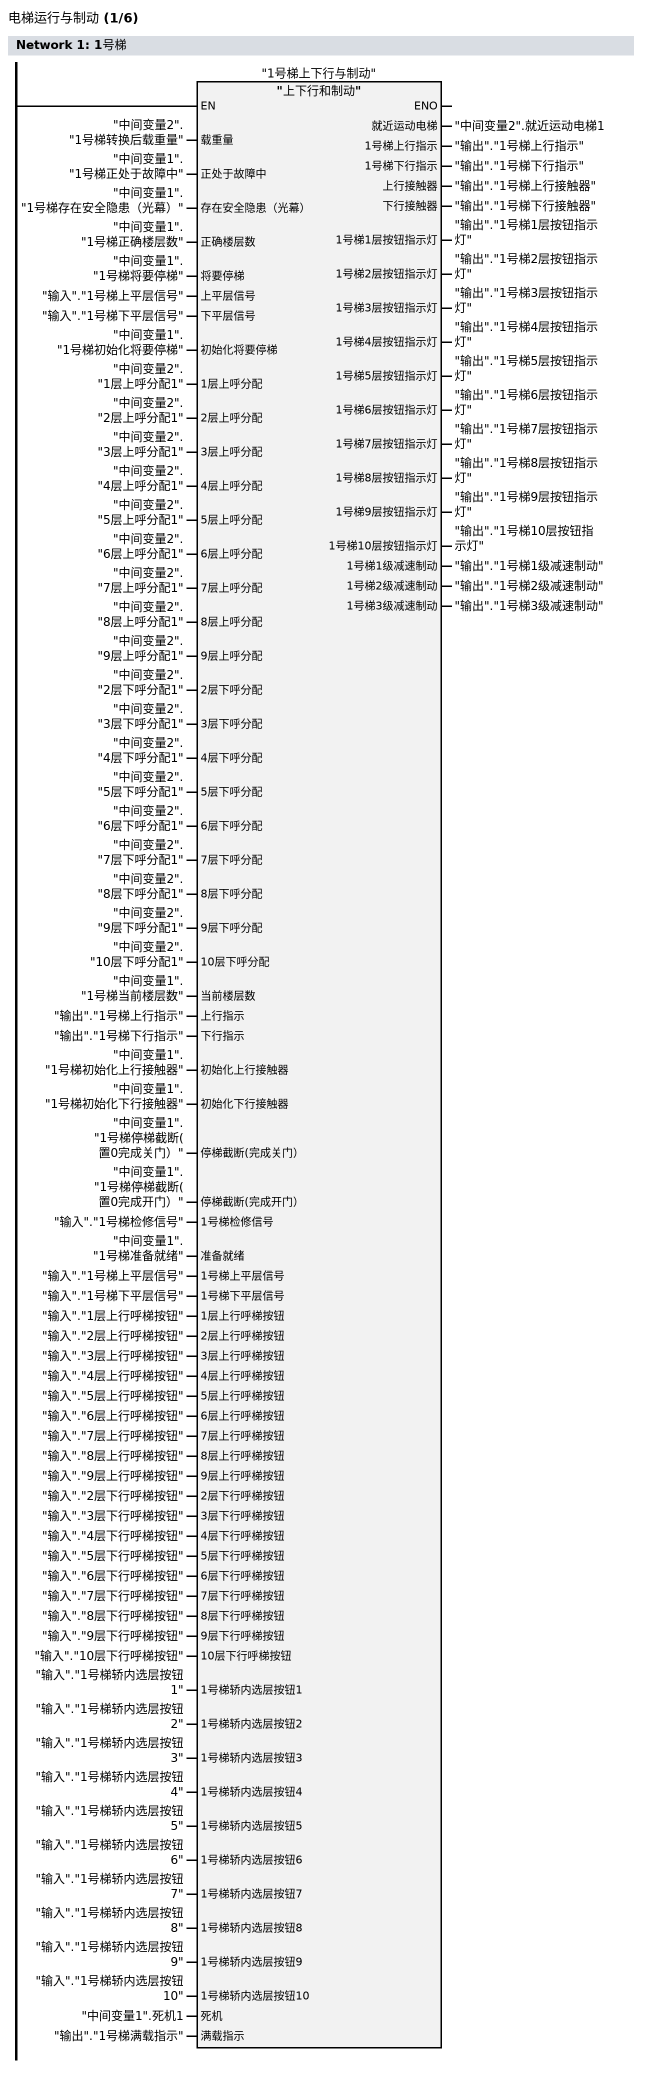
   RUNG wire#powerrail
      "1号梯上下行与制动"(载重量 := "中间变量2"."1号梯转换后载重量", 正处于故障中 := "中间变量1"."1号梯正处于故障中", "存在安全隐患（光幕）" := "中间变量1"."1号梯存在安全隐患（光幕）", 正确楼层数 := "中间变量1"."1号梯正确楼层数", 将要停梯 := "中间变量1"."1号梯将要停梯", 上平层信号 := "输入"."1号梯上平层信号", 下平层信号 := "输入"."1号梯下平层信号", 初始化将要停梯 := "中间变量1"."1号梯初始化将要停梯", "1层上呼分配" := "中间变量2"."1层上呼分配1", "2层上呼分配" := "中间变量2"."2层上呼分配1", "3层上呼分配" := "中间变量2"."3层上呼分配1", "4层上呼分配" := "中间变量2"."4层上呼分配1", "5层上呼分配" := "中间变量2"."5层上呼分配1", "6层上呼分配" := "中间变量2"."6层上呼分配1", "7层上呼分配" := "中间变量2"."7层上呼分配1", "8层上呼分配" := "中间变量2"."8层上呼分配1", "9层上呼分配" := "中间变量2"."9层上呼分配1", "2层下呼分配" := "中间变量2"."2层下呼分配1", "3层下呼分配" := "中间变量2"."3层下呼分配1", "4层下呼分配" := "中间变量2"."4层下呼分配1", "5层下呼分配" := "中间变量2"."5层下呼分配1", "6层下呼分配" := "中间变量2"."6层下呼分配1", "7层下呼分配" := "中间变量2"."7层下呼分配1", "8层下呼分配" := "中间变量2"."8层下呼分配1", "9层下呼分配" := "中间变量2"."9层下呼分配1", "10层下呼分配" := "中间变量2"."10层下呼分配1", 当前楼层数 := "中间变量1"."1号梯当前楼层数", 上行指示 := "输出"."1号梯上行指示", 下行指示 := "输出"."1号梯下行指示", 初始化上行接触器 := "中间变量1"."1号梯初始化上行接触器", 初始化下行接触器 := "中间变量1"."1号梯初始化下行接触器", "停梯截断(完成关门）" := "中间变量1"."1号梯停梯截断(置0完成关门）", "停梯截断(完成开门）" := "中间变量1"."1号梯停梯截断(置0完成开门）", "1号梯检修信号" := "输入"."1号梯检修信号", 准备就绪 := "中间变量1"."1号梯准备就绪", "1号梯上平层信号" := "输入"."1号梯上平层信号", "1号梯下平层信号" := "输入"."1号梯下平层信号", "1层上行呼梯按钮" := "输入"."1层上行呼梯按钮", "2层上行呼梯按钮" := "输入"."2层上行呼梯按钮", "3层上行呼梯按钮" := "输入"."3层上行呼梯按钮", "4层上行呼梯按钮" := "输入"."4层上行呼梯按钮", "5层上行呼梯按钮" := "输入"."5层上行呼梯按钮", "6层上行呼梯按钮" := "输入"."6层上行呼梯按钮", "7层上行呼梯按钮" := "输入"."7层上行呼梯按钮", "8层上行呼梯按钮" := "输入"."8层上行呼梯按钮", "9层上行呼梯按钮" := "输入"."9层上行呼梯按钮", "2层下行呼梯按钮" := "输入"."2层下行呼梯按钮", "3层下行呼梯按钮" := "输入"."3层下行呼梯按钮", "4层下行呼梯按钮" := "输入"."4层下行呼梯按钮", "5层下行呼梯按钮" := "输入"."5层下行呼梯按钮", "6层下行呼梯按钮" := "输入"."6层下行呼梯按钮", "7层下行呼梯按钮" := "输入"."7层下行呼梯按钮", "8层下行呼梯按钮" := "输入"."8层下行呼梯按钮", "9层下行呼梯按钮" := "输入"."9层下行呼梯按钮", "10层下行呼梯按钮" := "输入"."10层下行呼梯按钮", "1号梯轿内选层按钮1" := "输入"."1号梯轿内选层按钮1", "1号梯轿内选层按钮2" := "输入"."1号梯轿内选层按钮2", "1号梯轿内选层按钮3" := "输入"."1号梯轿内选层按钮3", "1号梯轿内选层按钮4" := "输入"."1号梯轿内选层按钮4", "1号梯轿内选层按钮5" := "输入"."1号梯轿内选层按钮5", "1号梯轿内选层按钮6" := "输入"."1号梯轿内选层按钮6", "1号梯轿内选层按钮7" := "输入"."1号梯轿内选层按钮7", "1号梯轿内选层按钮8" := "输入"."1号梯轿内选层按钮8", "1号梯轿内选层按钮9" := "输入"."1号梯轿内选层按钮9", "1号梯轿内选层按钮10" := "输入"."1号梯轿内选层按钮10", 死机 := "中间变量1".死机1, 满载指示 := "输出"."1号梯满载指示", 就近运动电梯 => "中间变量2".就近运动电梯1, "1号梯上行指示" => "输出"."1号梯上行指示", "1号梯下行指示" => "输出"."1号梯下行指示", 上行接触器 => "输出"."1号梯上行接触器", 下行接触器 => "输出"."1号梯下行接触器", "1号梯1层按钮指示灯" => "输出"."1号梯1层按钮指示灯", "1号梯2层按钮指示灯" => "输出"."1号梯2层按钮指示灯", "1号梯3层按钮指示灯" => "输出"."1号梯3层按钮指示灯", "1号梯4层按钮指示灯" => "输出"."1号梯4层按钮指示灯", "1号梯5层按钮指示灯" => "输出"."1号梯5层按钮指示灯", "1号梯6层按钮指示灯" => "输出"."1号梯6层按钮指示灯", "1号梯7层按钮指示灯" => "输出"."1号梯7层按钮指示灯", "1号梯8层按钮指示灯" => "输出"."1号梯8层按钮指示灯", "1号梯9层按钮指示灯" => "输出"."1号梯9层按钮指示灯", "1号梯10层按钮指示灯" => "输出"."1号梯10层按钮指示灯", "1号梯1级减速制动" => "输出"."1号梯1级减速制动", "1号梯2级减速制动" => "输出"."1号梯2级减速制动", "1号梯3级减速制动" => "输出"."1号梯3级减速制动")
   END_RUNG
   // the same network as SCL:
   "1号梯上下行与制动"(载重量 := "中间变量2"."1号梯转换后载重量",   // "上下行和制动"
               正处于故障中 := "中间变量1"."1号梯正处于故障中",
               "存在安全隐患（光幕）" := "中间变量1"."1号梯存在安全隐患（光幕）",
               正确楼层数 := "中间变量1"."1号梯正确楼层数",
               将要停梯 := "中间变量1"."1号梯将要停梯",
               上平层信号 := "输入"."1号梯上平层信号",
               下平层信号 := "输入"."1号梯下平层信号",
               初始化将要停梯 := "中间变量1"."1号梯初始化将要停梯",
               "1层上呼分配" := "中间变量2"."1层上呼分配1",
               "2层上呼分配" := "中间变量2"."2层上呼分配1",
               "3层上呼分配" := "中间变量2"."3层上呼分配1",
               "4层上呼分配" := "中间变量2"."4层上呼分配1",
               "5层上呼分配" := "中间变量2"."5层上呼分配1",
               "6层上呼分配" := "中间变量2"."6层上呼分配1",
               "7层上呼分配" := "中间变量2"."7层上呼分配1",
               "8层上呼分配" := "中间变量2"."8层上呼分配1",
               "9层上呼分配" := "中间变量2"."9层上呼分配1",
               "2层下呼分配" := "中间变量2"."2层下呼分配1",
               "3层下呼分配" := "中间变量2"."3层下呼分配1",
               "4层下呼分配" := "中间变量2"."4层下呼分配1",
               "5层下呼分配" := "中间变量2"."5层下呼分配1",
               "6层下呼分配" := "中间变量2"."6层下呼分配1",
               "7层下呼分配" := "中间变量2"."7层下呼分配1",
               "8层下呼分配" := "中间变量2"."8层下呼分配1",
               "9层下呼分配" := "中间变量2"."9层下呼分配1",
               "10层下呼分配" := "中间变量2"."10层下呼分配1",
               当前楼层数 := "中间变量1"."1号梯当前楼层数",
               上行指示 := "输出"."1号梯上行指示",
               下行指示 := "输出"."1号梯下行指示",
               初始化上行接触器 := "中间变量1"."1号梯初始化上行接触器",
               初始化下行接触器 := "中间变量1"."1号梯初始化下行接触器",
               "停梯截断(完成关门）" := "中间变量1"."1号梯停梯截断(置0完成关门）",
               "停梯截断(完成开门）" := "中间变量1"."1号梯停梯截断(置0完成开门）",
               "1号梯检修信号" := "输入"."1号梯检修信号",
               准备就绪 := "中间变量1"."1号梯准备就绪",
               "1号梯上平层信号" := "输入"."1号梯上平层信号",
               "1号梯下平层信号" := "输入"."1号梯下平层信号",
               "1层上行呼梯按钮" := "输入"."1层上行呼梯按钮",
               "2层上行呼梯按钮" := "输入"."2层上行呼梯按钮",
               "3层上行呼梯按钮" := "输入"."3层上行呼梯按钮",
               "4层上行呼梯按钮" := "输入"."4层上行呼梯按钮",
               "5层上行呼梯按钮" := "输入"."5层上行呼梯按钮",
               "6层上行呼梯按钮" := "输入"."6层上行呼梯按钮",
               "7层上行呼梯按钮" := "输入"."7层上行呼梯按钮",
               "8层上行呼梯按钮" := "输入"."8层上行呼梯按钮",
               "9层上行呼梯按钮" := "输入"."9层上行呼梯按钮",
               "2层下行呼梯按钮" := "输入"."2层下行呼梯按钮",
               "3层下行呼梯按钮" := "输入"."3层下行呼梯按钮",
               "4层下行呼梯按钮" := "输入"."4层下行呼梯按钮",
               "5层下行呼梯按钮" := "输入"."5层下行呼梯按钮",
               "6层下行呼梯按钮" := "输入"."6层下行呼梯按钮",
               "7层下行呼梯按钮" := "输入"."7层下行呼梯按钮",
               "8层下行呼梯按钮" := "输入"."8层下行呼梯按钮",
               "9层下行呼梯按钮" := "输入"."9层下行呼梯按钮",
               "10层下行呼梯按钮" := "输入"."10层下行呼梯按钮",
               "1号梯轿内选层按钮1" := "输入"."1号梯轿内选层按钮1",
               "1号梯轿内选层按钮2" := "输入"."1号梯轿内选层按钮2",
               "1号梯轿内选层按钮3" := "输入"."1号梯轿内选层按钮3",
               "1号梯轿内选层按钮4" := "输入"."1号梯轿内选层按钮4",
               "1号梯轿内选层按钮5" := "输入"."1号梯轿内选层按钮5",
               "1号梯轿内选层按钮6" := "输入"."1号梯轿内选层按钮6",
               "1号梯轿内选层按钮7" := "输入"."1号梯轿内选层按钮7",
               "1号梯轿内选层按钮8" := "输入"."1号梯轿内选层按钮8",
               "1号梯轿内选层按钮9" := "输入"."1号梯轿内选层按钮9",
               "1号梯轿内选层按钮10" := "输入"."1号梯轿内选层按钮10",
               死机 := "中间变量1".死机1,
               满载指示 := "输出"."1号梯满载指示",
               就近运动电梯 => "中间变量2".就近运动电梯1,
               "1号梯上行指示" => "输出"."1号梯上行指示",
               "1号梯下行指示" => "输出"."1号梯下行指示",
               上行接触器 => "输出"."1号梯上行接触器",
               下行接触器 => "输出"."1号梯下行接触器",
               "1号梯1层按钮指示灯" => "输出"."1号梯1层按钮指示灯",
               "1号梯2层按钮指示灯" => "输出"."1号梯2层按钮指示灯",
               "1号梯3层按钮指示灯" => "输出"."1号梯3层按钮指示灯",
               "1号梯4层按钮指示灯" => "输出"."1号梯4层按钮指示灯",
               "1号梯5层按钮指示灯" => "输出"."1号梯5层按钮指示灯",
               "1号梯6层按钮指示灯" => "输出"."1号梯6层按钮指示灯",
               "1号梯7层按钮指示灯" => "输出"."1号梯7层按钮指示灯",
               "1号梯8层按钮指示灯" => "输出"."1号梯8层按钮指示灯",
               "1号梯9层按钮指示灯" => "输出"."1号梯9层按钮指示灯",
               "1号梯10层按钮指示灯" => "输出"."1号梯10层按钮指示灯",
               "1号梯1级减速制动" => "输出"."1号梯1级减速制动",
               "1号梯2级减速制动" => "输出"."1号梯2级减速制动",
               "1号梯3级减速制动" => "输出"."1号梯3级减速制动");
END_REGION

REGION Network 2: 2号梯
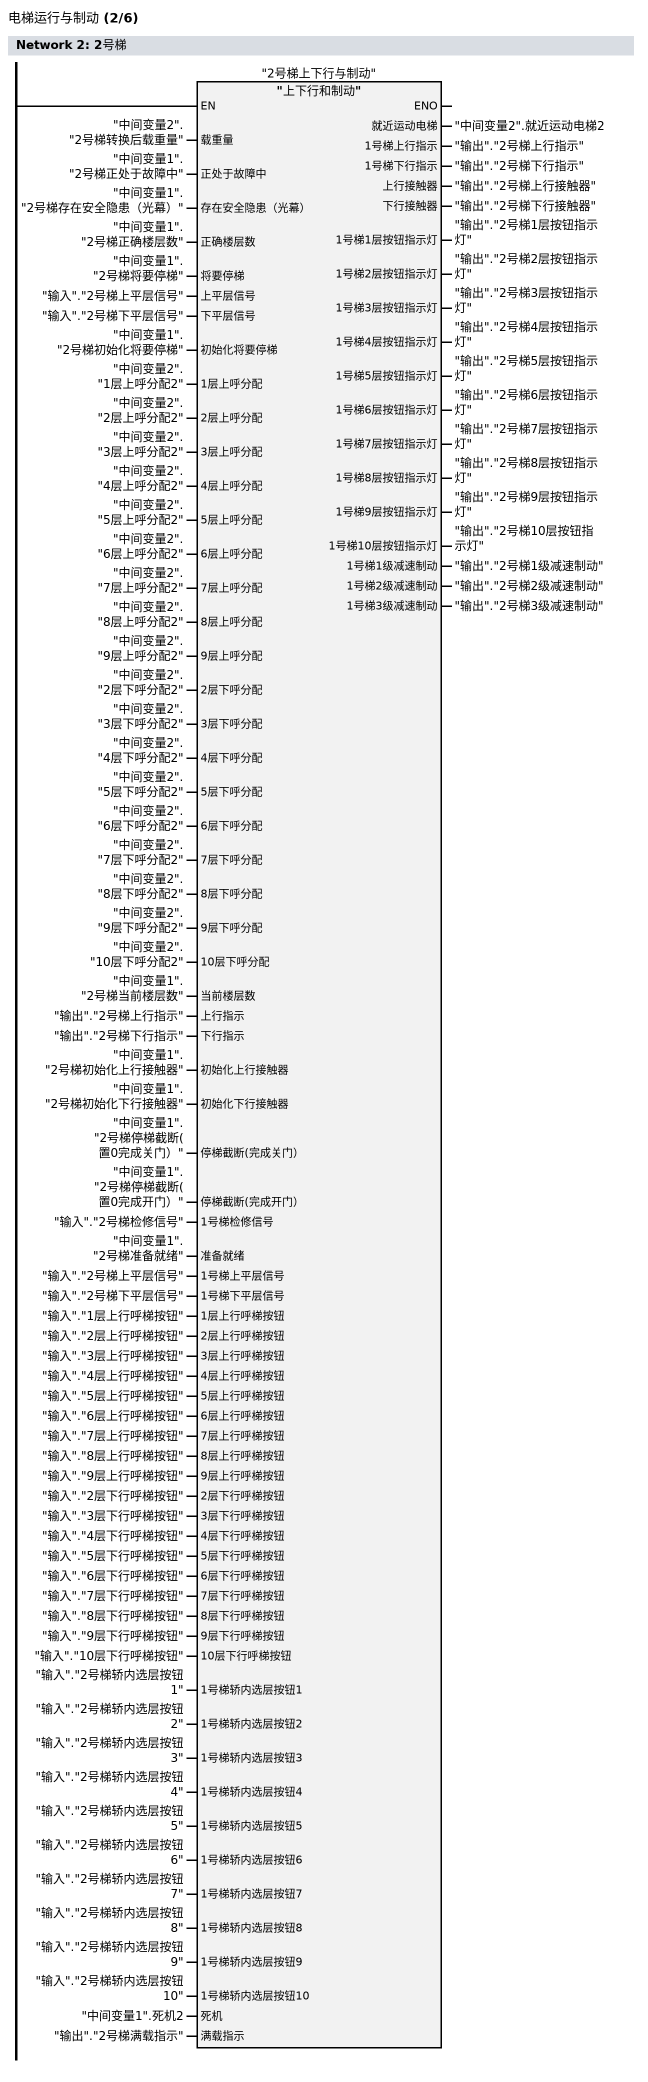
   RUNG wire#powerrail
      "2号梯上下行与制动"(载重量 := "中间变量2"."2号梯转换后载重量", 正处于故障中 := "中间变量1"."2号梯正处于故障中", "存在安全隐患（光幕）" := "中间变量1"."2号梯存在安全隐患（光幕）", 正确楼层数 := "中间变量1"."2号梯正确楼层数", 将要停梯 := "中间变量1"."2号梯将要停梯", 上平层信号 := "输入"."2号梯上平层信号", 下平层信号 := "输入"."2号梯下平层信号", 初始化将要停梯 := "中间变量1"."2号梯初始化将要停梯", "1层上呼分配" := "中间变量2"."1层上呼分配2", "2层上呼分配" := "中间变量2"."2层上呼分配2", "3层上呼分配" := "中间变量2"."3层上呼分配2", "4层上呼分配" := "中间变量2"."4层上呼分配2", "5层上呼分配" := "中间变量2"."5层上呼分配2", "6层上呼分配" := "中间变量2"."6层上呼分配2", "7层上呼分配" := "中间变量2"."7层上呼分配2", "8层上呼分配" := "中间变量2"."8层上呼分配2", "9层上呼分配" := "中间变量2"."9层上呼分配2", "2层下呼分配" := "中间变量2"."2层下呼分配2", "3层下呼分配" := "中间变量2"."3层下呼分配2", "4层下呼分配" := "中间变量2"."4层下呼分配2", "5层下呼分配" := "中间变量2"."5层下呼分配2", "6层下呼分配" := "中间变量2"."6层下呼分配2", "7层下呼分配" := "中间变量2"."7层下呼分配2", "8层下呼分配" := "中间变量2"."8层下呼分配2", "9层下呼分配" := "中间变量2"."9层下呼分配2", "10层下呼分配" := "中间变量2"."10层下呼分配2", 当前楼层数 := "中间变量1"."2号梯当前楼层数", 上行指示 := "输出"."2号梯上行指示", 下行指示 := "输出"."2号梯下行指示", 初始化上行接触器 := "中间变量1"."2号梯初始化上行接触器", 初始化下行接触器 := "中间变量1"."2号梯初始化下行接触器", "停梯截断(完成关门）" := "中间变量1"."2号梯停梯截断(置0完成关门）", "停梯截断(完成开门）" := "中间变量1"."2号梯停梯截断(置0完成开门）", "1号梯检修信号" := "输入"."2号梯检修信号", 准备就绪 := "中间变量1"."2号梯准备就绪", "1号梯上平层信号" := "输入"."2号梯上平层信号", "1号梯下平层信号" := "输入"."2号梯下平层信号", "1层上行呼梯按钮" := "输入"."1层上行呼梯按钮", "2层上行呼梯按钮" := "输入"."2层上行呼梯按钮", "3层上行呼梯按钮" := "输入"."3层上行呼梯按钮", "4层上行呼梯按钮" := "输入"."4层上行呼梯按钮", "5层上行呼梯按钮" := "输入"."5层上行呼梯按钮", "6层上行呼梯按钮" := "输入"."6层上行呼梯按钮", "7层上行呼梯按钮" := "输入"."7层上行呼梯按钮", "8层上行呼梯按钮" := "输入"."8层上行呼梯按钮", "9层上行呼梯按钮" := "输入"."9层上行呼梯按钮", "2层下行呼梯按钮" := "输入"."2层下行呼梯按钮", "3层下行呼梯按钮" := "输入"."3层下行呼梯按钮", "4层下行呼梯按钮" := "输入"."4层下行呼梯按钮", "5层下行呼梯按钮" := "输入"."5层下行呼梯按钮", "6层下行呼梯按钮" := "输入"."6层下行呼梯按钮", "7层下行呼梯按钮" := "输入"."7层下行呼梯按钮", "8层下行呼梯按钮" := "输入"."8层下行呼梯按钮", "9层下行呼梯按钮" := "输入"."9层下行呼梯按钮", "10层下行呼梯按钮" := "输入"."10层下行呼梯按钮", "1号梯轿内选层按钮1" := "输入"."2号梯轿内选层按钮1", "1号梯轿内选层按钮2" := "输入"."2号梯轿内选层按钮2", "1号梯轿内选层按钮3" := "输入"."2号梯轿内选层按钮3", "1号梯轿内选层按钮4" := "输入"."2号梯轿内选层按钮4", "1号梯轿内选层按钮5" := "输入"."2号梯轿内选层按钮5", "1号梯轿内选层按钮6" := "输入"."2号梯轿内选层按钮6", "1号梯轿内选层按钮7" := "输入"."2号梯轿内选层按钮7", "1号梯轿内选层按钮8" := "输入"."2号梯轿内选层按钮8", "1号梯轿内选层按钮9" := "输入"."2号梯轿内选层按钮9", "1号梯轿内选层按钮10" := "输入"."2号梯轿内选层按钮10", 死机 := "中间变量1".死机2, 满载指示 := "输出"."2号梯满载指示", 就近运动电梯 => "中间变量2".就近运动电梯2, "1号梯上行指示" => "输出"."2号梯上行指示", "1号梯下行指示" => "输出"."2号梯下行指示", 上行接触器 => "输出"."2号梯上行接触器", 下行接触器 => "输出"."2号梯下行接触器", "1号梯1层按钮指示灯" => "输出"."2号梯1层按钮指示灯", "1号梯2层按钮指示灯" => "输出"."2号梯2层按钮指示灯", "1号梯3层按钮指示灯" => "输出"."2号梯3层按钮指示灯", "1号梯4层按钮指示灯" => "输出"."2号梯4层按钮指示灯", "1号梯5层按钮指示灯" => "输出"."2号梯5层按钮指示灯", "1号梯6层按钮指示灯" => "输出"."2号梯6层按钮指示灯", "1号梯7层按钮指示灯" => "输出"."2号梯7层按钮指示灯", "1号梯8层按钮指示灯" => "输出"."2号梯8层按钮指示灯", "1号梯9层按钮指示灯" => "输出"."2号梯9层按钮指示灯", "1号梯10层按钮指示灯" => "输出"."2号梯10层按钮指示灯", "1号梯1级减速制动" => "输出"."2号梯1级减速制动", "1号梯2级减速制动" => "输出"."2号梯2级减速制动", "1号梯3级减速制动" => "输出"."2号梯3级减速制动")
   END_RUNG
   // the same network as SCL:
   "2号梯上下行与制动"(载重量 := "中间变量2"."2号梯转换后载重量",   // "上下行和制动"
               正处于故障中 := "中间变量1"."2号梯正处于故障中",
               "存在安全隐患（光幕）" := "中间变量1"."2号梯存在安全隐患（光幕）",
               正确楼层数 := "中间变量1"."2号梯正确楼层数",
               将要停梯 := "中间变量1"."2号梯将要停梯",
               上平层信号 := "输入"."2号梯上平层信号",
               下平层信号 := "输入"."2号梯下平层信号",
               初始化将要停梯 := "中间变量1"."2号梯初始化将要停梯",
               "1层上呼分配" := "中间变量2"."1层上呼分配2",
               "2层上呼分配" := "中间变量2"."2层上呼分配2",
               "3层上呼分配" := "中间变量2"."3层上呼分配2",
               "4层上呼分配" := "中间变量2"."4层上呼分配2",
               "5层上呼分配" := "中间变量2"."5层上呼分配2",
               "6层上呼分配" := "中间变量2"."6层上呼分配2",
               "7层上呼分配" := "中间变量2"."7层上呼分配2",
               "8层上呼分配" := "中间变量2"."8层上呼分配2",
               "9层上呼分配" := "中间变量2"."9层上呼分配2",
               "2层下呼分配" := "中间变量2"."2层下呼分配2",
               "3层下呼分配" := "中间变量2"."3层下呼分配2",
               "4层下呼分配" := "中间变量2"."4层下呼分配2",
               "5层下呼分配" := "中间变量2"."5层下呼分配2",
               "6层下呼分配" := "中间变量2"."6层下呼分配2",
               "7层下呼分配" := "中间变量2"."7层下呼分配2",
               "8层下呼分配" := "中间变量2"."8层下呼分配2",
               "9层下呼分配" := "中间变量2"."9层下呼分配2",
               "10层下呼分配" := "中间变量2"."10层下呼分配2",
               当前楼层数 := "中间变量1"."2号梯当前楼层数",
               上行指示 := "输出"."2号梯上行指示",
               下行指示 := "输出"."2号梯下行指示",
               初始化上行接触器 := "中间变量1"."2号梯初始化上行接触器",
               初始化下行接触器 := "中间变量1"."2号梯初始化下行接触器",
               "停梯截断(完成关门）" := "中间变量1"."2号梯停梯截断(置0完成关门）",
               "停梯截断(完成开门）" := "中间变量1"."2号梯停梯截断(置0完成开门）",
               "1号梯检修信号" := "输入"."2号梯检修信号",
               准备就绪 := "中间变量1"."2号梯准备就绪",
               "1号梯上平层信号" := "输入"."2号梯上平层信号",
               "1号梯下平层信号" := "输入"."2号梯下平层信号",
               "1层上行呼梯按钮" := "输入"."1层上行呼梯按钮",
               "2层上行呼梯按钮" := "输入"."2层上行呼梯按钮",
               "3层上行呼梯按钮" := "输入"."3层上行呼梯按钮",
               "4层上行呼梯按钮" := "输入"."4层上行呼梯按钮",
               "5层上行呼梯按钮" := "输入"."5层上行呼梯按钮",
               "6层上行呼梯按钮" := "输入"."6层上行呼梯按钮",
               "7层上行呼梯按钮" := "输入"."7层上行呼梯按钮",
               "8层上行呼梯按钮" := "输入"."8层上行呼梯按钮",
               "9层上行呼梯按钮" := "输入"."9层上行呼梯按钮",
               "2层下行呼梯按钮" := "输入"."2层下行呼梯按钮",
               "3层下行呼梯按钮" := "输入"."3层下行呼梯按钮",
               "4层下行呼梯按钮" := "输入"."4层下行呼梯按钮",
               "5层下行呼梯按钮" := "输入"."5层下行呼梯按钮",
               "6层下行呼梯按钮" := "输入"."6层下行呼梯按钮",
               "7层下行呼梯按钮" := "输入"."7层下行呼梯按钮",
               "8层下行呼梯按钮" := "输入"."8层下行呼梯按钮",
               "9层下行呼梯按钮" := "输入"."9层下行呼梯按钮",
               "10层下行呼梯按钮" := "输入"."10层下行呼梯按钮",
               "1号梯轿内选层按钮1" := "输入"."2号梯轿内选层按钮1",
               "1号梯轿内选层按钮2" := "输入"."2号梯轿内选层按钮2",
               "1号梯轿内选层按钮3" := "输入"."2号梯轿内选层按钮3",
               "1号梯轿内选层按钮4" := "输入"."2号梯轿内选层按钮4",
               "1号梯轿内选层按钮5" := "输入"."2号梯轿内选层按钮5",
               "1号梯轿内选层按钮6" := "输入"."2号梯轿内选层按钮6",
               "1号梯轿内选层按钮7" := "输入"."2号梯轿内选层按钮7",
               "1号梯轿内选层按钮8" := "输入"."2号梯轿内选层按钮8",
               "1号梯轿内选层按钮9" := "输入"."2号梯轿内选层按钮9",
               "1号梯轿内选层按钮10" := "输入"."2号梯轿内选层按钮10",
               死机 := "中间变量1".死机2,
               满载指示 := "输出"."2号梯满载指示",
               就近运动电梯 => "中间变量2".就近运动电梯2,
               "1号梯上行指示" => "输出"."2号梯上行指示",
               "1号梯下行指示" => "输出"."2号梯下行指示",
               上行接触器 => "输出"."2号梯上行接触器",
               下行接触器 => "输出"."2号梯下行接触器",
               "1号梯1层按钮指示灯" => "输出"."2号梯1层按钮指示灯",
               "1号梯2层按钮指示灯" => "输出"."2号梯2层按钮指示灯",
               "1号梯3层按钮指示灯" => "输出"."2号梯3层按钮指示灯",
               "1号梯4层按钮指示灯" => "输出"."2号梯4层按钮指示灯",
               "1号梯5层按钮指示灯" => "输出"."2号梯5层按钮指示灯",
               "1号梯6层按钮指示灯" => "输出"."2号梯6层按钮指示灯",
               "1号梯7层按钮指示灯" => "输出"."2号梯7层按钮指示灯",
               "1号梯8层按钮指示灯" => "输出"."2号梯8层按钮指示灯",
               "1号梯9层按钮指示灯" => "输出"."2号梯9层按钮指示灯",
               "1号梯10层按钮指示灯" => "输出"."2号梯10层按钮指示灯",
               "1号梯1级减速制动" => "输出"."2号梯1级减速制动",
               "1号梯2级减速制动" => "输出"."2号梯2级减速制动",
               "1号梯3级减速制动" => "输出"."2号梯3级减速制动");
END_REGION

REGION Network 3: 3号梯
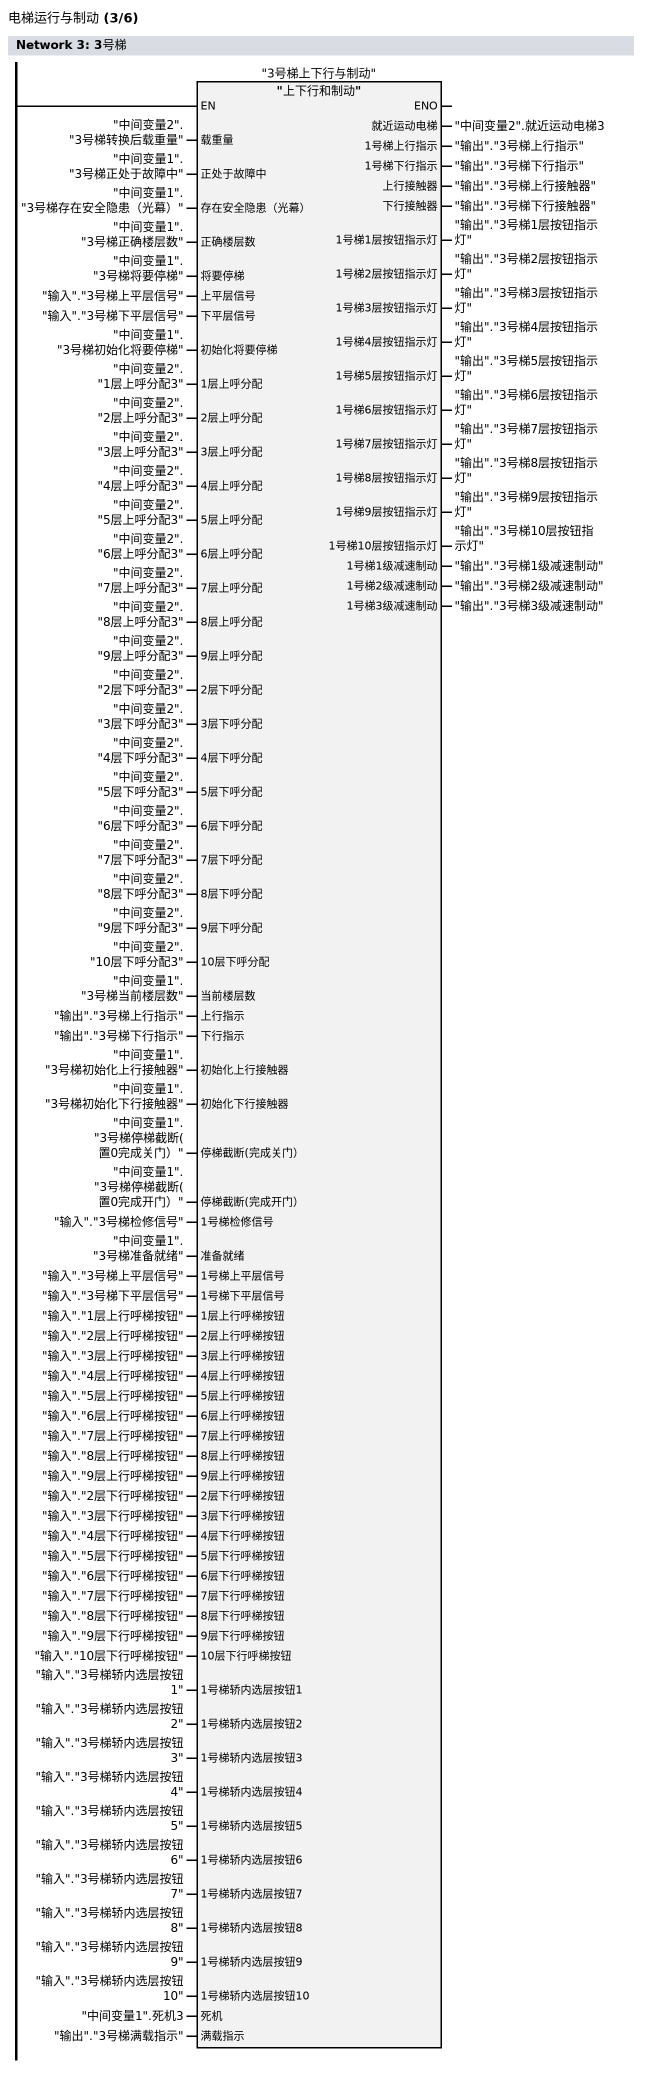
   RUNG wire#powerrail
      "3号梯上下行与制动"(载重量 := "中间变量2"."3号梯转换后载重量", 正处于故障中 := "中间变量1"."3号梯正处于故障中", "存在安全隐患（光幕）" := "中间变量1"."3号梯存在安全隐患（光幕）", 正确楼层数 := "中间变量1"."3号梯正确楼层数", 将要停梯 := "中间变量1"."3号梯将要停梯", 上平层信号 := "输入"."3号梯上平层信号", 下平层信号 := "输入"."3号梯下平层信号", 初始化将要停梯 := "中间变量1"."3号梯初始化将要停梯", "1层上呼分配" := "中间变量2"."1层上呼分配3", "2层上呼分配" := "中间变量2"."2层上呼分配3", "3层上呼分配" := "中间变量2"."3层上呼分配3", "4层上呼分配" := "中间变量2"."4层上呼分配3", "5层上呼分配" := "中间变量2"."5层上呼分配3", "6层上呼分配" := "中间变量2"."6层上呼分配3", "7层上呼分配" := "中间变量2"."7层上呼分配3", "8层上呼分配" := "中间变量2"."8层上呼分配3", "9层上呼分配" := "中间变量2"."9层上呼分配3", "2层下呼分配" := "中间变量2"."2层下呼分配3", "3层下呼分配" := "中间变量2"."3层下呼分配3", "4层下呼分配" := "中间变量2"."4层下呼分配3", "5层下呼分配" := "中间变量2"."5层下呼分配3", "6层下呼分配" := "中间变量2"."6层下呼分配3", "7层下呼分配" := "中间变量2"."7层下呼分配3", "8层下呼分配" := "中间变量2"."8层下呼分配3", "9层下呼分配" := "中间变量2"."9层下呼分配3", "10层下呼分配" := "中间变量2"."10层下呼分配3", 当前楼层数 := "中间变量1"."3号梯当前楼层数", 上行指示 := "输出"."3号梯上行指示", 下行指示 := "输出"."3号梯下行指示", 初始化上行接触器 := "中间变量1"."3号梯初始化上行接触器", 初始化下行接触器 := "中间变量1"."3号梯初始化下行接触器", "停梯截断(完成关门）" := "中间变量1"."3号梯停梯截断(置0完成关门）", "停梯截断(完成开门）" := "中间变量1"."3号梯停梯截断(置0完成开门）", "1号梯检修信号" := "输入"."3号梯检修信号", 准备就绪 := "中间变量1"."3号梯准备就绪", "1号梯上平层信号" := "输入"."3号梯上平层信号", "1号梯下平层信号" := "输入"."3号梯下平层信号", "1层上行呼梯按钮" := "输入"."1层上行呼梯按钮", "2层上行呼梯按钮" := "输入"."2层上行呼梯按钮", "3层上行呼梯按钮" := "输入"."3层上行呼梯按钮", "4层上行呼梯按钮" := "输入"."4层上行呼梯按钮", "5层上行呼梯按钮" := "输入"."5层上行呼梯按钮", "6层上行呼梯按钮" := "输入"."6层上行呼梯按钮", "7层上行呼梯按钮" := "输入"."7层上行呼梯按钮", "8层上行呼梯按钮" := "输入"."8层上行呼梯按钮", "9层上行呼梯按钮" := "输入"."9层上行呼梯按钮", "2层下行呼梯按钮" := "输入"."2层下行呼梯按钮", "3层下行呼梯按钮" := "输入"."3层下行呼梯按钮", "4层下行呼梯按钮" := "输入"."4层下行呼梯按钮", "5层下行呼梯按钮" := "输入"."5层下行呼梯按钮", "6层下行呼梯按钮" := "输入"."6层下行呼梯按钮", "7层下行呼梯按钮" := "输入"."7层下行呼梯按钮", "8层下行呼梯按钮" := "输入"."8层下行呼梯按钮", "9层下行呼梯按钮" := "输入"."9层下行呼梯按钮", "10层下行呼梯按钮" := "输入"."10层下行呼梯按钮", "1号梯轿内选层按钮1" := "输入"."3号梯轿内选层按钮1", "1号梯轿内选层按钮2" := "输入"."3号梯轿内选层按钮2", "1号梯轿内选层按钮3" := "输入"."3号梯轿内选层按钮3", "1号梯轿内选层按钮4" := "输入"."3号梯轿内选层按钮4", "1号梯轿内选层按钮5" := "输入"."3号梯轿内选层按钮5", "1号梯轿内选层按钮6" := "输入"."3号梯轿内选层按钮6", "1号梯轿内选层按钮7" := "输入"."3号梯轿内选层按钮7", "1号梯轿内选层按钮8" := "输入"."3号梯轿内选层按钮8", "1号梯轿内选层按钮9" := "输入"."3号梯轿内选层按钮9", "1号梯轿内选层按钮10" := "输入"."3号梯轿内选层按钮10", 死机 := "中间变量1".死机3, 满载指示 := "输出"."3号梯满载指示", 就近运动电梯 => "中间变量2".就近运动电梯3, "1号梯上行指示" => "输出"."3号梯上行指示", "1号梯下行指示" => "输出"."3号梯下行指示", 上行接触器 => "输出"."3号梯上行接触器", 下行接触器 => "输出"."3号梯下行接触器", "1号梯1层按钮指示灯" => "输出"."3号梯1层按钮指示灯", "1号梯2层按钮指示灯" => "输出"."3号梯2层按钮指示灯", "1号梯3层按钮指示灯" => "输出"."3号梯3层按钮指示灯", "1号梯4层按钮指示灯" => "输出"."3号梯4层按钮指示灯", "1号梯5层按钮指示灯" => "输出"."3号梯5层按钮指示灯", "1号梯6层按钮指示灯" => "输出"."3号梯6层按钮指示灯", "1号梯7层按钮指示灯" => "输出"."3号梯7层按钮指示灯", "1号梯8层按钮指示灯" => "输出"."3号梯8层按钮指示灯", "1号梯9层按钮指示灯" => "输出"."3号梯9层按钮指示灯", "1号梯10层按钮指示灯" => "输出"."3号梯10层按钮指示灯", "1号梯1级减速制动" => "输出"."3号梯1级减速制动", "1号梯2级减速制动" => "输出"."3号梯2级减速制动", "1号梯3级减速制动" => "输出"."3号梯3级减速制动")
   END_RUNG
   // the same network as SCL:
   "3号梯上下行与制动"(载重量 := "中间变量2"."3号梯转换后载重量",   // "上下行和制动"
               正处于故障中 := "中间变量1"."3号梯正处于故障中",
               "存在安全隐患（光幕）" := "中间变量1"."3号梯存在安全隐患（光幕）",
               正确楼层数 := "中间变量1"."3号梯正确楼层数",
               将要停梯 := "中间变量1"."3号梯将要停梯",
               上平层信号 := "输入"."3号梯上平层信号",
               下平层信号 := "输入"."3号梯下平层信号",
               初始化将要停梯 := "中间变量1"."3号梯初始化将要停梯",
               "1层上呼分配" := "中间变量2"."1层上呼分配3",
               "2层上呼分配" := "中间变量2"."2层上呼分配3",
               "3层上呼分配" := "中间变量2"."3层上呼分配3",
               "4层上呼分配" := "中间变量2"."4层上呼分配3",
               "5层上呼分配" := "中间变量2"."5层上呼分配3",
               "6层上呼分配" := "中间变量2"."6层上呼分配3",
               "7层上呼分配" := "中间变量2"."7层上呼分配3",
               "8层上呼分配" := "中间变量2"."8层上呼分配3",
               "9层上呼分配" := "中间变量2"."9层上呼分配3",
               "2层下呼分配" := "中间变量2"."2层下呼分配3",
               "3层下呼分配" := "中间变量2"."3层下呼分配3",
               "4层下呼分配" := "中间变量2"."4层下呼分配3",
               "5层下呼分配" := "中间变量2"."5层下呼分配3",
               "6层下呼分配" := "中间变量2"."6层下呼分配3",
               "7层下呼分配" := "中间变量2"."7层下呼分配3",
               "8层下呼分配" := "中间变量2"."8层下呼分配3",
               "9层下呼分配" := "中间变量2"."9层下呼分配3",
               "10层下呼分配" := "中间变量2"."10层下呼分配3",
               当前楼层数 := "中间变量1"."3号梯当前楼层数",
               上行指示 := "输出"."3号梯上行指示",
               下行指示 := "输出"."3号梯下行指示",
               初始化上行接触器 := "中间变量1"."3号梯初始化上行接触器",
               初始化下行接触器 := "中间变量1"."3号梯初始化下行接触器",
               "停梯截断(完成关门）" := "中间变量1"."3号梯停梯截断(置0完成关门）",
               "停梯截断(完成开门）" := "中间变量1"."3号梯停梯截断(置0完成开门）",
               "1号梯检修信号" := "输入"."3号梯检修信号",
               准备就绪 := "中间变量1"."3号梯准备就绪",
               "1号梯上平层信号" := "输入"."3号梯上平层信号",
               "1号梯下平层信号" := "输入"."3号梯下平层信号",
               "1层上行呼梯按钮" := "输入"."1层上行呼梯按钮",
               "2层上行呼梯按钮" := "输入"."2层上行呼梯按钮",
               "3层上行呼梯按钮" := "输入"."3层上行呼梯按钮",
               "4层上行呼梯按钮" := "输入"."4层上行呼梯按钮",
               "5层上行呼梯按钮" := "输入"."5层上行呼梯按钮",
               "6层上行呼梯按钮" := "输入"."6层上行呼梯按钮",
               "7层上行呼梯按钮" := "输入"."7层上行呼梯按钮",
               "8层上行呼梯按钮" := "输入"."8层上行呼梯按钮",
               "9层上行呼梯按钮" := "输入"."9层上行呼梯按钮",
               "2层下行呼梯按钮" := "输入"."2层下行呼梯按钮",
               "3层下行呼梯按钮" := "输入"."3层下行呼梯按钮",
               "4层下行呼梯按钮" := "输入"."4层下行呼梯按钮",
               "5层下行呼梯按钮" := "输入"."5层下行呼梯按钮",
               "6层下行呼梯按钮" := "输入"."6层下行呼梯按钮",
               "7层下行呼梯按钮" := "输入"."7层下行呼梯按钮",
               "8层下行呼梯按钮" := "输入"."8层下行呼梯按钮",
               "9层下行呼梯按钮" := "输入"."9层下行呼梯按钮",
               "10层下行呼梯按钮" := "输入"."10层下行呼梯按钮",
               "1号梯轿内选层按钮1" := "输入"."3号梯轿内选层按钮1",
               "1号梯轿内选层按钮2" := "输入"."3号梯轿内选层按钮2",
               "1号梯轿内选层按钮3" := "输入"."3号梯轿内选层按钮3",
               "1号梯轿内选层按钮4" := "输入"."3号梯轿内选层按钮4",
               "1号梯轿内选层按钮5" := "输入"."3号梯轿内选层按钮5",
               "1号梯轿内选层按钮6" := "输入"."3号梯轿内选层按钮6",
               "1号梯轿内选层按钮7" := "输入"."3号梯轿内选层按钮7",
               "1号梯轿内选层按钮8" := "输入"."3号梯轿内选层按钮8",
               "1号梯轿内选层按钮9" := "输入"."3号梯轿内选层按钮9",
               "1号梯轿内选层按钮10" := "输入"."3号梯轿内选层按钮10",
               死机 := "中间变量1".死机3,
               满载指示 := "输出"."3号梯满载指示",
               就近运动电梯 => "中间变量2".就近运动电梯3,
               "1号梯上行指示" => "输出"."3号梯上行指示",
               "1号梯下行指示" => "输出"."3号梯下行指示",
               上行接触器 => "输出"."3号梯上行接触器",
               下行接触器 => "输出"."3号梯下行接触器",
               "1号梯1层按钮指示灯" => "输出"."3号梯1层按钮指示灯",
               "1号梯2层按钮指示灯" => "输出"."3号梯2层按钮指示灯",
               "1号梯3层按钮指示灯" => "输出"."3号梯3层按钮指示灯",
               "1号梯4层按钮指示灯" => "输出"."3号梯4层按钮指示灯",
               "1号梯5层按钮指示灯" => "输出"."3号梯5层按钮指示灯",
               "1号梯6层按钮指示灯" => "输出"."3号梯6层按钮指示灯",
               "1号梯7层按钮指示灯" => "输出"."3号梯7层按钮指示灯",
               "1号梯8层按钮指示灯" => "输出"."3号梯8层按钮指示灯",
               "1号梯9层按钮指示灯" => "输出"."3号梯9层按钮指示灯",
               "1号梯10层按钮指示灯" => "输出"."3号梯10层按钮指示灯",
               "1号梯1级减速制动" => "输出"."3号梯1级减速制动",
               "1号梯2级减速制动" => "输出"."3号梯2级减速制动",
               "1号梯3级减速制动" => "输出"."3号梯3级减速制动");
END_REGION

REGION Network 4: 4号梯
